    RC2_Transmit_PDO_Mapping_Torque_actual_value_6077_00 : INT;
    RC2_Transmit_PDO_Mapping_Digital_inputs_60FD_00 : UDINT;
    RC2_Transmit_PDO_Mapping_Error_code_603F_00 : UINT;
    RC3_Receive_PDO_Mapping_ControlWord_6040_00 : UINT;
    RC3_Receive_PDO_Mapping_Target_Position_607A_00 : DINT;
    RC3_Receive_PDO_Mapping_Mode_of_operation_6060_00 : SINT;
    RC3_Receive_PDO_Mapping_Profile_velocity_6081_00 : UDINT;
    RC3_Receive_PDO_Mapping_Profile_acceleration_6083_00 : UDINT;
    RC3_Receive_PDO_Mapping_Profile_deceleration_6084_00 : UDINT;
    RC3_Receive_PDO_Mapping_Physical_outputs_60FE_01 : UDINT;
    RC3_Transmit_PDO_Mapping_StatusWord_6041_00 : UINT;
    RC3_Transmit_PDO_Mapping_Position_actual_value_6064_00 : DINT;
    RC3_Transmit_PDO_Mapping_Mode_of_operation_display_6061_00 : SINT;
    RC3_Transmit_PDO_Mapping_Following_error_actual_valu_60F4_00 : DINT;
    RC3_Transmit_PDO_Mapping_Torque_actual_value_6077_00 : INT;
    RC3_Transmit_PDO_Mapping_Digital_inputs_60FD_00 : UDINT;
    RC3_Transmit_PDO_Mapping_Error_code_603F_00 : UINT;
    RC4_Receive_PDO_Mapping_ControlWord_6040_00 : UINT;
    RC4_Receive_PDO_Mapping_Target_Position_607A_00 : DINT;
    RC4_Receive_PDO_Mapping_Mode_of_operation_6060_00 : SINT;
    RC4_Receive_PDO_Mapping_Profile_velocity_6081_00 : UDINT;
    RC4_Receive_PDO_Mapping_Profile_acceleration_6083_00 : UDINT;
    RC4_Receive_PDO_Mapping_Profile_deceleration_6084_00 : UDINT;
    RC4_Receive_PDO_Mapping_Physical_outputs_60FE_01 : UDINT;
    RC4_Transmit_PDO_Mapping_StatusWord_6041_00 : UINT;
    RC4_Transmit_PDO_Mapping_Position_actual_value_6064_00 : DINT;
    RC4_Transmit_PDO_Mapping_Mode_of_operation_display_6061_00 : SINT;
    RC4_Transmit_PDO_Mapping_Following_error_actual_valu_60F4_00 : DINT;
    RC4_Transmit_PDO_Mapping_Torque_actual_value_6077_00 : INT;
    RC4_Transmit_PDO_Mapping_Digital_inputs_60FD_00 : UDINT;
    RC4_Transmit_PDO_Mapping_Error_code_603F_00 : UINT;
    RC5_Receive_PDO_Mapping_ControlWord_6040_00 : UINT;
    RC5_Receive_PDO_Mapping_Target_Position_607A_00 : DINT;
    RC5_Receive_PDO_Mapping_Mode_of_operation_6060_00 : SINT;
    RC5_Receive_PDO_Mapping_Profile_velocity_6081_00 : UDINT;
    RC5_Receive_PDO_Mapping_Profile_acceleration_6083_00 : UDINT;
    RC5_Receive_PDO_Mapping_Profile_deceleration_6084_00 : UDINT;
    RC5_Receive_PDO_Mapping_Physical_outputs_60FE_01 : UDINT;
    RC5_Transmit_PDO_Mapping_StatusWord_6041_00 : UINT;
    RC5_Transmit_PDO_Mapping_Position_actual_value_6064_00 : DINT;
    RC5_Transmit_PDO_Mapping_Mode_of_operation_display_6061_00 : SINT;
    RC5_Transmit_PDO_Mapping_Following_error_actual_valu_60F4_00 : DINT;
    RC5_Transmit_PDO_Mapping_Torque_actual_value_6077_00 : INT;
    RC5_Transmit_PDO_Mapping_Digital_inputs_60FD_00 : UDINT;
    RC5_Transmit_PDO_Mapping_Error_code_603F_00 : UINT;
    RC6_Receive_PDO_Mapping_ControlWord_6040_00 : UINT;
    RC6_Receive_PDO_Mapping_ControlWord_6040_00_1 : UINT;
    RC6_Receive_PDO_Mapping_Target_Position_607A_00 : DINT;
    RC6_Receive_PDO_Mapping_Mode_of_operation_6060_00 : SINT;
    RC6_Receive_PDO_Mapping_Profile_velocity_6081_00 : UDINT;
    RC6_Receive_PDO_Mapping_Profile_acceleration_6083_00 : UDINT;
    RC6_Receive_PDO_Mapping_Profile_deceleration_6084_00 : UDINT;
    RC6_Receive_PDO_Mapping_Physical_outputs_60FE_01 : UDINT;
    RC6_Transmit_PDO_Mapping_StatusWord_6041_00 : UINT;
    RC6_Transmit_PDO_Mapping_Position_actual_value_6064_00 : DINT;
    RC6_Transmit_PDO_Mapping_Mode_of_operation_display_6061_00 : SINT;
    RC6_Transmit_PDO_Mapping_Following_error_actual_valu_60F4_00 : DINT;
    RC6_Transmit_PDO_Mapping_Torque_actual_value_6077_00 : INT;
    RC6_Transmit_PDO_Mapping_Digital_inputs_60FD_00 : UDINT;
    RC6_Transmit_PDO_Mapping_Error_code_603F_00 : UINT;
END_VAR
VAR_GLOBAL RETAIN
    RCON1_OUT : ARRAY[1..6] OF ST_RCON_Direct_OUT_Axis;  (* RCON1 (PLC→RCON); [2] 2軸目; [3] 3軸目; [4] 4軸目; [5] 5軸目; [6] 6軸目; [1].Control.Pause 一時停止（STP/b2）; [1] 1軸目 *)
    RCON1_IN : ARRAY[1..6] OF ST_RCON_Direct_IN_Axis;  (* RCON1 (RCON→PLC); [1] 1軸目; [2] 2軸目; [3] 3軸目; [4] 4軸目; [5] 5軸目; [6] 6軸目 *)
END_VAR
VAR_GLOBAL
    RCON1_SpeedUnit_mm_s : LREAL;  (* RCON1 速度単位 [mm/s/カウント]（1.0/0.1） *)
    RCON1_OUT_GwControl0Raw : UINT;  (* 未割付・不使用 OUT00 共通制御（MON/RTE） *)
    RCON1_OUT_GwControl1ReservedRaw : UINT;  (* 未割付・不使用 OUT01 予約（書込禁止） *)
    RCON1_OUT_ReservedOut02Raw : UINT;  (* 未割付・不使用 OUT02 予約（書込禁止） *)
    RCON1_OUT_ReservedOut03Raw : UINT;  (* 未割付・不使用 OUT03 予約（書込禁止） *)
    RCON1_OUT_ReservedOut04Raw : UINT;  (* 未割付・不使用 OUT04 予約（書込禁止） *)
    RCON1_OUT_ReservedOut05Raw : UINT;  (* 未割付・不使用 OUT05 予約（書込禁止） *)
    RCON1_OUT_ReservedOut06Raw : UINT;  (* 未割付・不使用 OUT06 予約（書込禁止） *)
    RCON1_OUT_ReservedOut07Raw : UINT;  (* 未割付・不使用 OUT07 予約（書込禁止） *)
    RCON1_OUT_Axis1_TargetPosLoRaw : UINT;  (* 未割付・不使用 OUT08 1軸目 目標位置 下位 [0.01mm] *)
    RCON1_OUT_Axis1_TargetPosHiRaw : UINT;  (* 未割付・不使用 OUT09 1軸目 目標位置 上位 [0.01mm] *)
    RCON1_OUT_Axis1_PositionBandLoRaw : UINT;  (* 未割付・不使用 OUT10 1軸目 位置決め幅 下位 [0.01mm] *)
    RCON1_OUT_Axis1_PositionBandHiRaw : UINT;  (* 未割付・不使用 OUT11 1軸目 位置決め幅 上位 [0.01mm] *)
    RCON1_OUT_Axis1_SpeedRaw : UINT;  (* 未割付・不使用 OUT12 1軸目 速度指令 [実機単位] *)
    RCON1_OUT_Axis1_AccDecRaw : UINT;  (* 未割付・不使用 OUT13 1軸目 共通加減速 [0.01G] *)
    RCON1_OUT_Axis1_PushLimitRaw : UINT;  (* 未割付・不使用 OUT14 1軸目 押付け制限 [255=100%] *)
    RCON1_OUT_Axis1_ControlRaw : UINT;  (* 未割付・不使用 OUT15 1軸目 制御信号（DSTR/SON等） *)
    RCON1_OUT_Axis2_TargetPosLoRaw : UINT;  (* 未割付・不使用 OUT16 2軸目 目標位置 下位 [0.01mm] *)
    RCON1_OUT_Axis2_TargetPosHiRaw : UINT;  (* 未割付・不使用 OUT17 2軸目 目標位置 上位 [0.01mm] *)
    RCON1_OUT_Axis2_PositionBandLoRaw : UINT;  (* 未割付・不使用 OUT18 2軸目 位置決め幅 下位 [0.01mm] *)
    RCON1_OUT_Axis2_PositionBandHiRaw : UINT;  (* 未割付・不使用 OUT19 2軸目 位置決め幅 上位 [0.01mm] *)
    RCON1_OUT_Axis2_SpeedRaw : UINT;  (* 未割付・不使用 OUT20 2軸目 速度指令 [実機単位] *)
    RCON1_OUT_Axis2_AccDecRaw : UINT;  (* 未割付・不使用 OUT21 2軸目 共通加減速 [0.01G] *)
    RCON1_OUT_Axis2_PushLimitRaw : UINT;  (* 未割付・不使用 OUT22 2軸目 押付け制限 [255=100%] *)
    RCON1_OUT_Axis2_ControlRaw : UINT;  (* 未割付・不使用 OUT23 2軸目 制御信号（DSTR/SON等） *)
    RCON1_OUT_Axis3_TargetPosLoRaw : UINT;  (* 未割付・不使用 OUT24 3軸目 目標位置 下位 [0.01mm] *)
    RCON1_OUT_Axis3_TargetPosHiRaw : UINT;  (* 未割付・不使用 OUT25 3軸目 目標位置 上位 [0.01mm] *)
    RCON1_OUT_Axis3_PositionBandLoRaw : UINT;  (* 未割付・不使用 OUT26 3軸目 位置決め幅 下位 [0.01mm] *)
    RCON1_OUT_Axis3_PositionBandHiRaw : UINT;  (* 未割付・不使用 OUT27 3軸目 位置決め幅 上位 [0.01mm] *)
    RCON1_OUT_Axis3_SpeedRaw : UINT;  (* 未割付・不使用 OUT28 3軸目 速度指令 [実機単位] *)
    RCON1_OUT_Axis3_AccDecRaw : UINT;  (* 未割付・不使用 OUT29 3軸目 共通加減速 [0.01G] *)
    RCON1_OUT_Axis3_PushLimitRaw : UINT;  (* 未割付・不使用 OUT30 3軸目 押付け制限 [255=100%] *)
    RCON1_OUT_Axis3_ControlRaw : UINT;  (* 未割付・不使用 OUT31 3軸目 制御信号（DSTR/SON等） *)
    RCON1_OUT_Axis4_TargetPosLoRaw : UINT;  (* 未割付・不使用 OUT32 4軸目 目標位置 下位 [0.01mm] *)
    RCON1_OUT_Axis4_TargetPosHiRaw : UINT;  (* 未割付・不使用 OUT33 4軸目 目標位置 上位 [0.01mm] *)
    RCON1_OUT_Axis4_PositionBandLoRaw : UINT;  (* 未割付・不使用 OUT34 4軸目 位置決め幅 下位 [0.01mm] *)
    RCON1_OUT_Axis4_PositionBandHiRaw : UINT;  (* 未割付・不使用 OUT35 4軸目 位置決め幅 上位 [0.01mm] *)
    RCON1_OUT_Axis4_SpeedRaw : UINT;  (* 未割付・不使用 OUT36 4軸目 速度指令 [実機単位] *)
    RCON1_OUT_Axis4_AccDecRaw : UINT;  (* 未割付・不使用 OUT37 4軸目 共通加減速 [0.01G] *)
    RCON1_OUT_Axis4_PushLimitRaw : UINT;  (* 未割付・不使用 OUT38 4軸目 押付け制限 [255=100%] *)
    RCON1_OUT_Axis4_ControlRaw : UINT;  (* 未割付・不使用 OUT39 4軸目 制御信号（DSTR/SON等） *)
    RCON1_OUT_Axis5_TargetPosLoRaw : UINT;  (* 未割付・不使用 OUT40 5軸目 目標位置 下位 [0.01mm] *)
    RCON1_OUT_Axis5_TargetPosHiRaw : UINT;  (* 未割付・不使用 OUT41 5軸目 目標位置 上位 [0.01mm] *)
    RCON1_OUT_Axis5_PositionBandLoRaw : UINT;  (* 未割付・不使用 OUT42 5軸目 位置決め幅 下位 [0.01mm] *)
    RCON1_OUT_Axis5_PositionBandHiRaw : UINT;  (* 未割付・不使用 OUT43 5軸目 位置決め幅 上位 [0.01mm] *)
    RCON1_OUT_Axis5_SpeedRaw : UINT;  (* 未割付・不使用 OUT44 5軸目 速度指令 [実機単位] *)
    RCON1_OUT_Axis5_AccDecRaw : UINT;  (* 未割付・不使用 OUT45 5軸目 共通加減速 [0.01G] *)
    RCON1_OUT_Axis5_PushLimitRaw : UINT;  (* 未割付・不使用 OUT46 5軸目 押付け制限 [255=100%] *)
    RCON1_OUT_Axis5_ControlRaw : UINT;  (* 未割付・不使用 OUT47 5軸目 制御信号（DSTR/SON等） *)
    RCON1_OUT_Axis6_TargetPosLoRaw : UINT;  (* 未割付・不使用 OUT48 6軸目 目標位置 下位 [0.01mm] *)
    RCON1_OUT_Axis6_TargetPosHiRaw : UINT;  (* 未割付・不使用 OUT49 6軸目 目標位置 上位 [0.01mm] *)
    RCON1_OUT_Axis6_PositionBandLoRaw : UINT;  (* 未割付・不使用 OUT50 6軸目 位置決め幅 下位 [0.01mm] *)
    RCON1_OUT_Axis6_PositionBandHiRaw : UINT;  (* 未割付・不使用 OUT51 6軸目 位置決め幅 上位 [0.01mm] *)
    RCON1_OUT_Axis6_SpeedRaw : UINT;  (* 未割付・不使用 OUT52 6軸目 速度指令 [実機単位] *)
    RCON1_OUT_Axis6_AccDecRaw : UINT;  (* 未割付・不使用 OUT53 6軸目 共通加減速 [0.01G] *)
    RCON1_OUT_Axis6_PushLimitRaw : UINT;  (* 未割付・不使用 OUT54 6軸目 押付け制限 [255=100%] *)
    RCON1_OUT_Axis6_ControlRaw : UINT;  (* 未割付・不使用 OUT55 6軸目 制御信号（DSTR/SON等） *)
    RCON1_IN_GwStatus0Raw : UINT;  (* 未割付・不使用 IN00 GW状態 *)
    RCON1_IN_AxisLinkStatusRaw : UINT;  (* 未割付・不使用 IN01 軸リンク状態 *)
    RCON1_IN_PowerStatus0Raw : UINT;  (* 未割付・不使用 IN02 電源状態0 *)
    RCON1_IN_PowerStatus1Raw : UINT;  (* 未割付・不使用 IN03 電源状態1 *)
    RCON1_IN_PowerStatus2Raw : UINT;  (* 未割付・不使用 IN04 電源状態2 *)
    RCON1_IN_PowerStatus3Raw : UINT;  (* 未割付・不使用 IN05 電源状態3 *)
    RCON1_IN_PowerStatus4MaintenanceRaw : UINT;  (* 未割付・不使用 IN06 電源状態4（構成依存） *)
    RCON1_IN_ReservedIn07Raw : UINT;  (* 未割付・不使用 IN07 予約（使用禁止） *)
    RCON1_IN_Axis1_ActualPosLoRaw : UINT;  (* 未割付・不使用 IN08 1軸目 現在位置 下位 [0.01mm] *)
    RCON1_IN_Axis1_ActualPosHiRaw : UINT;  (* 未割付・不使用 IN09 1軸目 現在位置 上位 [0.01mm] *)
    RCON1_IN_Axis1_CurrentLoRaw : UINT;  (* 未割付・不使用 IN10 1軸目 指令電流 下位 [mA] *)
    RCON1_IN_Axis1_CurrentHiRaw : UINT;  (* 未割付・不使用 IN11 1軸目 指令電流 上位 [mA] *)
    RCON1_IN_Axis1_ActualSpeedRaw : UINT;  (* 未割付・不使用 IN12 1軸目 現在速度 [実機単位・符号付き] *)
    RCON1_IN_Axis1_ReservedInRaw : UINT;  (* 未割付・不使用 IN13 1軸目 予約（使用禁止） *)
    RCON1_IN_Axis1_AlarmCodeRaw : UINT;  (* 未割付・不使用 IN14 1軸目 軸異常コード *)
    RCON1_IN_Axis1_StatusRaw : UINT;  (* 未割付・不使用 IN15 1軸目 状態信号（PEND/SV等） *)
    RCON1_IN_Axis2_ActualPosLoRaw : UINT;  (* 未割付・不使用 IN16 2軸目 現在位置 下位 [0.01mm] *)
    RCON1_IN_Axis2_ActualPosHiRaw : UINT;  (* 未割付・不使用 IN17 2軸目 現在位置 上位 [0.01mm] *)
    RCON1_IN_Axis2_CurrentLoRaw : UINT;  (* 未割付・不使用 IN18 2軸目 指令電流 下位 [mA] *)
    RCON1_IN_Axis2_CurrentHiRaw : UINT;  (* 未割付・不使用 IN19 2軸目 指令電流 上位 [mA] *)
    RCON1_IN_Axis2_ActualSpeedRaw : UINT;  (* 未割付・不使用 IN20 2軸目 現在速度 [実機単位・符号付き] *)
    RCON1_IN_Axis2_ReservedInRaw : UINT;  (* 未割付・不使用 IN21 2軸目 予約（使用禁止） *)
    RCON1_IN_Axis2_AlarmCodeRaw : UINT;  (* 未割付・不使用 IN22 2軸目 軸異常コード *)
    RCON1_IN_Axis2_StatusRaw : UINT;  (* 未割付・不使用 IN23 2軸目 状態信号（PEND/SV等） *)
    RCON1_IN_Axis3_ActualPosLoRaw : UINT;  (* 未割付・不使用 IN24 3軸目 現在位置 下位 [0.01mm] *)
    RCON1_IN_Axis3_ActualPosHiRaw : UINT;  (* 未割付・不使用 IN25 3軸目 現在位置 上位 [0.01mm] *)
    RCON1_IN_Axis3_CurrentLoRaw : UINT;  (* 未割付・不使用 IN26 3軸目 指令電流 下位 [mA] *)
    RCON1_IN_Axis3_CurrentHiRaw : UINT;  (* 未割付・不使用 IN27 3軸目 指令電流 上位 [mA] *)
    RCON1_IN_Axis3_ActualSpeedRaw : UINT;  (* 未割付・不使用 IN28 3軸目 現在速度 [実機単位・符号付き] *)
    RCON1_IN_Axis3_ReservedInRaw : UINT;  (* 未割付・不使用 IN29 3軸目 予約（使用禁止） *)
    RCON1_IN_Axis3_AlarmCodeRaw : UINT;  (* 未割付・不使用 IN30 3軸目 軸異常コード *)
    RCON1_IN_Axis3_StatusRaw : UINT;  (* 未割付・不使用 IN31 3軸目 状態信号（PEND/SV等） *)
    RCON1_IN_Axis4_ActualPosLoRaw : UINT;  (* 未割付・不使用 IN32 4軸目 現在位置 下位 [0.01mm] *)
    RCON1_IN_Axis4_ActualPosHiRaw : UINT;  (* 未割付・不使用 IN33 4軸目 現在位置 上位 [0.01mm] *)
    RCON1_IN_Axis4_CurrentLoRaw : UINT;  (* 未割付・不使用 IN34 4軸目 指令電流 下位 [mA] *)
    RCON1_IN_Axis4_CurrentHiRaw : UINT;  (* 未割付・不使用 IN35 4軸目 指令電流 上位 [mA] *)
    RCON1_IN_Axis4_ActualSpeedRaw : UINT;  (* 未割付・不使用 IN36 4軸目 現在速度 [実機単位・符号付き] *)
    RCON1_IN_Axis4_ReservedInRaw : UINT;  (* 未割付・不使用 IN37 4軸目 予約（使用禁止） *)
    RCON1_IN_Axis4_AlarmCodeRaw : UINT;  (* 未割付・不使用 IN38 4軸目 軸異常コード *)
    RCON1_IN_Axis4_StatusRaw : UINT;  (* 未割付・不使用 IN39 4軸目 状態信号（PEND/SV等） *)
    RCON1_IN_Axis5_ActualPosLoRaw : UINT;  (* 未割付・不使用 IN40 5軸目 現在位置 下位 [0.01mm] *)
    RCON1_IN_Axis5_ActualPosHiRaw : UINT;  (* 未割付・不使用 IN41 5軸目 現在位置 上位 [0.01mm] *)
    RCON1_IN_Axis5_CurrentLoRaw : UINT;  (* 未割付・不使用 IN42 5軸目 指令電流 下位 [mA] *)
    RCON1_IN_Axis5_CurrentHiRaw : UINT;  (* 未割付・不使用 IN43 5軸目 指令電流 上位 [mA] *)
    RCON1_IN_Axis5_ActualSpeedRaw : UINT;  (* 未割付・不使用 IN44 5軸目 現在速度 [実機単位・符号付き] *)
    RCON1_IN_Axis5_ReservedInRaw : UINT;  (* 未割付・不使用 IN45 5軸目 予約（使用禁止） *)
    RCON1_IN_Axis5_AlarmCodeRaw : UINT;  (* 未割付・不使用 IN46 5軸目 軸異常コード *)
    RCON1_IN_Axis5_StatusRaw : UINT;  (* 未割付・不使用 IN47 5軸目 状態信号（PEND/SV等） *)
    RCON1_IN_Axis6_ActualPosLoRaw : UINT;  (* 未割付・不使用 IN48 6軸目 現在位置 下位 [0.01mm] *)
    RCON1_IN_Axis6_ActualPosHiRaw : UINT;  (* 未割付・不使用 IN49 6軸目 現在位置 上位 [0.01mm] *)
    RCON1_IN_Axis6_CurrentLoRaw : UINT;  (* 未割付・不使用 IN50 6軸目 指令電流 下位 [mA] *)
    RCON1_IN_Axis6_CurrentHiRaw : UINT;  (* 未割付・不使用 IN51 6軸目 指令電流 上位 [mA] *)
    RCON1_IN_Axis6_ActualSpeedRaw : UINT;  (* 未割付・不使用 IN52 6軸目 現在速度 [実機単位・符号付き] *)
    RCON1_IN_Axis6_ReservedInRaw : UINT;  (* 未割付・不使用 IN53 6軸目 予約（使用禁止） *)
    RCON1_IN_Axis6_AlarmCodeRaw : UINT;  (* 未割付・不使用 IN54 6軸目 軸異常コード *)
END_VAR
VAR_GLOBAL RETAIN
    RCON1_IN_Axis6_StatusRaw : UINT;  (* 未割付・不使用 IN55 6軸目 状態信号（PEND/SV等） *)
    RCON2_OUT : ARRAY[1..5] OF ST_RCON_Direct_OUT_Axis;  (* RCON2 出力指令（PLC→RCON）; [1] 1軸目（No.0）出力指令; [2] 2軸目（No.1）出力指令; [3] 3軸目（No.2）出力指令; [4] 4軸目（No.3）出力指令; [5] 5軸目（No.4）出力指令 *)
END_VAR
VAR_GLOBAL
    RCON2_IN : ARRAY[1..5] OF ST_RCON_Direct_IN_Axis;  (* RCON2 入力情報（RCON→PLC）; [1] 1軸目（No.0）入力情報; [2] 2軸目（No.1）入力情報; [3] 3軸目（No.2）入力情報; [4] 4軸目（No.3）入力情報; [5] 5軸目（No.4）入力情報 *)
    RCON2_SpeedUnit_mm_s : LREAL;  (* RCON2 速度単位 [mm/s/カウント]（1.0/0.1） *)
    RCON2_OUT_GwControl0Raw : UINT;  (* 未割付・不使用 OUT00 共通制御（MON/RTE） *)
    RCON2_OUT_GwControl1ReservedRaw : UINT;  (* 未割付・不使用 OUT01 予約（書込禁止） *)
    RCON2_OUT_ReservedOut02Raw : UINT;  (* 未割付・不使用 OUT02 予約（書込禁止） *)
    RCON2_OUT_ReservedOut03Raw : UINT;  (* 未割付・不使用 OUT03 予約（書込禁止） *)
    RCON2_OUT_ReservedOut04Raw : UINT;  (* 未割付・不使用 OUT04 予約（書込禁止） *)
    RCON2_OUT_ReservedOut05Raw : UINT;  (* 未割付・不使用 OUT05 予約（書込禁止） *)
    RCON2_OUT_ReservedOut06Raw : UINT;  (* 未割付・不使用 OUT06 予約（書込禁止） *)
    RCON2_OUT_ReservedOut07Raw : UINT;  (* 未割付・不使用 OUT07 予約（書込禁止） *)
    RCON2_OUT_Axis1_TargetPosLoRaw : UINT;  (* 未割付・不使用 OUT08 1軸目 目標位置 下位 [0.01mm] *)
    RCON2_OUT_Axis1_TargetPosHiRaw : UINT;  (* 未割付・不使用 OUT09 1軸目 目標位置 上位 [0.01mm] *)
    RCON2_OUT_Axis1_PositionBandLoRaw : UINT;  (* 未割付・不使用 OUT10 1軸目 位置決め幅 下位 [0.01mm] *)
    RCON2_OUT_Axis1_PositionBandHiRaw : UINT;  (* 未割付・不使用 OUT11 1軸目 位置決め幅 上位 [0.01mm] *)
    RCON2_OUT_Axis1_SpeedRaw : UINT;  (* 未割付・不使用 OUT12 1軸目 速度指令 [実機単位] *)
    RCON2_OUT_Axis1_AccDecRaw : UINT;  (* 未割付・不使用 OUT13 1軸目 共通加減速 [0.01G] *)
    RCON2_OUT_Axis1_PushLimitRaw : UINT;  (* 未割付・不使用 OUT14 1軸目 押付け制限 [255=100%] *)
    RCON2_OUT_Axis1_ControlRaw : UINT;  (* 未割付・不使用 OUT15 1軸目 制御信号（DSTR/SON等） *)
    RCON2_OUT_Axis2_TargetPosLoRaw : UINT;  (* 未割付・不使用 OUT16 2軸目 目標位置 下位 [0.01mm] *)
    RCON2_OUT_Axis2_TargetPosHiRaw : UINT;  (* 未割付・不使用 OUT17 2軸目 目標位置 上位 [0.01mm] *)
    RCON2_OUT_Axis2_PositionBandLoRaw : UINT;  (* 未割付・不使用 OUT18 2軸目 位置決め幅 下位 [0.01mm] *)
    RCON2_OUT_Axis2_PositionBandHiRaw : UINT;  (* 未割付・不使用 OUT19 2軸目 位置決め幅 上位 [0.01mm] *)
    RCON2_OUT_Axis2_SpeedRaw : UINT;  (* 未割付・不使用 OUT20 2軸目 速度指令 [実機単位] *)
    RCON2_OUT_Axis2_AccDecRaw : UINT;  (* 未割付・不使用 OUT21 2軸目 共通加減速 [0.01G] *)
    RCON2_OUT_Axis2_PushLimitRaw : UINT;  (* 未割付・不使用 OUT22 2軸目 押付け制限 [255=100%] *)
    RCON2_OUT_Axis2_ControlRaw : UINT;  (* 未割付・不使用 OUT23 2軸目 制御信号（DSTR/SON等） *)
    RCON2_OUT_Axis3_TargetPosLoRaw : UINT;  (* 未割付・不使用 OUT24 3軸目 目標位置 下位 [0.01mm] *)
    RCON2_OUT_Axis3_TargetPosHiRaw : UINT;  (* 未割付・不使用 OUT25 3軸目 目標位置 上位 [0.01mm] *)
    RCON2_OUT_Axis3_PositionBandLoRaw : UINT;  (* 未割付・不使用 OUT26 3軸目 位置決め幅 下位 [0.01mm] *)
    RCON2_OUT_Axis3_PositionBandHiRaw : UINT;  (* 未割付・不使用 OUT27 3軸目 位置決め幅 上位 [0.01mm] *)
    RCON2_OUT_Axis3_SpeedRaw : UINT;  (* 未割付・不使用 OUT28 3軸目 速度指令 [実機単位] *)
    RCON2_OUT_Axis3_AccDecRaw : UINT;  (* 未割付・不使用 OUT29 3軸目 共通加減速 [0.01G] *)
    RCON2_OUT_Axis3_PushLimitRaw : UINT;  (* 未割付・不使用 OUT30 3軸目 押付け制限 [255=100%] *)
    RCON2_OUT_Axis3_ControlRaw : UINT;  (* 未割付・不使用 OUT31 3軸目 制御信号（DSTR/SON等） *)
    RCON2_OUT_Axis4_TargetPosLoRaw : UINT;  (* 未割付・不使用 OUT32 4軸目 目標位置 下位 [0.01mm] *)
    RCON2_OUT_Axis4_TargetPosHiRaw : UINT;  (* 未割付・不使用 OUT33 4軸目 目標位置 上位 [0.01mm] *)
    RCON2_OUT_Axis4_PositionBandLoRaw : UINT;  (* 未割付・不使用 OUT34 4軸目 位置決め幅 下位 [0.01mm] *)
    RCON2_OUT_Axis4_PositionBandHiRaw : UINT;  (* 未割付・不使用 OUT35 4軸目 位置決め幅 上位 [0.01mm] *)
    RCON2_OUT_Axis4_SpeedRaw : UINT;  (* 未割付・不使用 OUT36 4軸目 速度指令 [実機単位] *)
    RCON2_OUT_Axis4_AccDecRaw : UINT;  (* 未割付・不使用 OUT37 4軸目 共通加減速 [0.01G] *)
    RCON2_OUT_Axis4_PushLimitRaw : UINT;  (* 未割付・不使用 OUT38 4軸目 押付け制限 [255=100%] *)
    RCON2_OUT_Axis4_ControlRaw : UINT;  (* 未割付・不使用 OUT39 4軸目 制御信号（DSTR/SON等） *)
    RCON2_OUT_Axis5_TargetPosLoRaw : UINT;  (* 未割付・不使用 OUT40 5軸目 目標位置 下位 [0.01mm] *)
    RCON2_OUT_Axis5_TargetPosHiRaw : UINT;  (* 未割付・不使用 OUT41 5軸目 目標位置 上位 [0.01mm] *)
    RCON2_OUT_Axis5_PositionBandLoRaw : UINT;  (* 未割付・不使用 OUT42 5軸目 位置決め幅 下位 [0.01mm] *)
    RCON2_OUT_Axis5_PositionBandHiRaw : UINT;  (* 未割付・不使用 OUT43 5軸目 位置決め幅 上位 [0.01mm] *)
    RCON2_OUT_Axis5_SpeedRaw : UINT;  (* 未割付・不使用 OUT44 5軸目 速度指令 [実機単位] *)
    RCON2_OUT_Axis5_AccDecRaw : UINT;  (* 未割付・不使用 OUT45 5軸目 共通加減速 [0.01G] *)
    RCON2_OUT_Axis5_PushLimitRaw : UINT;  (* 未割付・不使用 OUT46 5軸目 押付け制限 [255=100%] *)
    RCON2_OUT_Axis5_ControlRaw : UINT;  (* 未割付・不使用 OUT47 5軸目 制御信号（DSTR/SON等） *)
    RCON2_IN_GwStatus0Raw : UINT;  (* 未割付・不使用 IN00 GW状態 *)
    RCON2_IN_AxisLinkStatusRaw : UINT;  (* 未割付・不使用 IN01 軸リンク状態 *)
    RCON2_IN_PowerStatus0Raw : UINT;  (* 未割付・不使用 IN02 電源状態0 *)
    RCON2_IN_PowerStatus1Raw : UINT;  (* 未割付・不使用 IN03 電源状態1 *)
    RCON2_IN_PowerStatus2Raw : UINT;  (* 未割付・不使用 IN04 電源状態2 *)
    RCON2_IN_PowerStatus3Raw : UINT;  (* 未割付・不使用 IN05 電源状態3 *)
    RCON2_IN_PowerStatus4MaintenanceRaw : UINT;  (* 未割付・不使用 IN06 電源状態4（構成依存） *)
    RCON2_IN_ReservedIn07Raw : UINT;  (* 未割付・不使用 IN07 予約（使用禁止） *)
    RCON2_IN_Axis1_ActualPosLoRaw : UINT;  (* 未割付・不使用 IN08 1軸目 現在位置 下位 [0.01mm] *)
    RCON2_IN_Axis1_ActualPosHiRaw : UINT;  (* 未割付・不使用 IN09 1軸目 現在位置 上位 [0.01mm] *)
    RCON2_IN_Axis1_CurrentLoRaw : UINT;  (* 未割付・不使用 IN10 1軸目 指令電流 下位 [mA] *)
    RCON2_IN_Axis1_CurrentHiRaw : UINT;  (* 未割付・不使用 IN11 1軸目 指令電流 上位 [mA] *)
    RCON2_IN_Axis1_ActualSpeedRaw : UINT;  (* 未割付・不使用 IN12 1軸目 現在速度 [実機単位・符号付き] *)
    RCON2_IN_Axis1_ReservedInRaw : UINT;  (* 未割付・不使用 IN13 1軸目 予約（使用禁止） *)
    RCON2_IN_Axis1_AlarmCodeRaw : UINT;  (* 未割付・不使用 IN14 1軸目 軸異常コード *)
    RCON2_IN_Axis1_StatusRaw : UINT;  (* 未割付・不使用 IN15 1軸目 状態信号（PEND/SV等） *)
    RCON2_IN_Axis2_ActualPosLoRaw : UINT;  (* 未割付・不使用 IN16 2軸目 現在位置 下位 [0.01mm] *)
    RCON2_IN_Axis2_ActualPosHiRaw : UINT;  (* 未割付・不使用 IN17 2軸目 現在位置 上位 [0.01mm] *)
    RCON2_IN_Axis2_CurrentLoRaw : UINT;  (* 未割付・不使用 IN18 2軸目 指令電流 下位 [mA] *)
    RCON2_IN_Axis2_CurrentHiRaw : UINT;  (* 未割付・不使用 IN19 2軸目 指令電流 上位 [mA] *)
    RCON2_IN_Axis2_ActualSpeedRaw : UINT;  (* 未割付・不使用 IN20 2軸目 現在速度 [実機単位・符号付き] *)
    RCON2_IN_Axis2_ReservedInRaw : UINT;  (* 未割付・不使用 IN21 2軸目 予約（使用禁止） *)
    RCON2_IN_Axis2_AlarmCodeRaw : UINT;  (* 未割付・不使用 IN22 2軸目 軸異常コード *)
    RCON2_IN_Axis2_StatusRaw : UINT;  (* 未割付・不使用 IN23 2軸目 状態信号（PEND/SV等） *)
    RCON2_IN_Axis3_ActualPosLoRaw : UINT;  (* 未割付・不使用 IN24 3軸目 現在位置 下位 [0.01mm] *)
    RCON2_IN_Axis3_ActualPosHiRaw : UINT;  (* 未割付・不使用 IN25 3軸目 現在位置 上位 [0.01mm] *)
    RCON2_IN_Axis3_CurrentLoRaw : UINT;  (* 未割付・不使用 IN26 3軸目 指令電流 下位 [mA] *)
    RCON2_IN_Axis3_CurrentHiRaw : UINT;  (* 未割付・不使用 IN27 3軸目 指令電流 上位 [mA] *)
    RCON2_IN_Axis3_ActualSpeedRaw : UINT;  (* 未割付・不使用 IN28 3軸目 現在速度 [実機単位・符号付き] *)
    RCON2_IN_Axis3_ReservedInRaw : UINT;  (* 未割付・不使用 IN29 3軸目 予約（使用禁止） *)
    RCON2_IN_Axis3_AlarmCodeRaw : UINT;  (* 未割付・不使用 IN30 3軸目 軸異常コード *)
    RCON2_IN_Axis3_StatusRaw : UINT;  (* 未割付・不使用 IN31 3軸目 状態信号（PEND/SV等） *)
    RCON2_IN_Axis4_ActualPosLoRaw : UINT;  (* 未割付・不使用 IN32 4軸目 現在位置 下位 [0.01mm] *)
    RCON2_IN_Axis4_ActualPosHiRaw : UINT;  (* 未割付・不使用 IN33 4軸目 現在位置 上位 [0.01mm] *)
    RCON2_IN_Axis4_CurrentLoRaw : UINT;  (* 未割付・不使用 IN34 4軸目 指令電流 下位 [mA] *)
    RCON2_IN_Axis4_CurrentHiRaw : UINT;  (* 未割付・不使用 IN35 4軸目 指令電流 上位 [mA] *)
    RCON2_IN_Axis4_ActualSpeedRaw : UINT;  (* 未割付・不使用 IN36 4軸目 現在速度 [実機単位・符号付き] *)
    RCON2_IN_Axis4_ReservedInRaw : UINT;  (* 未割付・不使用 IN37 4軸目 予約（使用禁止） *)
    RCON2_IN_Axis4_AlarmCodeRaw : UINT;  (* 未割付・不使用 IN38 4軸目 軸異常コード *)
    RCON2_IN_Axis4_StatusRaw : UINT;  (* 未割付・不使用 IN39 4軸目 状態信号（PEND/SV等） *)
    RCON2_IN_Axis5_ActualPosLoRaw : UINT;  (* 未割付・不使用 IN40 5軸目 現在位置 下位 [0.01mm] *)
    RCON2_IN_Axis5_ActualPosHiRaw : UINT;  (* 未割付・不使用 IN41 5軸目 現在位置 上位 [0.01mm] *)
    RCON2_IN_Axis5_CurrentLoRaw : UINT;  (* 未割付・不使用 IN42 5軸目 指令電流 下位 [mA] *)
    RCON2_IN_Axis5_CurrentHiRaw : UINT;  (* 未割付・不使用 IN43 5軸目 指令電流 上位 [mA] *)
    RCON2_IN_Axis5_ActualSpeedRaw : UINT;  (* 未割付・不使用 IN44 5軸目 現在速度 [実機単位・符号付き] *)
    RCON2_IN_Axis5_ReservedInRaw : UINT;  (* 未割付・不使用 IN45 5軸目 予約（使用禁止） *)
    RCON2_IN_Axis5_AlarmCodeRaw : UINT;  (* 未割付・不使用 IN46 5軸目 軸異常コード *)
    RCON2_IN_Axis5_StatusRaw : UINT;  (* 未割付・不使用 IN47 5軸目 状態信号（PEND/SV等） *)
    E005_Out_OUT00_2003_01 : UINT;  (* 旧I/O候補（未割付・不使用） *)
    E005_Out_OUT01_2003_02 : UINT;  (* 旧I/O候補（未割付・不使用） *)
    E005_Out_OUT02_2003_03 : UINT;  (* 旧I/O候補（未割付・不使用） *)
    E005_Out_OUT03_2003_04 : UINT;  (* 旧I/O候補（未割付・不使用） *)
    E005_Out_OUT04_2003_05 : UINT;  (* 旧I/O候補（未割付・不使用） *)
    E005_Out_OUT05_2003_06 : UINT;  (* 旧I/O候補（未割付・不使用） *)
    E005_Out_OUT06_2003_07 : UINT;  (* 旧I/O候補（未割付・不使用） *)
    E005_Out_OUT07_2003_08 : UINT;  (* 旧I/O候補（未割付・不使用） *)
    E005_Out_OUT08_2003_09 : UINT;  (* 旧I/O候補（未割付・不使用） *)
    E005_Out_OUT09_2003_0A : UINT;  (* 旧I/O候補（未割付・不使用） *)
    E005_Out_OUT10_2003_0B : UINT;  (* 旧I/O候補（未割付・不使用） *)
    E005_Out_OUT11_2003_0C : UINT;  (* 旧I/O候補（未割付・不使用） *)
    E005_Out_OUT12_2003_0D : UINT;  (* 旧I/O候補（未割付・不使用） *)
    E005_Out_OUT13_2003_0E : UINT;  (* 旧I/O候補（未割付・不使用） *)
    E005_Out_OUT14_2003_0F : UINT;  (* 旧I/O候補（未割付・不使用） *)
    E005_Out_OUT15_2003_10 : UINT;  (* 旧I/O候補（未割付・不使用） *)
    E005_Out_OUT16_2003_11 : UINT;  (* 旧I/O候補（未割付・不使用） *)
    E005_Out_OUT17_2003_12 : UINT;  (* 旧I/O候補（未割付・不使用） *)
    E005_Out_OUT18_2003_13 : UINT;  (* 旧I/O候補（未割付・不使用） *)
    E005_Out_OUT19_2003_14 : UINT;  (* 旧I/O候補（未割付・不使用） *)
    E005_Out_OUT20_2003_15 : UINT;  (* 旧I/O候補（未割付・不使用） *)
    E005_Out_OUT21_2003_16 : UINT;  (* 旧I/O候補（未割付・不使用） *)
    E005_Out_OUT22_2003_17 : UINT;  (* 旧I/O候補（未割付・不使用） *)
    E005_Out_OUT23_2003_18 : UINT;  (* 旧I/O候補（未割付・不使用） *)
    E005_Out_OUT24_2003_19 : UINT;  (* 旧I/O候補（未割付・不使用） *)
    E005_Out_OUT25_2003_1A : UINT;  (* 旧I/O候補（未割付・不使用） *)
    E005_Out_OUT26_2003_1B : UINT;  (* 旧I/O候補（未割付・不使用） *)
    E005_Out_OUT27_2003_1C : UINT;  (* 旧I/O候補（未割付・不使用） *)
    E005_Out_OUT28_2003_1D : UINT;  (* 旧I/O候補（未割付・不使用） *)
    E005_Out_OUT29_2003_1E : UINT;  (* 旧I/O候補（未割付・不使用） *)
    E005_Out_OUT30_2003_1F : UINT;  (* 旧I/O候補（未割付・不使用） *)
    E005_Out_OUT31_2003_20 : UINT;  (* 旧I/O候補（未割付・不使用） *)
    E005_Out_OUT32_2003_21 : UINT;  (* 旧I/O候補（未割付・不使用） *)
    E005_Out_OUT33_2003_22 : UINT;  (* 旧I/O候補（未割付・不使用） *)
    E005_Out_OUT34_2003_23 : UINT;  (* 旧I/O候補（未割付・不使用） *)
    E005_Out_OUT35_2003_24 : UINT;  (* 旧I/O候補（未割付・不使用） *)
    E005_Out_OUT36_2003_25 : UINT;  (* 旧I/O候補（未割付・不使用） *)
    E005_Out_OUT37_2003_26 : UINT;  (* 旧I/O候補（未割付・不使用） *)
    E005_Out_OUT38_2003_27 : UINT;  (* 旧I/O候補（未割付・不使用） *)
    E005_Out_OUT39_2003_28 : UINT;  (* 旧I/O候補（未割付・不使用） *)
    E005_Out_OUT40_2003_29 : UINT;  (* 旧I/O候補（未割付・不使用） *)
    E005_Out_OUT41_2003_2A : UINT;  (* 旧I/O候補（未割付・不使用） *)
    E005_Out_OUT42_2003_2B : UINT;  (* 旧I/O候補（未割付・不使用） *)
    E005_Out_OUT43_2003_2C : UINT;  (* 旧I/O候補（未割付・不使用） *)
    E005_Out_OUT44_2003_2D : UINT;  (* 旧I/O候補（未割付・不使用） *)
    E005_Out_OUT45_2003_2E : UINT;  (* 旧I/O候補（未割付・不使用） *)
    E005_Out_OUT46_2003_2F : UINT;  (* 旧I/O候補（未割付・不使用） *)
    E005_Out_OUT47_2003_30 : UINT;  (* 旧I/O候補（未割付・不使用） *)
    E005_Out_OUT48_2003_31 : UINT;  (* 旧I/O候補（未割付・不使用） *)
    E005_Out_OUT49_2003_32 : UINT;  (* 旧I/O候補（未割付・不使用） *)
    E005_Out_OUT50_2003_33 : UINT;  (* 旧I/O候補（未割付・不使用） *)
    E005_Out_OUT51_2003_34 : UINT;  (* 旧I/O候補（未割付・不使用） *)
    E005_Out_OUT52_2003_35 : UINT;  (* 旧I/O候補（未割付・不使用） *)
    E005_Out_OUT53_2003_36 : UINT;  (* 旧I/O候補（未割付・不使用） *)
    E005_Out_OUT54_2003_37 : UINT;  (* 旧I/O候補（未割付・不使用） *)
    E005_Out_OUT55_2003_38 : UINT;  (* 旧I/O候補（未割付・不使用） *)
    E005_Out_OUT56_2003_39 : UINT;  (* 旧I/O候補（未割付・不使用） *)
    E005_Out_OUT57_2003_3A : UINT;  (* 旧I/O候補（未割付・不使用） *)
    E005_Out_OUT58_2003_3B : UINT;  (* 旧I/O候補（未割付・不使用） *)
    E005_Out_OUT59_2003_3C : UINT;  (* 旧I/O候補（未割付・不使用） *)
    E005_Out_OUT60_2003_3D : UINT;  (* 旧I/O候補（未割付・不使用） *)
    E005_Out_OUT61_2003_3E : UINT;  (* 旧I/O候補（未割付・不使用） *)
    E005_Out_OUT62_2003_3F : UINT;  (* 旧I/O候補（未割付・不使用） *)
    E005_Out_OUT63_2003_40 : UINT;  (* 旧I/O候補（未割付・不使用） *)
    E005_Out_OUT64_2003_41 : UINT;  (* 旧I/O候補（未割付・不使用） *)
    E005_Out_OUT65_2003_42 : UINT;  (* 旧I/O候補（未割付・不使用） *)
    E005_Out_OUT66_2003_43 : UINT;  (* 旧I/O候補（未割付・不使用） *)
    E005_Out_OUT67_2003_44 : UINT;  (* 旧I/O候補（未割付・不使用） *)
    E005_Out_OUT68_2003_45 : UINT;  (* 旧I/O候補（未割付・不使用） *)
    E005_Out_OUT69_2003_46 : UINT;  (* 旧I/O候補（未割付・不使用） *)
    E005_Out_OUT70_2003_47 : UINT;  (* 旧I/O候補（未割付・不使用） *)
    E005_Out_OUT71_2003_48 : UINT;  (* 旧I/O候補（未割付・不使用） *)
    E005_In_IN00_2004_01 : UINT;  (* 旧I/O候補（未割付・不使用） *)
    E005_In_IN01_2004_02 : UINT;  (* 旧I/O候補（未割付・不使用） *)
    E005_In_IN02_2004_03 : UINT;  (* 旧I/O候補（未割付・不使用） *)
    E005_In_IN03_2004_04 : UINT;  (* 旧I/O候補（未割付・不使用） *)
    E005_In_IN04_2004_05 : UINT;  (* 旧I/O候補（未割付・不使用） *)
    E005_In_IN05_2004_06 : UINT;  (* 旧I/O候補（未割付・不使用） *)
    E005_In_IN06_2004_07 : UINT;  (* 旧I/O候補（未割付・不使用） *)
    E005_In_IN07_2004_08 : UINT;  (* 旧I/O候補（未割付・不使用） *)
    E005_In_IN08_2004_09 : UINT;  (* 旧I/O候補（未割付・不使用） *)
    E005_In_IN09_2004_0A : UINT;  (* 旧I/O候補（未割付・不使用） *)
    E005_In_IN10_2004_0B : UINT;  (* 旧I/O候補（未割付・不使用） *)
    E005_In_IN11_2004_0C : UINT;  (* 旧I/O候補（未割付・不使用） *)
    E005_In_IN12_2004_0D : UINT;  (* 旧I/O候補（未割付・不使用） *)
    E005_In_IN13_2004_0E : UINT;  (* 旧I/O候補（未割付・不使用） *)
    E005_In_IN14_2004_0F : UINT;  (* 旧I/O候補（未割付・不使用） *)
    E005_In_IN15_2004_10 : UINT;  (* 旧I/O候補（未割付・不使用） *)
    E005_In_IN16_2004_11 : UINT;  (* 旧I/O候補（未割付・不使用） *)
    E005_In_IN17_2004_12 : UINT;  (* 旧I/O候補（未割付・不使用） *)
    E005_In_IN18_2004_13 : UINT;  (* 旧I/O候補（未割付・不使用） *)
    E005_In_IN19_2004_14 : UINT;  (* 旧I/O候補（未割付・不使用） *)
    E005_In_IN20_2004_15 : UINT;  (* 旧I/O候補（未割付・不使用） *)
    E005_In_IN21_2004_16 : UINT;  (* 旧I/O候補（未割付・不使用） *)
    E005_In_IN22_2004_17 : UINT;  (* 旧I/O候補（未割付・不使用） *)
    E005_In_IN23_2004_18 : UINT;  (* 旧I/O候補（未割付・不使用） *)
    E005_In_IN24_2004_19 : UINT;  (* 旧I/O候補（未割付・不使用） *)
    E005_In_IN25_2004_1A : UINT;  (* 旧I/O候補（未割付・不使用） *)
    E005_In_IN26_2004_1B : UINT;  (* 旧I/O候補（未割付・不使用） *)
    E005_In_IN27_2004_1C : UINT;  (* 旧I/O候補（未割付・不使用） *)
    E005_In_IN28_2004_1D : UINT;  (* 旧I/O候補（未割付・不使用） *)
    E005_In_IN29_2004_1E : UINT;  (* 旧I/O候補（未割付・不使用） *)
    E005_In_IN30_2004_1F : UINT;  (* 旧I/O候補（未割付・不使用） *)
    E005_In_IN31_2004_20 : UINT;  (* 旧I/O候補（未割付・不使用） *)
    E005_In_IN32_2004_21 : UINT;  (* 旧I/O候補（未割付・不使用） *)
    E005_In_IN33_2004_22 : UINT;  (* 旧I/O候補（未割付・不使用） *)
    E005_In_IN34_2004_23 : UINT;  (* 旧I/O候補（未割付・不使用） *)
    E005_In_IN35_2004_24 : UINT;  (* 旧I/O候補（未割付・不使用） *)
    E005_In_IN36_2004_25 : UINT;  (* 旧I/O候補（未割付・不使用） *)
    E005_In_IN37_2004_26 : UINT;  (* 旧I/O候補（未割付・不使用） *)
    E005_In_IN38_2004_27 : UINT;  (* 旧I/O候補（未割付・不使用） *)
    E005_In_IN39_2004_28 : UINT;  (* 旧I/O候補（未割付・不使用） *)
    E005_In_IN40_2004_29 : UINT;  (* 旧I/O候補（未割付・不使用） *)
    E005_In_IN41_2004_2A : UINT;  (* 旧I/O候補（未割付・不使用） *)
    E005_In_IN42_2004_2B : UINT;  (* 旧I/O候補（未割付・不使用） *)
    E005_In_IN43_2004_2C : UINT;  (* 旧I/O候補（未割付・不使用） *)
    E005_In_IN44_2004_2D : UINT;  (* 旧I/O候補（未割付・不使用） *)
    E005_In_IN45_2004_2E : UINT;  (* 旧I/O候補（未割付・不使用） *)
    E005_In_IN46_2004_2F : UINT;  (* 旧I/O候補（未割付・不使用） *)
    E005_In_IN47_2004_30 : UINT;  (* 旧I/O候補（未割付・不使用） *)
    E005_In_IN48_2004_31 : UINT;  (* 旧I/O候補（未割付・不使用） *)
    E005_In_IN49_2004_32 : UINT;  (* 旧I/O候補（未割付・不使用） *)
    E005_In_IN50_2004_33 : UINT;  (* 旧I/O候補（未割付・不使用） *)
    E005_In_IN51_2004_34 : UINT;  (* 旧I/O候補（未割付・不使用） *)
    E005_In_IN52_2004_35 : UINT;  (* 旧I/O候補（未割付・不使用） *)
    E005_In_IN53_2004_36 : UINT;  (* 旧I/O候補（未割付・不使用） *)
    E005_In_IN54_2004_37 : UINT;  (* 旧I/O候補（未割付・不使用） *)
    E005_In_IN55_2004_38 : UINT;  (* 旧I/O候補（未割付・不使用） *)
    E005_In_IN56_2004_39 : UINT;  (* 旧I/O候補（未割付・不使用） *)
    E005_In_IN57_2004_3A : UINT;  (* 旧I/O候補（未割付・不使用） *)
    E005_In_IN58_2004_3B : UINT;  (* 旧I/O候補（未割付・不使用） *)
    E005_In_IN59_2004_3C : UINT;  (* 旧I/O候補（未割付・不使用） *)
    E005_In_IN60_2004_3D : UINT;  (* 旧I/O候補（未割付・不使用） *)
    E005_In_IN61_2004_3E : UINT;  (* 旧I/O候補（未割付・不使用） *)
    E005_In_IN62_2004_3F : UINT;  (* 旧I/O候補（未割付・不使用） *)
    E005_In_IN63_2004_40 : UINT;  (* 旧I/O候補（未割付・不使用） *)
    E005_In_IN64_2004_41 : UINT;  (* 旧I/O候補（未割付・不使用） *)
    E005_In_IN65_2004_42 : UINT;  (* 旧I/O候補（未割付・不使用） *)
    E005_In_IN66_2004_43 : UINT;  (* 旧I/O候補（未割付・不使用） *)
    E005_In_IN67_2004_44 : UINT;  (* 旧I/O候補（未割付・不使用） *)
    E005_In_IN68_2004_45 : UINT;  (* 旧I/O候補（未割付・不使用） *)
    E005_In_IN69_2004_46 : UINT;  (* 旧I/O候補（未割付・不使用） *)
    E005_In_IN70_2004_47 : UINT;  (* 旧I/O候補（未割付・不使用） *)
    E005_In_IN71_2004_48 : UINT;  (* 旧I/O候補（未割付・不使用） *)
    E005_Out_OUT00_2003_01_1 : UINT;  (* RCON2 OUT00 共通制御（MON/RTE）; at ECAT://node#5/Out_OUT00_2003_01 *)
    E005_Out_OUT01_2003_02_1 : UINT;  (* RCON2 OUT01 予約（書込禁止）; at ECAT://node#5/Out_OUT01_2003_02 *)
    E005_Out_OUT02_2003_03_1 : UINT;  (* RCON2 OUT02 予約（書込禁止）; at ECAT://node#5/Out_OUT02_2003_03 *)
    E005_Out_OUT03_2003_04_1 : UINT;  (* RCON2 OUT03 予約（書込禁止）; at ECAT://node#5/Out_OUT03_2003_04 *)
    E005_Out_OUT04_2003_05_1 : UINT;  (* RCON2 OUT04 予約（書込禁止）; at ECAT://node#5/Out_OUT04_2003_05 *)
    E005_Out_OUT05_2003_06_1 : UINT;  (* RCON2 OUT05 予約（書込禁止）; at ECAT://node#5/Out_OUT05_2003_06 *)
    E005_Out_OUT06_2003_07_1 : UINT;  (* RCON2 OUT06 予約（書込禁止）; at ECAT://node#5/Out_OUT06_2003_07 *)
    E005_Out_OUT07_2003_08_1 : UINT;  (* RCON2 OUT07 予約（書込禁止）; at ECAT://node#5/Out_OUT07_2003_08 *)
    E005_Out_OUT08_2003_09_1 : UINT;  (* RCON2 OUT08 1軸目 目標位置 下位 [0.01mm]; at ECAT://node#5/Out_OUT08_2003_09 *)
    E005_Out_OUT09_2003_0A_1 : UINT;  (* RCON2 OUT09 1軸目 目標位置 上位 [0.01mm]; at ECAT://node#5/Out_OUT09_2003_0A *)
    E005_Out_OUT10_2003_0B_1 : UINT;  (* RCON2 OUT10 1軸目 位置決め幅 下位 [0.01mm]; at ECAT://node#5/Out_OUT10_2003_0B *)
    E005_Out_OUT11_2003_0C_1 : UINT;  (* RCON2 OUT11 1軸目 位置決め幅 上位 [0.01mm]; at ECAT://node#5/Out_OUT11_2003_0C *)
    E005_Out_OUT12_2003_0D_1 : UINT;  (* RCON2 OUT12 1軸目 速度指令 [実機単位]; at ECAT://node#5/Out_OUT12_2003_0D *)
    E005_Out_OUT13_2003_0E_1 : UINT;  (* RCON2 OUT13 1軸目 共通加減速 [0.01G]; at ECAT://node#5/Out_OUT13_2003_0E *)
    E005_Out_OUT14_2003_0F_1 : UINT;  (* RCON2 OUT14 1軸目 押付け制限 [255=100%]; at ECAT://node#5/Out_OUT14_2003_0F *)
    E005_Out_OUT15_2003_10_1 : UINT;  (* RCON2 OUT15 1軸目 制御信号（DSTR/SON等）; at ECAT://node#5/Out_OUT15_2003_10 *)
    E005_Out_OUT16_2003_11_1 : UINT;  (* RCON2 OUT16 2軸目 目標位置 下位 [0.01mm]; at ECAT://node#5/Out_OUT16_2003_11 *)
    E005_Out_OUT17_2003_12_1 : UINT;  (* RCON2 OUT17 2軸目 目標位置 上位 [0.01mm]; at ECAT://node#5/Out_OUT17_2003_12 *)
    E005_Out_OUT18_2003_13_1 : UINT;  (* RCON2 OUT18 2軸目 位置決め幅 下位 [0.01mm]; at ECAT://node#5/Out_OUT18_2003_13 *)
    E005_Out_OUT19_2003_14_1 : UINT;  (* RCON2 OUT19 2軸目 位置決め幅 上位 [0.01mm]; at ECAT://node#5/Out_OUT19_2003_14 *)
    E005_Out_OUT20_2003_15_1 : UINT;  (* RCON2 OUT20 2軸目 速度指令 [実機単位]; at ECAT://node#5/Out_OUT20_2003_15 *)
    E005_Out_OUT21_2003_16_1 : UINT;  (* RCON2 OUT21 2軸目 共通加減速 [0.01G]; at ECAT://node#5/Out_OUT21_2003_16 *)
    E005_Out_OUT22_2003_17_1 : UINT;  (* RCON2 OUT22 2軸目 押付け制限 [255=100%]; at ECAT://node#5/Out_OUT22_2003_17 *)
    E005_Out_OUT23_2003_18_1 : UINT;  (* RCON2 OUT23 2軸目 制御信号（DSTR/SON等）; at ECAT://node#5/Out_OUT23_2003_18 *)
    E005_Out_OUT24_2003_19_1 : UINT;  (* RCON2 OUT24 3軸目 目標位置 下位 [0.01mm]; at ECAT://node#5/Out_OUT24_2003_19 *)
    E005_Out_OUT25_2003_1A_1 : UINT;  (* RCON2 OUT25 3軸目 目標位置 上位 [0.01mm]; at ECAT://node#5/Out_OUT25_2003_1A *)
    E005_Out_OUT26_2003_1B_1 : UINT;  (* RCON2 OUT26 3軸目 位置決め幅 下位 [0.01mm]; at ECAT://node#5/Out_OUT26_2003_1B *)
    E005_Out_OUT27_2003_1C_1 : UINT;  (* RCON2 OUT27 3軸目 位置決め幅 上位 [0.01mm]; at ECAT://node#5/Out_OUT27_2003_1C *)
    E005_Out_OUT28_2003_1D_1 : UINT;  (* RCON2 OUT28 3軸目 速度指令 [実機単位]; at ECAT://node#5/Out_OUT28_2003_1D *)
    E005_Out_OUT29_2003_1E_1 : UINT;  (* RCON2 OUT29 3軸目 共通加減速 [0.01G]; at ECAT://node#5/Out_OUT29_2003_1E *)
    E005_Out_OUT30_2003_1F_1 : UINT;  (* RCON2 OUT30 3軸目 押付け制限 [255=100%]; at ECAT://node#5/Out_OUT30_2003_1F *)
    E005_Out_OUT31_2003_20_1 : UINT;  (* RCON2 OUT31 3軸目 制御信号（DSTR/SON等）; at ECAT://node#5/Out_OUT31_2003_20 *)
    E005_Out_OUT32_2003_21_1 : UINT;  (* RCON2 OUT32 4軸目 目標位置 下位 [0.01mm]; at ECAT://node#5/Out_OUT32_2003_21 *)
    E005_Out_OUT33_2003_22_1 : UINT;  (* RCON2 OUT33 4軸目 目標位置 上位 [0.01mm]; at ECAT://node#5/Out_OUT33_2003_22 *)
    E005_Out_OUT34_2003_23_1 : UINT;  (* RCON2 OUT34 4軸目 位置決め幅 下位 [0.01mm]; at ECAT://node#5/Out_OUT34_2003_23 *)
    E005_Out_OUT35_2003_24_1 : UINT;  (* RCON2 OUT35 4軸目 位置決め幅 上位 [0.01mm]; at ECAT://node#5/Out_OUT35_2003_24 *)
    E005_Out_OUT36_2003_25_1 : UINT;  (* RCON2 OUT36 4軸目 速度指令 [実機単位]; at ECAT://node#5/Out_OUT36_2003_25 *)
    E005_Out_OUT37_2003_26_1 : UINT;  (* RCON2 OUT37 4軸目 共通加減速 [0.01G]; at ECAT://node#5/Out_OUT37_2003_26 *)
    E005_Out_OUT38_2003_27_1 : UINT;  (* RCON2 OUT38 4軸目 押付け制限 [255=100%]; at ECAT://node#5/Out_OUT38_2003_27 *)
    E005_Out_OUT39_2003_28_1 : UINT;  (* RCON2 OUT39 4軸目 制御信号（DSTR/SON等）; at ECAT://node#5/Out_OUT39_2003_28 *)
    E005_Out_OUT40_2003_29_1 : UINT;  (* RCON2 OUT40 5軸目 目標位置 下位 [0.01mm]; at ECAT://node#5/Out_OUT40_2003_29 *)
    E005_Out_OUT41_2003_2A_1 : UINT;  (* RCON2 OUT41 5軸目 目標位置 上位 [0.01mm]; at ECAT://node#5/Out_OUT41_2003_2A *)
    E005_Out_OUT42_2003_2B_1 : UINT;  (* RCON2 OUT42 5軸目 位置決め幅 下位 [0.01mm]; at ECAT://node#5/Out_OUT42_2003_2B *)
    E005_Out_OUT43_2003_2C_1 : UINT;  (* RCON2 OUT43 5軸目 位置決め幅 上位 [0.01mm]; at ECAT://node#5/Out_OUT43_2003_2C *)
    E005_Out_OUT44_2003_2D_1 : UINT;  (* RCON2 OUT44 5軸目 速度指令 [実機単位]; at ECAT://node#5/Out_OUT44_2003_2D *)
    E005_Out_OUT45_2003_2E_1 : UINT;  (* RCON2 OUT45 5軸目 共通加減速 [0.01G]; at ECAT://node#5/Out_OUT45_2003_2E *)
    E005_Out_OUT46_2003_2F_1 : UINT;  (* RCON2 OUT46 5軸目 押付け制限 [255=100%]; at ECAT://node#5/Out_OUT46_2003_2F *)
    E005_Out_OUT47_2003_30_1 : UINT;  (* RCON2 OUT47 5軸目 制御信号（DSTR/SON等）; at ECAT://node#5/Out_OUT47_2003_30 *)
    E005_Out_OUT48_2003_31_1 : UINT;  (* RCON2 OUT48 用途未確認（今回未使用）; at ECAT://node#5/Out_OUT48_2003_31 *)
    E005_Out_OUT49_2003_32_1 : UINT;  (* RCON2 OUT49 用途未確認（今回未使用）; at ECAT://node#5/Out_OUT49_2003_32 *)
    E005_Out_OUT50_2003_33_1 : UINT;  (* RCON2 OUT50 用途未確認（今回未使用）; at ECAT://node#5/Out_OUT50_2003_33 *)
    E005_Out_OUT51_2003_34_1 : UINT;  (* RCON2 OUT51 用途未確認（今回未使用）; at ECAT://node#5/Out_OUT51_2003_34 *)
    E005_Out_OUT52_2003_35_1 : UINT;  (* RCON2 OUT52 用途未確認（今回未使用）; at ECAT://node#5/Out_OUT52_2003_35 *)
    E005_Out_OUT53_2003_36_1 : UINT;  (* RCON2 OUT53 用途未確認（今回未使用）; at ECAT://node#5/Out_OUT53_2003_36 *)
    E005_Out_OUT54_2003_37_1 : UINT;  (* RCON2 OUT54 用途未確認（今回未使用）; at ECAT://node#5/Out_OUT54_2003_37 *)
    E005_Out_OUT55_2003_38_1 : UINT;  (* RCON2 OUT55 用途未確認（今回未使用）; at ECAT://node#5/Out_OUT55_2003_38 *)
    E005_In_IN00_2004_01_1 : UINT;  (* RCON2 IN00 GW状態; at ECAT://node#5/In_IN00_2004_01 *)
    E005_In_IN01_2004_02_1 : UINT;  (* RCON2 IN01 軸リンク状態; at ECAT://node#5/In_IN01_2004_02 *)
    E005_In_IN02_2004_03_1 : UINT;  (* RCON2 IN02 電源状態0; at ECAT://node#5/In_IN02_2004_03 *)
    E005_In_IN03_2004_04_1 : UINT;  (* RCON2 IN03 電源状態1; at ECAT://node#5/In_IN03_2004_04 *)
    E005_In_IN04_2004_05_1 : UINT;  (* RCON2 IN04 電源状態2; at ECAT://node#5/In_IN04_2004_05 *)
    E005_In_IN05_2004_06_1 : UINT;  (* RCON2 IN05 電源状態3; at ECAT://node#5/In_IN05_2004_06 *)
    E005_In_IN06_2004_07_1 : UINT;  (* RCON2 IN06 電源状態4（構成依存）; at ECAT://node#5/In_IN06_2004_07 *)
    E005_In_IN07_2004_08_1 : UINT;  (* RCON2 IN07 予約（使用禁止）; at ECAT://node#5/In_IN07_2004_08 *)
    E005_In_IN08_2004_09_1 : UINT;  (* RCON2 IN08 1軸目 現在位置 下位 [0.01mm]; at ECAT://node#5/In_IN08_2004_09 *)
    E005_In_IN09_2004_0A_1 : UINT;  (* RCON2 IN09 1軸目 現在位置 上位 [0.01mm]; at ECAT://node#5/In_IN09_2004_0A *)
    E005_In_IN10_2004_0B_1 : UINT;  (* RCON2 IN10 1軸目 指令電流 下位 [mA]; at ECAT://node#5/In_IN10_2004_0B *)
    E005_In_IN11_2004_0C_1 : UINT;  (* RCON2 IN11 1軸目 指令電流 上位 [mA]; at ECAT://node#5/In_IN11_2004_0C *)
    E005_In_IN12_2004_0D_1 : UINT;  (* RCON2 IN12 1軸目 現在速度 [実機単位・符号付き]; at ECAT://node#5/In_IN12_2004_0D *)
    E005_In_IN13_2004_0E_1 : UINT;  (* RCON2 IN13 1軸目 予約（使用禁止）; at ECAT://node#5/In_IN13_2004_0E *)
    E005_In_IN14_2004_0F_1 : UINT;  (* RCON2 IN14 1軸目 軸異常コード; at ECAT://node#5/In_IN14_2004_0F *)
    E005_In_IN15_2004_10_1 : UINT;  (* RCON2 IN15 1軸目 状態信号（PEND/SV等）; at ECAT://node#5/In_IN15_2004_10 *)
    E005_In_IN16_2004_11_1 : UINT;  (* RCON2 IN16 2軸目 現在位置 下位 [0.01mm]; at ECAT://node#5/In_IN16_2004_11 *)
    E005_In_IN17_2004_12_1 : UINT;  (* RCON2 IN17 2軸目 現在位置 上位 [0.01mm]; at ECAT://node#5/In_IN17_2004_12 *)
    E005_In_IN18_2004_13_1 : UINT;  (* RCON2 IN18 2軸目 指令電流 下位 [mA]; at ECAT://node#5/In_IN18_2004_13 *)
    E005_In_IN19_2004_14_1 : UINT;  (* RCON2 IN19 2軸目 指令電流 上位 [mA]; at ECAT://node#5/In_IN19_2004_14 *)
    E005_In_IN20_2004_15_1 : UINT;  (* RCON2 IN20 2軸目 現在速度 [実機単位・符号付き]; at ECAT://node#5/In_IN20_2004_15 *)
    E005_In_IN21_2004_16_1 : UINT;  (* RCON2 IN21 2軸目 予約（使用禁止）; at ECAT://node#5/In_IN21_2004_16 *)
    E005_In_IN22_2004_17_1 : UINT;  (* RCON2 IN22 2軸目 軸異常コード; at ECAT://node#5/In_IN22_2004_17 *)
    E005_In_IN23_2004_18_1 : UINT;  (* RCON2 IN23 2軸目 状態信号（PEND/SV等）; at ECAT://node#5/In_IN23_2004_18 *)
    E005_In_IN24_2004_19_1 : UINT;  (* RCON2 IN24 3軸目 現在位置 下位 [0.01mm]; at ECAT://node#5/In_IN24_2004_19 *)
    E005_In_IN25_2004_1A_1 : UINT;  (* RCON2 IN25 3軸目 現在位置 上位 [0.01mm]; at ECAT://node#5/In_IN25_2004_1A *)
    E005_In_IN26_2004_1B_1 : UINT;  (* RCON2 IN26 3軸目 指令電流 下位 [mA]; at ECAT://node#5/In_IN26_2004_1B *)
    E005_In_IN27_2004_1C_1 : UINT;  (* RCON2 IN27 3軸目 指令電流 上位 [mA]; at ECAT://node#5/In_IN27_2004_1C *)
    E005_In_IN28_2004_1D_1 : UINT;  (* RCON2 IN28 3軸目 現在速度 [実機単位・符号付き]; at ECAT://node#5/In_IN28_2004_1D *)
    E005_In_IN29_2004_1E_1 : UINT;  (* RCON2 IN29 3軸目 予約（使用禁止）; at ECAT://node#5/In_IN29_2004_1E *)
    E005_In_IN30_2004_1F_1 : UINT;  (* RCON2 IN30 3軸目 軸異常コード; at ECAT://node#5/In_IN30_2004_1F *)
    E005_In_IN31_2004_20_1 : UINT;  (* RCON2 IN31 3軸目 状態信号（PEND/SV等）; at ECAT://node#5/In_IN31_2004_20 *)
    E005_In_IN32_2004_21_1 : UINT;  (* RCON2 IN32 4軸目 現在位置 下位 [0.01mm]; at ECAT://node#5/In_IN32_2004_21 *)
    E005_In_IN33_2004_22_1 : UINT;  (* RCON2 IN33 4軸目 現在位置 上位 [0.01mm]; at ECAT://node#5/In_IN33_2004_22 *)
    E005_In_IN34_2004_23_1 : UINT;  (* RCON2 IN34 4軸目 指令電流 下位 [mA]; at ECAT://node#5/In_IN34_2004_23 *)
    E005_In_IN35_2004_24_1 : UINT;  (* RCON2 IN35 4軸目 指令電流 上位 [mA]; at ECAT://node#5/In_IN35_2004_24 *)
    E005_In_IN36_2004_25_1 : UINT;  (* RCON2 IN36 4軸目 現在速度 [実機単位・符号付き]; at ECAT://node#5/In_IN36_2004_25 *)
    E005_In_IN37_2004_26_1 : UINT;  (* RCON2 IN37 4軸目 予約（使用禁止）; at ECAT://node#5/In_IN37_2004_26 *)
    E005_In_IN38_2004_27_1 : UINT;  (* RCON2 IN38 4軸目 軸異常コード; at ECAT://node#5/In_IN38_2004_27 *)
    E005_In_IN39_2004_28_1 : UINT;  (* RCON2 IN39 4軸目 状態信号（PEND/SV等）; at ECAT://node#5/In_IN39_2004_28 *)
    E005_In_IN40_2004_29_1 : UINT;  (* RCON2 IN40 5軸目 現在位置 下位 [0.01mm]; at ECAT://node#5/In_IN40_2004_29 *)
    E005_In_IN41_2004_2A_1 : UINT;  (* RCON2 IN41 5軸目 現在位置 上位 [0.01mm]; at ECAT://node#5/In_IN41_2004_2A *)
    E005_In_IN42_2004_2B_1 : UINT;  (* RCON2 IN42 5軸目 指令電流 下位 [mA]; at ECAT://node#5/In_IN42_2004_2B *)
    E005_In_IN43_2004_2C_1 : UINT;  (* RCON2 IN43 5軸目 指令電流 上位 [mA]; at ECAT://node#5/In_IN43_2004_2C *)
    E005_In_IN44_2004_2D_1 : UINT;  (* RCON2 IN44 5軸目 現在速度 [実機単位・符号付き]; at ECAT://node#5/In_IN44_2004_2D *)
    E005_In_IN45_2004_2E_1 : UINT;  (* RCON2 IN45 5軸目 予約（使用禁止）; at ECAT://node#5/In_IN45_2004_2E *)
    E005_In_IN46_2004_2F_1 : UINT;  (* RCON2 IN46 5軸目 軸異常コード; at ECAT://node#5/In_IN46_2004_2F *)
    E005_In_IN47_2004_30_1 : UINT;  (* RCON2 IN47 5軸目 状態信号（PEND/SV等）; at ECAT://node#5/In_IN47_2004_30 *)
    E005_In_IN48_2004_31_1 : UINT;  (* RCON2 IN48 用途未確認（今回未使用）; at ECAT://node#5/In_IN48_2004_31 *)
    E005_In_IN49_2004_32_1 : UINT;  (* RCON2 IN49 用途未確認（今回未使用）; at ECAT://node#5/In_IN49_2004_32 *)
    E005_In_IN50_2004_33_1 : UINT;  (* RCON2 IN50 用途未確認（今回未使用）; at ECAT://node#5/In_IN50_2004_33 *)
    E005_In_IN51_2004_34_1 : UINT;  (* RCON2 IN51 用途未確認（今回未使用）; at ECAT://node#5/In_IN51_2004_34 *)
    E005_In_IN52_2004_35_1 : UINT;  (* RCON2 IN52 用途未確認（今回未使用）; at ECAT://node#5/In_IN52_2004_35 *)
    E005_In_IN53_2004_36_1 : UINT;  (* RCON2 IN53 用途未確認（今回未使用）; at ECAT://node#5/In_IN53_2004_36 *)
    E005_In_IN54_2004_37_1 : UINT;  (* RCON2 IN54 用途未確認（今回未使用）; at ECAT://node#5/In_IN54_2004_37 *)
    E005_In_IN55_2004_38_1 : UINT;  (* RCON2 IN55 用途未確認（今回未使用）; at ECAT://node#5/In_IN55_2004_38 *)
    E001_Out_OUT00_2003_01 : UINT;  (* RCON1 OUT00 共通制御（MON/RTE）; at ECAT://node#1/Out_OUT00_2003_01 *)
    E001_Out_OUT01_2003_02 : UINT;  (* RCON1 OUT01 予約（書込禁止）; at ECAT://node#1/Out_OUT01_2003_02 *)
    E001_Out_OUT02_2003_03 : UINT;  (* RCON1 OUT02 予約（書込禁止）; at ECAT://node#1/Out_OUT02_2003_03 *)
    E001_Out_OUT03_2003_04 : UINT;  (* RCON1 OUT03 予約（書込禁止）; at ECAT://node#1/Out_OUT03_2003_04 *)
    E001_Out_OUT04_2003_05 : UINT;  (* RCON1 OUT04 予約（書込禁止）; at ECAT://node#1/Out_OUT04_2003_05 *)
    E001_Out_OUT05_2003_06 : UINT;  (* RCON1 OUT05 予約（書込禁止）; at ECAT://node#1/Out_OUT05_2003_06 *)
    E001_Out_OUT06_2003_07 : UINT;  (* RCON1 OUT06 予約（書込禁止）; at ECAT://node#1/Out_OUT06_2003_07 *)
    E001_Out_OUT07_2003_08 : UINT;  (* RCON1 OUT07 予約（書込禁止）; at ECAT://node#1/Out_OUT07_2003_08 *)
    E001_Out_OUT08_2003_09 : UINT;  (* RCON1 OUT08 1軸目 目標位置 下位 [0.01mm]; at ECAT://node#1/Out_OUT08_2003_09 *)
    E001_Out_OUT09_2003_0A : UINT;  (* RCON1 OUT09 1軸目 目標位置 上位 [0.01mm]; at ECAT://node#1/Out_OUT09_2003_0A *)
    E001_Out_OUT10_2003_0B : UINT;  (* RCON1 OUT10 1軸目 位置決め幅 下位 [0.01mm]; at ECAT://node#1/Out_OUT10_2003_0B *)
    E001_Out_OUT11_2003_0C : UINT;  (* RCON1 OUT11 1軸目 位置決め幅 上位 [0.01mm]; at ECAT://node#1/Out_OUT11_2003_0C *)
    E001_Out_OUT12_2003_0D : UINT;  (* RCON1 OUT12 1軸目 速度指令 [実機単位]; at ECAT://node#1/Out_OUT12_2003_0D *)
    E001_Out_OUT13_2003_0E : UINT;  (* RCON1 OUT13 1軸目 共通加減速 [0.01G]; at ECAT://node#1/Out_OUT13_2003_0E *)
    E001_Out_OUT14_2003_0F : UINT;  (* RCON1 OUT14 1軸目 押付け制限 [255=100%]; at ECAT://node#1/Out_OUT14_2003_0F *)
    E001_Out_OUT15_2003_10 : UINT;  (* RCON1 OUT15 1軸目 制御信号（DSTR/SON等）; at ECAT://node#1/Out_OUT15_2003_10 *)
    E001_Out_OUT16_2003_11 : UINT;  (* RCON1 OUT16 2軸目 目標位置 下位 [0.01mm]; at ECAT://node#1/Out_OUT16_2003_11 *)
    E001_Out_OUT17_2003_12 : UINT;  (* RCON1 OUT17 2軸目 目標位置 上位 [0.01mm]; at ECAT://node#1/Out_OUT17_2003_12 *)
    E001_Out_OUT18_2003_13 : UINT;  (* RCON1 OUT18 2軸目 位置決め幅 下位 [0.01mm]; at ECAT://node#1/Out_OUT18_2003_13 *)
    E001_Out_OUT19_2003_14 : UINT;  (* RCON1 OUT19 2軸目 位置決め幅 上位 [0.01mm]; at ECAT://node#1/Out_OUT19_2003_14 *)
    E001_Out_OUT20_2003_15 : UINT;  (* RCON1 OUT20 2軸目 速度指令 [実機単位]; at ECAT://node#1/Out_OUT20_2003_15 *)
    E001_Out_OUT21_2003_16 : UINT;  (* RCON1 OUT21 2軸目 共通加減速 [0.01G]; at ECAT://node#1/Out_OUT21_2003_16 *)
    E001_Out_OUT22_2003_17 : UINT;  (* RCON1 OUT22 2軸目 押付け制限 [255=100%]; at ECAT://node#1/Out_OUT22_2003_17 *)
    E001_Out_OUT23_2003_18 : UINT;  (* RCON1 OUT23 2軸目 制御信号（DSTR/SON等）; at ECAT://node#1/Out_OUT23_2003_18 *)
    E001_Out_OUT24_2003_19 : UINT;  (* RCON1 OUT24 3軸目 目標位置 下位 [0.01mm]; at ECAT://node#1/Out_OUT24_2003_19 *)
    E001_Out_OUT25_2003_1A : UINT;  (* RCON1 OUT25 3軸目 目標位置 上位 [0.01mm]; at ECAT://node#1/Out_OUT25_2003_1A *)
    E001_Out_OUT26_2003_1B : UINT;  (* RCON1 OUT26 3軸目 位置決め幅 下位 [0.01mm]; at ECAT://node#1/Out_OUT26_2003_1B *)
    E001_Out_OUT27_2003_1C : UINT;  (* RCON1 OUT27 3軸目 位置決め幅 上位 [0.01mm]; at ECAT://node#1/Out_OUT27_2003_1C *)
    E001_Out_OUT28_2003_1D : UINT;  (* RCON1 OUT28 3軸目 速度指令 [実機単位]; at ECAT://node#1/Out_OUT28_2003_1D *)
    E001_Out_OUT29_2003_1E : UINT;  (* RCON1 OUT29 3軸目 共通加減速 [0.01G]; at ECAT://node#1/Out_OUT29_2003_1E *)
    E001_Out_OUT30_2003_1F : UINT;  (* RCON1 OUT30 3軸目 押付け制限 [255=100%]; at ECAT://node#1/Out_OUT30_2003_1F *)
    E001_Out_OUT31_2003_20 : UINT;  (* RCON1 OUT31 3軸目 制御信号（DSTR/SON等）; at ECAT://node#1/Out_OUT31_2003_20 *)
    E001_Out_OUT32_2003_21 : UINT;  (* RCON1 OUT32 4軸目 目標位置 下位 [0.01mm]; at ECAT://node#1/Out_OUT32_2003_21 *)
    E001_Out_OUT33_2003_22 : UINT;  (* RCON1 OUT33 4軸目 目標位置 上位 [0.01mm]; at ECAT://node#1/Out_OUT33_2003_22 *)
    E001_Out_OUT34_2003_23 : UINT;  (* RCON1 OUT34 4軸目 位置決め幅 下位 [0.01mm]; at ECAT://node#1/Out_OUT34_2003_23 *)
    E001_Out_OUT35_2003_24 : UINT;  (* RCON1 OUT35 4軸目 位置決め幅 上位 [0.01mm]; at ECAT://node#1/Out_OUT35_2003_24 *)
    E001_Out_OUT36_2003_25 : UINT;  (* RCON1 OUT36 4軸目 速度指令 [実機単位]; at ECAT://node#1/Out_OUT36_2003_25 *)
    E001_Out_OUT37_2003_26 : UINT;  (* RCON1 OUT37 4軸目 共通加減速 [0.01G]; at ECAT://node#1/Out_OUT37_2003_26 *)
    E001_Out_OUT38_2003_27 : UINT;  (* RCON1 OUT38 4軸目 押付け制限 [255=100%]; at ECAT://node#1/Out_OUT38_2003_27 *)
    E001_Out_OUT39_2003_28 : UINT;  (* RCON1 OUT39 4軸目 制御信号（DSTR/SON等）; at ECAT://node#1/Out_OUT39_2003_28 *)
    E001_Out_OUT40_2003_29 : UINT;  (* RCON1 OUT40 5軸目 目標位置 下位 [0.01mm]; at ECAT://node#1/Out_OUT40_2003_29 *)
    E001_Out_OUT41_2003_2A : UINT;  (* RCON1 OUT41 5軸目 目標位置 上位 [0.01mm]; at ECAT://node#1/Out_OUT41_2003_2A *)
    E001_Out_OUT42_2003_2B : UINT;  (* RCON1 OUT42 5軸目 位置決め幅 下位 [0.01mm]; at ECAT://node#1/Out_OUT42_2003_2B *)
    E001_Out_OUT43_2003_2C : UINT;  (* RCON1 OUT43 5軸目 位置決め幅 上位 [0.01mm]; at ECAT://node#1/Out_OUT43_2003_2C *)
    E001_Out_OUT44_2003_2D : UINT;  (* RCON1 OUT44 5軸目 速度指令 [実機単位]; at ECAT://node#1/Out_OUT44_2003_2D *)
    E001_Out_OUT45_2003_2E : UINT;  (* RCON1 OUT45 5軸目 共通加減速 [0.01G]; at ECAT://node#1/Out_OUT45_2003_2E *)
    E001_Out_OUT46_2003_2F : UINT;  (* RCON1 OUT46 5軸目 押付け制限 [255=100%]; at ECAT://node#1/Out_OUT46_2003_2F *)
    E001_Out_OUT47_2003_30 : UINT;  (* RCON1 OUT47 5軸目 制御信号（DSTR/SON等）; at ECAT://node#1/Out_OUT47_2003_30 *)
    E001_Out_OUT48_2003_31 : UINT;  (* RCON1 OUT48 6軸目 目標位置 下位 [0.01mm]; at ECAT://node#1/Out_OUT48_2003_31 *)
    E001_Out_OUT49_2003_32 : UINT;  (* RCON1 OUT49 6軸目 目標位置 上位 [0.01mm]; at ECAT://node#1/Out_OUT49_2003_32 *)
    E001_Out_OUT50_2003_33 : UINT;  (* RCON1 OUT50 6軸目 位置決め幅 下位 [0.01mm]; at ECAT://node#1/Out_OUT50_2003_33 *)
    E001_Out_OUT51_2003_34 : UINT;  (* RCON1 OUT51 6軸目 位置決め幅 上位 [0.01mm]; at ECAT://node#1/Out_OUT51_2003_34 *)
    E001_Out_OUT52_2003_35 : UINT;  (* RCON1 OUT52 6軸目 速度指令 [実機単位]; at ECAT://node#1/Out_OUT52_2003_35 *)
    E001_Out_OUT53_2003_36 : UINT;  (* RCON1 OUT53 6軸目 共通加減速 [0.01G]; at ECAT://node#1/Out_OUT53_2003_36 *)
    E001_Out_OUT54_2003_37 : UINT;  (* RCON1 OUT54 6軸目 押付け制限 [255=100%]; at ECAT://node#1/Out_OUT54_2003_37 *)
    E001_Out_OUT55_2003_38 : UINT;  (* RCON1 OUT55 6軸目 制御信号（DSTR/SON等）; at ECAT://node#1/Out_OUT55_2003_38 *)
    E001_Out_OUT56_2003_39 : UINT;  (* RCON1 OUT56 用途未確認（今回未使用）; at ECAT://node#1/Out_OUT56_2003_39 *)
    E001_Out_OUT57_2003_3A : UINT;  (* RCON1 OUT57 用途未確認（今回未使用）; at ECAT://node#1/Out_OUT57_2003_3A *)
    E001_Out_OUT58_2003_3B : UINT;  (* RCON1 OUT58 用途未確認（今回未使用）; at ECAT://node#1/Out_OUT58_2003_3B *)
    E001_Out_OUT59_2003_3C : UINT;  (* RCON1 OUT59 用途未確認（今回未使用）; at ECAT://node#1/Out_OUT59_2003_3C *)
    E001_Out_OUT60_2003_3D : UINT;  (* RCON1 OUT60 用途未確認（今回未使用）; at ECAT://node#1/Out_OUT60_2003_3D *)
    E001_Out_OUT61_2003_3E : UINT;  (* RCON1 OUT61 用途未確認（今回未使用）; at ECAT://node#1/Out_OUT61_2003_3E *)
    E001_Out_OUT62_2003_3F : UINT;  (* RCON1 OUT62 用途未確認（今回未使用）; at ECAT://node#1/Out_OUT62_2003_3F *)
    E001_Out_OUT63_2003_40 : UINT;  (* RCON1 OUT63 用途未確認（今回未使用）; at ECAT://node#1/Out_OUT63_2003_40 *)
    E001_Out_OUT64_2003_41 : UINT;  (* RCON1 OUT64 用途未確認（今回未使用）; at ECAT://node#1/Out_OUT64_2003_41 *)
    E001_Out_OUT65_2003_42 : UINT;  (* RCON1 OUT65 用途未確認（今回未使用）; at ECAT://node#1/Out_OUT65_2003_42 *)
    E001_Out_OUT66_2003_43 : UINT;  (* RCON1 OUT66 用途未確認（今回未使用）; at ECAT://node#1/Out_OUT66_2003_43 *)
    E001_Out_OUT67_2003_44 : UINT;  (* RCON1 OUT67 用途未確認（今回未使用）; at ECAT://node#1/Out_OUT67_2003_44 *)
    E001_Out_OUT68_2003_45 : UINT;  (* RCON1 OUT68 用途未確認（今回未使用）; at ECAT://node#1/Out_OUT68_2003_45 *)
    E001_Out_OUT69_2003_46 : UINT;  (* RCON1 OUT69 用途未確認（今回未使用）; at ECAT://node#1/Out_OUT69_2003_46 *)
    E001_Out_OUT70_2003_47 : UINT;  (* RCON1 OUT70 用途未確認（今回未使用）; at ECAT://node#1/Out_OUT70_2003_47 *)
    E001_Out_OUT71_2003_48 : UINT;  (* RCON1 OUT71 用途未確認（今回未使用）; at ECAT://node#1/Out_OUT71_2003_48 *)
    E001_In_IN00_2004_01 : UINT;  (* RCON1 IN00 GW状態; at ECAT://node#1/In_IN00_2004_01 *)
    E001_In_IN01_2004_02 : UINT;  (* RCON1 IN01 軸リンク状態; at ECAT://node#1/In_IN01_2004_02 *)
    E001_In_IN02_2004_03 : UINT;  (* RCON1 IN02 電源状態0; at ECAT://node#1/In_IN02_2004_03 *)
    E001_In_IN03_2004_04 : UINT;  (* RCON1 IN03 電源状態1; at ECAT://node#1/In_IN03_2004_04 *)
    E001_In_IN04_2004_05 : UINT;  (* RCON1 IN04 電源状態2; at ECAT://node#1/In_IN04_2004_05 *)
    E001_In_IN05_2004_06 : UINT;  (* RCON1 IN05 電源状態3; at ECAT://node#1/In_IN05_2004_06 *)
    E001_In_IN06_2004_07 : UINT;  (* RCON1 IN06 電源状態4（構成依存）; at ECAT://node#1/In_IN06_2004_07 *)
    E001_In_IN07_2004_08 : UINT;  (* RCON1 IN07 予約（使用禁止）; at ECAT://node#1/In_IN07_2004_08 *)
    E001_In_IN08_2004_09 : UINT;  (* RCON1 IN08 1軸目 現在位置 下位 [0.01mm]; at ECAT://node#1/In_IN08_2004_09 *)
    E001_In_IN09_2004_0A : UINT;  (* RCON1 IN09 1軸目 現在位置 上位 [0.01mm]; at ECAT://node#1/In_IN09_2004_0A *)
    E001_In_IN10_2004_0B : UINT;  (* RCON1 IN10 1軸目 指令電流 下位 [mA]; at ECAT://node#1/In_IN10_2004_0B *)
    E001_In_IN11_2004_0C : UINT;  (* RCON1 IN11 1軸目 指令電流 上位 [mA]; at ECAT://node#1/In_IN11_2004_0C *)
    E001_In_IN12_2004_0D : UINT;  (* RCON1 IN12 1軸目 現在速度 [実機単位・符号付き]; at ECAT://node#1/In_IN12_2004_0D *)
    E001_In_IN13_2004_0E : UINT;  (* RCON1 IN13 1軸目 予約（使用禁止）; at ECAT://node#1/In_IN13_2004_0E *)
    E001_In_IN14_2004_0F : UINT;  (* RCON1 IN14 1軸目 軸異常コード; at ECAT://node#1/In_IN14_2004_0F *)
    E001_In_IN15_2004_10 : UINT;  (* RCON1 IN15 1軸目 状態信号（PEND/SV等）; at ECAT://node#1/In_IN15_2004_10 *)
    E001_In_IN16_2004_11 : UINT;  (* RCON1 IN16 2軸目 現在位置 下位 [0.01mm]; at ECAT://node#1/In_IN16_2004_11 *)
    E001_In_IN17_2004_12 : UINT;  (* RCON1 IN17 2軸目 現在位置 上位 [0.01mm]; at ECAT://node#1/In_IN17_2004_12 *)
    E001_In_IN18_2004_13 : UINT;  (* RCON1 IN18 2軸目 指令電流 下位 [mA]; at ECAT://node#1/In_IN18_2004_13 *)
    E001_In_IN19_2004_14 : UINT;  (* RCON1 IN19 2軸目 指令電流 上位 [mA]; at ECAT://node#1/In_IN19_2004_14 *)
    E001_In_IN20_2004_15 : UINT;  (* RCON1 IN20 2軸目 現在速度 [実機単位・符号付き]; at ECAT://node#1/In_IN20_2004_15 *)
    E001_In_IN21_2004_16 : UINT;  (* RCON1 IN21 2軸目 予約（使用禁止）; at ECAT://node#1/In_IN21_2004_16 *)
    E001_In_IN22_2004_17 : UINT;  (* RCON1 IN22 2軸目 軸異常コード; at ECAT://node#1/In_IN22_2004_17 *)
    E001_In_IN23_2004_18 : UINT;  (* RCON1 IN23 2軸目 状態信号（PEND/SV等）; at ECAT://node#1/In_IN23_2004_18 *)
    E001_In_IN24_2004_19 : UINT;  (* RCON1 IN24 3軸目 現在位置 下位 [0.01mm]; at ECAT://node#1/In_IN24_2004_19 *)
    E001_In_IN25_2004_1A : UINT;  (* RCON1 IN25 3軸目 現在位置 上位 [0.01mm]; at ECAT://node#1/In_IN25_2004_1A *)
    E001_In_IN26_2004_1B : UINT;  (* RCON1 IN26 3軸目 指令電流 下位 [mA]; at ECAT://node#1/In_IN26_2004_1B *)
    E001_In_IN27_2004_1C : UINT;  (* RCON1 IN27 3軸目 指令電流 上位 [mA]; at ECAT://node#1/In_IN27_2004_1C *)
    E001_In_IN28_2004_1D : UINT;  (* RCON1 IN28 3軸目 現在速度 [実機単位・符号付き]; at ECAT://node#1/In_IN28_2004_1D *)
    E001_In_IN29_2004_1E : UINT;  (* RCON1 IN29 3軸目 予約（使用禁止）; at ECAT://node#1/In_IN29_2004_1E *)
    E001_In_IN30_2004_1F : UINT;  (* RCON1 IN30 3軸目 軸異常コード; at ECAT://node#1/In_IN30_2004_1F *)
    E001_In_IN31_2004_20 : UINT;  (* RCON1 IN31 3軸目 状態信号（PEND/SV等）; at ECAT://node#1/In_IN31_2004_20 *)
    E001_In_IN32_2004_21 : UINT;  (* RCON1 IN32 4軸目 現在位置 下位 [0.01mm]; at ECAT://node#1/In_IN32_2004_21 *)
    E001_In_IN33_2004_22 : UINT;  (* RCON1 IN33 4軸目 現在位置 上位 [0.01mm]; at ECAT://node#1/In_IN33_2004_22 *)
    E001_In_IN34_2004_23 : UINT;  (* RCON1 IN34 4軸目 指令電流 下位 [mA]; at ECAT://node#1/In_IN34_2004_23 *)
    E001_In_IN35_2004_24 : UINT;  (* RCON1 IN35 4軸目 指令電流 上位 [mA]; at ECAT://node#1/In_IN35_2004_24 *)
    E001_In_IN36_2004_25 : UINT;  (* RCON1 IN36 4軸目 現在速度 [実機単位・符号付き]; at ECAT://node#1/In_IN36_2004_25 *)
    E001_In_IN37_2004_26 : UINT;  (* RCON1 IN37 4軸目 予約（使用禁止）; at ECAT://node#1/In_IN37_2004_26 *)
    E001_In_IN38_2004_27 : UINT;  (* RCON1 IN38 4軸目 軸異常コード; at ECAT://node#1/In_IN38_2004_27 *)
    E001_In_IN39_2004_28 : UINT;  (* RCON1 IN39 4軸目 状態信号（PEND/SV等）; at ECAT://node#1/In_IN39_2004_28 *)
    E001_In_IN40_2004_29 : UINT;  (* RCON1 IN40 5軸目 現在位置 下位 [0.01mm]; at ECAT://node#1/In_IN40_2004_29 *)
    E001_In_IN41_2004_2A : UINT;  (* RCON1 IN41 5軸目 現在位置 上位 [0.01mm]; at ECAT://node#1/In_IN41_2004_2A *)
    E001_In_IN42_2004_2B : UINT;  (* RCON1 IN42 5軸目 指令電流 下位 [mA]; at ECAT://node#1/In_IN42_2004_2B *)
    E001_In_IN43_2004_2C : UINT;  (* RCON1 IN43 5軸目 指令電流 上位 [mA]; at ECAT://node#1/In_IN43_2004_2C *)
    E001_In_IN44_2004_2D : UINT;  (* RCON1 IN44 5軸目 現在速度 [実機単位・符号付き]; at ECAT://node#1/In_IN44_2004_2D *)
    E001_In_IN45_2004_2E : UINT;  (* RCON1 IN45 5軸目 予約（使用禁止）; at ECAT://node#1/In_IN45_2004_2E *)
    E001_In_IN46_2004_2F : UINT;  (* RCON1 IN46 5軸目 軸異常コード; at ECAT://node#1/In_IN46_2004_2F *)
    E001_In_IN47_2004_30 : UINT;  (* RCON1 IN47 5軸目 状態信号（PEND/SV等）; at ECAT://node#1/In_IN47_2004_30 *)
    E001_In_IN48_2004_31 : UINT;  (* RCON1 IN48 6軸目 現在位置 下位 [0.01mm]; at ECAT://node#1/In_IN48_2004_31 *)
    E001_In_IN49_2004_32 : UINT;  (* RCON1 IN49 6軸目 現在位置 上位 [0.01mm]; at ECAT://node#1/In_IN49_2004_32 *)
    E001_In_IN50_2004_33 : UINT;  (* RCON1 IN50 6軸目 指令電流 下位 [mA]; at ECAT://node#1/In_IN50_2004_33 *)
    E001_In_IN51_2004_34 : UINT;  (* RCON1 IN51 6軸目 指令電流 上位 [mA]; at ECAT://node#1/In_IN51_2004_34 *)
    E001_In_IN52_2004_35 : UINT;  (* RCON1 IN52 6軸目 現在速度 [実機単位・符号付き]; at ECAT://node#1/In_IN52_2004_35 *)
    E001_In_IN53_2004_36 : UINT;  (* RCON1 IN53 6軸目 予約（使用禁止）; at ECAT://node#1/In_IN53_2004_36 *)
    E001_In_IN54_2004_37 : UINT;  (* RCON1 IN54 6軸目 軸異常コード; at ECAT://node#1/In_IN54_2004_37 *)
    E001_In_IN55_2004_38 : UINT;  (* RCON1 IN55 6軸目 状態信号（PEND/SV等）; at ECAT://node#1/In_IN55_2004_38 *)
    E001_In_IN56_2004_39 : UINT;  (* RCON1 IN56 用途未確認（今回未使用）; at ECAT://node#1/In_IN56_2004_39 *)
    E001_In_IN57_2004_3A : UINT;  (* RCON1 IN57 用途未確認（今回未使用）; at ECAT://node#1/In_IN57_2004_3A *)
    E001_In_IN58_2004_3B : UINT;  (* RCON1 IN58 用途未確認（今回未使用）; at ECAT://node#1/In_IN58_2004_3B *)
    E001_In_IN59_2004_3C : UINT;  (* RCON1 IN59 用途未確認（今回未使用）; at ECAT://node#1/In_IN59_2004_3C *)
    E001_In_IN60_2004_3D : UINT;  (* RCON1 IN60 用途未確認（今回未使用）; at ECAT://node#1/In_IN60_2004_3D *)
    E001_In_IN61_2004_3E : UINT;  (* RCON1 IN61 用途未確認（今回未使用）; at ECAT://node#1/In_IN61_2004_3E *)
    E001_In_IN62_2004_3F : UINT;  (* RCON1 IN62 用途未確認（今回未使用）; at ECAT://node#1/In_IN62_2004_3F *)
    E001_In_IN63_2004_40 : UINT;  (* RCON1 IN63 用途未確認（今回未使用）; at ECAT://node#1/In_IN63_2004_40 *)
    E001_In_IN64_2004_41 : UINT;  (* RCON1 IN64 用途未確認（今回未使用）; at ECAT://node#1/In_IN64_2004_41 *)
    E001_In_IN65_2004_42 : UINT;  (* RCON1 IN65 用途未確認（今回未使用）; at ECAT://node#1/In_IN65_2004_42 *)
    E001_In_IN66_2004_43 : UINT;  (* RCON1 IN66 用途未確認（今回未使用）; at ECAT://node#1/In_IN66_2004_43 *)
    E001_In_IN67_2004_44 : UINT;  (* RCON1 IN67 用途未確認（今回未使用）; at ECAT://node#1/In_IN67_2004_44 *)
    E001_In_IN68_2004_45 : UINT;  (* RCON1 IN68 用途未確認（今回未使用）; at ECAT://node#1/In_IN68_2004_45 *)
    E001_In_IN69_2004_46 : UINT;  (* RCON1 IN69 用途未確認（今回未使用）; at ECAT://node#1/In_IN69_2004_46 *)
    E001_In_IN70_2004_47 : UINT;  (* RCON1 IN70 用途未確認（今回未使用）; at ECAT://node#1/In_IN70_2004_47 *)
    E001_In_IN71_2004_48 : UINT;  (* RCON1 IN71 用途未確認（今回未使用）; at ECAT://node#1/In_IN71_2004_48 *)
    RCON1_RxRaw : ARRAY[0..71] OF UINT;  (* RCON1 受信値（バイト交換前）; [0] IN00 GW状態; [1] IN01 軸リンク状態; [2] IN02 電源状態0; [3] IN03 電源状態1; [4] IN04 電源状態2; [5] IN05 電源状態3; [6] IN06 電源状態4（構成依存）; [7] IN07 予約（使用禁止）; [8] IN08 1軸目 現在位置 下位 [0.01mm]; [9] IN09 1軸目 現在位置 上位 [0.01mm]; [10] IN10 1軸目 指令電流 下位 [mA]; [11] IN11 1軸目 指令電流 上位 [mA]; [12] IN12 1軸目 現在速度 [実機単位・符号付き]; [13] IN13 1軸目 予約（使用禁止）; [14] IN14 1軸目 軸異常コード; [15] IN15 1軸目 状態信号（PEND/SV等）; [16] IN16 2軸目 現在位置 下位 [0.01mm]; [17] IN17 2軸目 現在位置 上位 [0.01mm]; [18] IN18 2軸目 指令電流 下位 [mA]; [19] IN19 2軸目 指令電流 上位 [mA]; [20] IN20 2軸目 現在速度 [実機単位・符号付き]; [21] IN21 2軸目 予約（使用禁止）; [22] IN22 2軸目 軸異常コード; [23] IN23 2軸目 状態信号（PEND/SV等）; [24] IN24 3軸目 現在位置 下位 [0.01mm]; [25] IN25 3軸目 現在位置 上位 [0.01mm]; [26] IN26 3軸目 指令電流 下位 [mA]; [27] IN27 3軸目 指令電流 上位 [mA]; [28] IN28 3軸目 現在速度 [実機単位・符号付き]; [29] IN29 3軸目 予約（使用禁止）; [30] IN30 3軸目 軸異常コード; [31] IN31 3軸目 状態信号（PEND/SV等）; [32] IN32 4軸目 現在位置 下位 [0.01mm]; [33] IN33 4軸目 現在位置 上位 [0.01mm]; [34] IN34 4軸目 指令電流 下位 [mA]; [35] IN35 4軸目 指令電流 上位 [mA]; [36] IN36 4軸目 現在速度 [実機単位・符号付き]; [37] IN37 4軸目 予約（使用禁止）; [38] IN38 4軸目 軸異常コード; [39] IN39 4軸目 状態信号（PEND/SV等）; [40] IN40 5軸目 現在位置 下位 [0.01mm]; [41] IN41 5軸目 現在位置 上位 [0.01mm]; [42] IN42 5軸目 指令電流 下位 [mA]; [43] IN43 5軸目 指令電流 上位 [mA]; [44] IN44 5軸目 現在速度 [実機単位・符号付き]; [45] IN45 5軸目 予約（使用禁止）; [46] IN46 5軸目 軸異常コード; [47] IN47 5軸目 状態信号（PEND/SV等）; [48] IN48 6軸目 現在位置 下位 [0.01mm]; [49] IN49 6軸目 現在位置 上位 [0.01mm]; [50] IN50 6軸目 指令電流 下位 [mA]; [51] IN51 6軸目 指令電流 上位 [mA]; [52] IN52 6軸目 現在速度 [実機単位・符号付き]; [53] IN53 6軸目 予約（使用禁止）; [54] IN54 6軸目 軸異常コード; [55] IN55 6軸目 状態信号（PEND/SV等）; [56] IN56 用途未確認（今回未使用）; [57] IN57 用途未確認（今回未使用）; [58] IN58 用途未確認（今回未使用）; [59] IN59 用途未確認（今回未使用）; [60] IN60 用途未確認（今回未使用）; [61] IN61 用途未確認（今回未使用）; [62] IN62 用途未確認（今回未使用）; [63] IN63 用途未確認（今回未使用）; [64] IN64 用途未確認（今回未使用）; [65] IN65 用途未確認（今回未使用）; [66] IN66 用途未確認（今回未使用）; [67] IN67 用途未確認（今回未使用）; [68] IN68 用途未確認（今回未使用）; [69] IN69 用途未確認（今回未使用）; [70] IN70 用途未確認（今回未使用）; [71] IN71 用途未確認（今回未使用） *)
    RCON1_RxWord : ARRAY[0..71] OF WORD;  (* RCON1 受信ワード（正規化後）; [0] IN00 GW状態; [1] IN01 軸リンク状態; [2] IN02 電源状態0; [3] IN03 電源状態1; [4] IN04 電源状態2; [5] IN05 電源状態3; [6] IN06 電源状態4（構成依存）; [7] IN07 予約（使用禁止）; [8] IN08 1軸目 現在位置 下位 [0.01mm]; [9] IN09 1軸目 現在位置 上位 [0.01mm]; [10] IN10 1軸目 指令電流 下位 [mA]; [11] IN11 1軸目 指令電流 上位 [mA]; [12] IN12 1軸目 現在速度 [実機単位・符号付き]; [13] IN13 1軸目 予約（使用禁止）; [14] IN14 1軸目 軸異常コード; [15] IN15 1軸目 状態信号（PEND/SV等）; [16] IN16 2軸目 現在位置 下位 [0.01mm]; [17] IN17 2軸目 現在位置 上位 [0.01mm]; [18] IN18 2軸目 指令電流 下位 [mA]; [19] IN19 2軸目 指令電流 上位 [mA]; [20] IN20 2軸目 現在速度 [実機単位・符号付き]; [21] IN21 2軸目 予約（使用禁止）; [22] IN22 2軸目 軸異常コード; [23] IN23 2軸目 状態信号（PEND/SV等）; [24] IN24 3軸目 現在位置 下位 [0.01mm]; [25] IN25 3軸目 現在位置 上位 [0.01mm]; [26] IN26 3軸目 指令電流 下位 [mA]; [27] IN27 3軸目 指令電流 上位 [mA]; [28] IN28 3軸目 現在速度 [実機単位・符号付き]; [29] IN29 3軸目 予約（使用禁止）; [30] IN30 3軸目 軸異常コード; [31] IN31 3軸目 状態信号（PEND/SV等）; [32] IN32 4軸目 現在位置 下位 [0.01mm]; [33] IN33 4軸目 現在位置 上位 [0.01mm]; [34] IN34 4軸目 指令電流 下位 [mA]; [35] IN35 4軸目 指令電流 上位 [mA]; [36] IN36 4軸目 現在速度 [実機単位・符号付き]; [37] IN37 4軸目 予約（使用禁止）; [38] IN38 4軸目 軸異常コード; [39] IN39 4軸目 状態信号（PEND/SV等）; [40] IN40 5軸目 現在位置 下位 [0.01mm]; [41] IN41 5軸目 現在位置 上位 [0.01mm]; [42] IN42 5軸目 指令電流 下位 [mA]; [43] IN43 5軸目 指令電流 上位 [mA]; [44] IN44 5軸目 現在速度 [実機単位・符号付き]; [45] IN45 5軸目 予約（使用禁止）; [46] IN46 5軸目 軸異常コード; [47] IN47 5軸目 状態信号（PEND/SV等）; [48] IN48 6軸目 現在位置 下位 [0.01mm]; [49] IN49 6軸目 現在位置 上位 [0.01mm]; [50] IN50 6軸目 指令電流 下位 [mA]; [51] IN51 6軸目 指令電流 上位 [mA]; [52] IN52 6軸目 現在速度 [実機単位・符号付き]; [53] IN53 6軸目 予約（使用禁止）; [54] IN54 6軸目 軸異常コード; [55] IN55 6軸目 状態信号（PEND/SV等）; [56] IN56 用途未確認（今回未使用）; [57] IN57 用途未確認（今回未使用）; [58] IN58 用途未確認（今回未使用）; [59] IN59 用途未確認（今回未使用）; [60] IN60 用途未確認（今回未使用）; [61] IN61 用途未確認（今回未使用）; [62] IN62 用途未確認（今回未使用）; [63] IN63 用途未確認（今回未使用）; [64] IN64 用途未確認（今回未使用）; [65] IN65 用途未確認（今回未使用）; [66] IN66 用途未確認（今回未使用）; [67] IN67 用途未確認（今回未使用）; [68] IN68 用途未確認（今回未使用）; [69] IN69 用途未確認（今回未使用）; [70] IN70 用途未確認（今回未使用）; [71] IN71 用途未確認（今回未使用） *)
    RCON1_TxWord : ARRAY[0..55] OF WORD;  (* RCON1 送信ワード候補; [0] OUT00 共通制御（MON/RTE）; [1] OUT01 予約（書込禁止）; [2] OUT02 予約（書込禁止）; [3] OUT03 予約（書込禁止）; [4] OUT04 予約（書込禁止）; [5] OUT05 予約（書込禁止）; [6] OUT06 予約（書込禁止）; [7] OUT07 予約（書込禁止）; [8] OUT08 1軸目 目標位置 下位 [0.01mm]; [9] OUT09 1軸目 目標位置 上位 [0.01mm]; [10] OUT10 1軸目 位置決め幅 下位 [0.01mm]; [11] OUT11 1軸目 位置決め幅 上位 [0.01mm]; [12] OUT12 1軸目 速度指令 [実機単位]; [13] OUT13 1軸目 共通加減速 [0.01G]; [14] OUT14 1軸目 押付け制限 [255=100%]; [15] OUT15 1軸目 制御信号（DSTR/SON等）; [16] OUT16 2軸目 目標位置 下位 [0.01mm]; [17] OUT17 2軸目 目標位置 上位 [0.01mm]; [18] OUT18 2軸目 位置決め幅 下位 [0.01mm]; [19] OUT19 2軸目 位置決め幅 上位 [0.01mm]; [20] OUT20 2軸目 速度指令 [実機単位]; [21] OUT21 2軸目 共通加減速 [0.01G]; [22] OUT22 2軸目 押付け制限 [255=100%]; [23] OUT23 2軸目 制御信号（DSTR/SON等）; [24] OUT24 3軸目 目標位置 下位 [0.01mm]; [25] OUT25 3軸目 目標位置 上位 [0.01mm]; [26] OUT26 3軸目 位置決め幅 下位 [0.01mm]; [27] OUT27 3軸目 位置決め幅 上位 [0.01mm]; [28] OUT28 3軸目 速度指令 [実機単位]; [29] OUT29 3軸目 共通加減速 [0.01G]; [30] OUT30 3軸目 押付け制限 [255=100%]; [31] OUT31 3軸目 制御信号（DSTR/SON等）; [32] OUT32 4軸目 目標位置 下位 [0.01mm]; [33] OUT33 4軸目 目標位置 上位 [0.01mm]; [34] OUT34 4軸目 位置決め幅 下位 [0.01mm]; [35] OUT35 4軸目 位置決め幅 上位 [0.01mm]; [36] OUT36 4軸目 速度指令 [実機単位]; [37] OUT37 4軸目 共通加減速 [0.01G]; [38] OUT38 4軸目 押付け制限 [255=100%]; [39] OUT39 4軸目 制御信号（DSTR/SON等）; [40] OUT40 5軸目 目標位置 下位 [0.01mm]; [41] OUT41 5軸目 目標位置 上位 [0.01mm]; [42] OUT42 5軸目 位置決め幅 下位 [0.01mm]; [43] OUT43 5軸目 位置決め幅 上位 [0.01mm]; [44] OUT44 5軸目 速度指令 [実機単位]; [45] OUT45 5軸目 共通加減速 [0.01G]; [46] OUT46 5軸目 押付け制限 [255=100%]; [47] OUT47 5軸目 制御信号（DSTR/SON等）; [48] OUT48 6軸目 目標位置 下位 [0.01mm]; [49] OUT49 6軸目 目標位置 上位 [0.01mm]; [50] OUT50 6軸目 位置決め幅 下位 [0.01mm]; [51] OUT51 6軸目 位置決め幅 上位 [0.01mm]; [52] OUT52 6軸目 速度指令 [実機単位]; [53] OUT53 6軸目 共通加減速 [0.01G]; [54] OUT54 6軸目 押付け制限 [255=100%]; [55] OUT55 6軸目 制御信号（DSTR/SON等） *)
    RCON1_TxUInt : ARRAY[0..55] OF UINT;  (* RCON1 送信UINT候補（実I/Oではない）; [0] OUT00 共通制御（MON/RTE）; [1] OUT01 予約（書込禁止）; [2] OUT02 予約（書込禁止）; [3] OUT03 予約（書込禁止）; [4] OUT04 予約（書込禁止）; [5] OUT05 予約（書込禁止）; [6] OUT06 予約（書込禁止）; [7] OUT07 予約（書込禁止）; [8] OUT08 1軸目 目標位置 下位 [0.01mm]; [9] OUT09 1軸目 目標位置 上位 [0.01mm]; [10] OUT10 1軸目 位置決め幅 下位 [0.01mm]; [11] OUT11 1軸目 位置決め幅 上位 [0.01mm]; [12] OUT12 1軸目 速度指令 [実機単位]; [13] OUT13 1軸目 共通加減速 [0.01G]; [14] OUT14 1軸目 押付け制限 [255=100%]; [15] OUT15 1軸目 制御信号（DSTR/SON等）; [16] OUT16 2軸目 目標位置 下位 [0.01mm]; [17] OUT17 2軸目 目標位置 上位 [0.01mm]; [18] OUT18 2軸目 位置決め幅 下位 [0.01mm]; [19] OUT19 2軸目 位置決め幅 上位 [0.01mm]; [20] OUT20 2軸目 速度指令 [実機単位]; [21] OUT21 2軸目 共通加減速 [0.01G]; [22] OUT22 2軸目 押付け制限 [255=100%]; [23] OUT23 2軸目 制御信号（DSTR/SON等）; [24] OUT24 3軸目 目標位置 下位 [0.01mm]; [25] OUT25 3軸目 目標位置 上位 [0.01mm]; [26] OUT26 3軸目 位置決め幅 下位 [0.01mm]; [27] OUT27 3軸目 位置決め幅 上位 [0.01mm]; [28] OUT28 3軸目 速度指令 [実機単位]; [29] OUT29 3軸目 共通加減速 [0.01G]; [30] OUT30 3軸目 押付け制限 [255=100%]; [31] OUT31 3軸目 制御信号（DSTR/SON等）; [32] OUT32 4軸目 目標位置 下位 [0.01mm]; [33] OUT33 4軸目 目標位置 上位 [0.01mm]; [34] OUT34 4軸目 位置決め幅 下位 [0.01mm]; [35] OUT35 4軸目 位置決め幅 上位 [0.01mm]; [36] OUT36 4軸目 速度指令 [実機単位]; [37] OUT37 4軸目 共通加減速 [0.01G]; [38] OUT38 4軸目 押付け制限 [255=100%]; [39] OUT39 4軸目 制御信号（DSTR/SON等）; [40] OUT40 5軸目 目標位置 下位 [0.01mm]; [41] OUT41 5軸目 目標位置 上位 [0.01mm]; [42] OUT42 5軸目 位置決め幅 下位 [0.01mm]; [43] OUT43 5軸目 位置決め幅 上位 [0.01mm]; [44] OUT44 5軸目 速度指令 [実機単位]; [45] OUT45 5軸目 共通加減速 [0.01G]; [46] OUT46 5軸目 押付け制限 [255=100%]; [47] OUT47 5軸目 制御信号（DSTR/SON等）; [48] OUT48 6軸目 目標位置 下位 [0.01mm]; [49] OUT49 6軸目 目標位置 上位 [0.01mm]; [50] OUT50 6軸目 位置決め幅 下位 [0.01mm]; [51] OUT51 6軸目 位置決め幅 上位 [0.01mm]; [52] OUT52 6軸目 速度指令 [実機単位]; [53] OUT53 6軸目 共通加減速 [0.01G]; [54] OUT54 6軸目 押付け制限 [255=100%]; [55] OUT55 6軸目 制御信号（DSTR/SON等） *)
    RCON1_LayoutConfirmed : BOOL;  (* RCON1 I/O配置確認済み（初期OFF） *)
    RCON1_ByteOrderConfirmed : BOOL;  (* RCON1 ワード・バイト順確認済み（初期OFF） *)
    RCON1_SwapBytes : BOOL;  (* RCON1 上下バイト交換設定（ON=交換） *)
    RCON1_CommOK : BOOL;  (* RCON1 通信正常（外部判定・固定ON不可） *)
    RCON1_GwMON_Request : BOOL;  (* RCON1 MON要求（b15） *)
    RCON1_GwRTE_Request : BOOL;  (* RCON1 通信異常ラッチ解除要求（b13） *)
    RCON1_GwRun : BOOL;  (* RCON1 GW動作中（RUN/b15） *)
    RCON1_GwControllerCommLatch : BOOL;  (* RCON1 GW通信異常保持（LERC/b14） *)
    RCON1_GwAxisCommError : BOOL;  (* RCON1 GW－軸 通信異常（ERRT/b13） *)
    RCON1_GwManual : BOOL;  (* RCON1 手動モード（MOD/b12） *)
    RCON1_GwHeavyAlarm : BOOL;  (* RCON1 GW重故障（ALMH/b11） *)
    RCON1_GwLightAlarm : BOOL;  (* RCON1 GW軽故障（ALML/b10） *)
    RCON1_GwSystemStop : BOOL;  (* RCON1 システム停止状態（SEMG/b8・監視用） *)
    RCON1_GwAlarmCode : UINT;  (* RCON1 GW異常コード（ALMC/b0～7） *)
    RCON1_AxisLinked : ARRAY[1..6] OF BOOL;  (* RCON1 軸別リンク状態; [1] 1軸目（No.0）リンク状態; [2] 2軸目（No.1）リンク状態; [3] 3軸目（No.2）リンク状態; [4] 4軸目（No.3）リンク状態; [5] 5軸目（No.4）リンク状態; [6] 6軸目（No.5）リンク状態 *)
    RCON1_PowerStateRaw : ARRAY[0..4] OF WORD;  (* RCON1 電源状態ワード（詳細未確認）; [0] IN02 電源状態0（詳細未確認）; [1] IN03 電源状態1（詳細未確認）; [2] IN04 電源状態2（詳細未確認）; [3] IN05 電源状態3（詳細未確認）; [4] IN06 電源状態4（詳細未確認） *)
    RCON1_EncodeOK : ARRAY[1..6] OF BOOL;  (* RCON1 軸別変換正常（運転許可とは別）; [1] 1軸目（No.0）変換正常; [2] 2軸目（No.1）変換正常; [3] 3軸目（No.2）変換正常; [4] 4軸目（No.3）変換正常; [5] 5軸目（No.4）変換正常; [6] 6軸目（No.5）変換正常 *)
    RCON1_EncodeError : ARRAY[1..6] OF UINT;  (* RCON1 軸別変換エラー番号（0=正常）; [1] 1軸目（No.0）変換エラー番号; [2] 2軸目（No.1）変換エラー番号; [3] 3軸目（No.2）変換エラー番号; [4] 4軸目（No.3）変換エラー番号; [5] 5軸目（No.4）変換エラー番号; [6] 6軸目（No.5）変換エラー番号 *)
    RCON1_WriteEnable : BOOL;  (* RCON1 実出力書込み許可（OFF=前値保持・停止不可） *)
    RCON1_GwApply : BOOL;  (* RCON1 共通出力更新許可（OFF=前値保持） *)
    RCON1_AxisApply : ARRAY[1..6] OF BOOL;  (* RCON1 軸別出力更新許可（OFF=前値保持）; [1] 1軸目（No.0）出力更新許可（OFF=前値保持）; [2] 2軸目（No.1）出力更新許可（OFF=前値保持）; [3] 3軸目（No.2）出力更新許可（OFF=前値保持）; [4] 4軸目（No.3）出力更新許可（OFF=前値保持）; [5] 5軸目（No.4）出力更新許可（OFF=前値保持）; [6] 6軸目（No.5）出力更新許可（OFF=前値保持） *)
    RCON1_MotionPermit : ARRAY[1..6] OF BOOL;  (* RCON1 軸別運転許可（外部判定・初期OFF）; [1] 1軸目（No.0）運転許可（外部判定）; [2] 2軸目（No.1）運転許可（外部判定）; [3] 3軸目（No.2）運転許可（外部判定）; [4] 4軸目（No.3）運転許可（外部判定）; [5] 5軸目（No.4）運転許可（外部判定）; [6] 6軸目（No.5）運転許可（外部判定） *)
    RCON1_GwWritten : BOOL;  (* RCON1 共通出力代入済み（RCON受付とは別） *)
    RCON1_AxisWritten : ARRAY[1..6] OF BOOL;  (* RCON1 軸別出力代入済み（RCON受付とは別）; [1] 1軸目（No.0）出力代入済み（RCON受付とは別）; [2] 2軸目（No.1）出力代入済み（RCON受付とは別）; [3] 3軸目（No.2）出力代入済み（RCON受付とは別）; [4] 4軸目（No.3）出力代入済み（RCON受付とは別）; [5] 5軸目（No.4）出力代入済み（RCON受付とは別）; [6] 6軸目（No.5）出力代入済み（RCON受付とは別） *)
    RCON2_RxRaw : ARRAY[0..55] OF UINT;  (* RCON2 受信値（バイト交換前）; [0] IN00 GW状態; [1] IN01 軸リンク状態; [2] IN02 電源状態0; [3] IN03 電源状態1; [4] IN04 電源状態2; [5] IN05 電源状態3; [6] IN06 電源状態4（構成依存）; [7] IN07 予約（使用禁止）; [8] IN08 1軸目 現在位置 下位 [0.01mm]; [9] IN09 1軸目 現在位置 上位 [0.01mm]; [10] IN10 1軸目 指令電流 下位 [mA]; [11] IN11 1軸目 指令電流 上位 [mA]; [12] IN12 1軸目 現在速度 [実機単位・符号付き]; [13] IN13 1軸目 予約（使用禁止）; [14] IN14 1軸目 軸異常コード; [15] IN15 1軸目 状態信号（PEND/SV等）; [16] IN16 2軸目 現在位置 下位 [0.01mm]; [17] IN17 2軸目 現在位置 上位 [0.01mm]; [18] IN18 2軸目 指令電流 下位 [mA]; [19] IN19 2軸目 指令電流 上位 [mA]; [20] IN20 2軸目 現在速度 [実機単位・符号付き]; [21] IN21 2軸目 予約（使用禁止）; [22] IN22 2軸目 軸異常コード; [23] IN23 2軸目 状態信号（PEND/SV等）; [24] IN24 3軸目 現在位置 下位 [0.01mm]; [25] IN25 3軸目 現在位置 上位 [0.01mm]; [26] IN26 3軸目 指令電流 下位 [mA]; [27] IN27 3軸目 指令電流 上位 [mA]; [28] IN28 3軸目 現在速度 [実機単位・符号付き]; [29] IN29 3軸目 予約（使用禁止）; [30] IN30 3軸目 軸異常コード; [31] IN31 3軸目 状態信号（PEND/SV等）; [32] IN32 4軸目 現在位置 下位 [0.01mm]; [33] IN33 4軸目 現在位置 上位 [0.01mm]; [34] IN34 4軸目 指令電流 下位 [mA]; [35] IN35 4軸目 指令電流 上位 [mA]; [36] IN36 4軸目 現在速度 [実機単位・符号付き]; [37] IN37 4軸目 予約（使用禁止）; [38] IN38 4軸目 軸異常コード; [39] IN39 4軸目 状態信号（PEND/SV等）; [40] IN40 5軸目 現在位置 下位 [0.01mm]; [41] IN41 5軸目 現在位置 上位 [0.01mm]; [42] IN42 5軸目 指令電流 下位 [mA]; [43] IN43 5軸目 指令電流 上位 [mA]; [44] IN44 5軸目 現在速度 [実機単位・符号付き]; [45] IN45 5軸目 予約（使用禁止）; [46] IN46 5軸目 軸異常コード; [47] IN47 5軸目 状態信号（PEND/SV等）; [48] IN48 用途未確認（今回未使用）; [49] IN49 用途未確認（今回未使用）; [50] IN50 用途未確認（今回未使用）; [51] IN51 用途未確認（今回未使用）; [52] IN52 用途未確認（今回未使用）; [53] IN53 用途未確認（今回未使用）; [54] IN54 用途未確認（今回未使用）; [55] IN55 用途未確認（今回未使用） *)
    RCON2_RxWord : ARRAY[0..55] OF WORD;  (* RCON2 受信ワード（正規化後）; [0] IN00 GW状態; [1] IN01 軸リンク状態; [2] IN02 電源状態0; [3] IN03 電源状態1; [4] IN04 電源状態2; [5] IN05 電源状態3; [6] IN06 電源状態4（構成依存）; [7] IN07 予約（使用禁止）; [8] IN08 1軸目 現在位置 下位 [0.01mm]; [9] IN09 1軸目 現在位置 上位 [0.01mm]; [10] IN10 1軸目 指令電流 下位 [mA]; [11] IN11 1軸目 指令電流 上位 [mA]; [12] IN12 1軸目 現在速度 [実機単位・符号付き]; [13] IN13 1軸目 予約（使用禁止）; [14] IN14 1軸目 軸異常コード; [15] IN15 1軸目 状態信号（PEND/SV等）; [16] IN16 2軸目 現在位置 下位 [0.01mm]; [17] IN17 2軸目 現在位置 上位 [0.01mm]; [18] IN18 2軸目 指令電流 下位 [mA]; [19] IN19 2軸目 指令電流 上位 [mA]; [20] IN20 2軸目 現在速度 [実機単位・符号付き]; [21] IN21 2軸目 予約（使用禁止）; [22] IN22 2軸目 軸異常コード; [23] IN23 2軸目 状態信号（PEND/SV等）; [24] IN24 3軸目 現在位置 下位 [0.01mm]; [25] IN25 3軸目 現在位置 上位 [0.01mm]; [26] IN26 3軸目 指令電流 下位 [mA]; [27] IN27 3軸目 指令電流 上位 [mA]; [28] IN28 3軸目 現在速度 [実機単位・符号付き]; [29] IN29 3軸目 予約（使用禁止）; [30] IN30 3軸目 軸異常コード; [31] IN31 3軸目 状態信号（PEND/SV等）; [32] IN32 4軸目 現在位置 下位 [0.01mm]; [33] IN33 4軸目 現在位置 上位 [0.01mm]; [34] IN34 4軸目 指令電流 下位 [mA]; [35] IN35 4軸目 指令電流 上位 [mA]; [36] IN36 4軸目 現在速度 [実機単位・符号付き]; [37] IN37 4軸目 予約（使用禁止）; [38] IN38 4軸目 軸異常コード; [39] IN39 4軸目 状態信号（PEND/SV等）; [40] IN40 5軸目 現在位置 下位 [0.01mm]; [41] IN41 5軸目 現在位置 上位 [0.01mm]; [42] IN42 5軸目 指令電流 下位 [mA]; [43] IN43 5軸目 指令電流 上位 [mA]; [44] IN44 5軸目 現在速度 [実機単位・符号付き]; [45] IN45 5軸目 予約（使用禁止）; [46] IN46 5軸目 軸異常コード; [47] IN47 5軸目 状態信号（PEND/SV等）; [48] IN48 用途未確認（今回未使用）; [49] IN49 用途未確認（今回未使用）; [50] IN50 用途未確認（今回未使用）; [51] IN51 用途未確認（今回未使用）; [52] IN52 用途未確認（今回未使用）; [53] IN53 用途未確認（今回未使用）; [54] IN54 用途未確認（今回未使用）; [55] IN55 用途未確認（今回未使用） *)
    RCON2_TxWord : ARRAY[0..47] OF WORD;  (* RCON2 送信ワード候補; [0] OUT00 共通制御（MON/RTE）; [1] OUT01 予約（書込禁止）; [2] OUT02 予約（書込禁止）; [3] OUT03 予約（書込禁止）; [4] OUT04 予約（書込禁止）; [5] OUT05 予約（書込禁止）; [6] OUT06 予約（書込禁止）; [7] OUT07 予約（書込禁止）; [8] OUT08 1軸目 目標位置 下位 [0.01mm]; [9] OUT09 1軸目 目標位置 上位 [0.01mm]; [10] OUT10 1軸目 位置決め幅 下位 [0.01mm]; [11] OUT11 1軸目 位置決め幅 上位 [0.01mm]; [12] OUT12 1軸目 速度指令 [実機単位]; [13] OUT13 1軸目 共通加減速 [0.01G]; [14] OUT14 1軸目 押付け制限 [255=100%]; [15] OUT15 1軸目 制御信号（DSTR/SON等）; [16] OUT16 2軸目 目標位置 下位 [0.01mm]; [17] OUT17 2軸目 目標位置 上位 [0.01mm]; [18] OUT18 2軸目 位置決め幅 下位 [0.01mm]; [19] OUT19 2軸目 位置決め幅 上位 [0.01mm]; [20] OUT20 2軸目 速度指令 [実機単位]; [21] OUT21 2軸目 共通加減速 [0.01G]; [22] OUT22 2軸目 押付け制限 [255=100%]; [23] OUT23 2軸目 制御信号（DSTR/SON等）; [24] OUT24 3軸目 目標位置 下位 [0.01mm]; [25] OUT25 3軸目 目標位置 上位 [0.01mm]; [26] OUT26 3軸目 位置決め幅 下位 [0.01mm]; [27] OUT27 3軸目 位置決め幅 上位 [0.01mm]; [28] OUT28 3軸目 速度指令 [実機単位]; [29] OUT29 3軸目 共通加減速 [0.01G]; [30] OUT30 3軸目 押付け制限 [255=100%]; [31] OUT31 3軸目 制御信号（DSTR/SON等）; [32] OUT32 4軸目 目標位置 下位 [0.01mm]; [33] OUT33 4軸目 目標位置 上位 [0.01mm]; [34] OUT34 4軸目 位置決め幅 下位 [0.01mm]; [35] OUT35 4軸目 位置決め幅 上位 [0.01mm]; [36] OUT36 4軸目 速度指令 [実機単位]; [37] OUT37 4軸目 共通加減速 [0.01G]; [38] OUT38 4軸目 押付け制限 [255=100%]; [39] OUT39 4軸目 制御信号（DSTR/SON等）; [40] OUT40 5軸目 目標位置 下位 [0.01mm]; [41] OUT41 5軸目 目標位置 上位 [0.01mm]; [42] OUT42 5軸目 位置決め幅 下位 [0.01mm]; [43] OUT43 5軸目 位置決め幅 上位 [0.01mm]; [44] OUT44 5軸目 速度指令 [実機単位]; [45] OUT45 5軸目 共通加減速 [0.01G]; [46] OUT46 5軸目 押付け制限 [255=100%]; [47] OUT47 5軸目 制御信号（DSTR/SON等） *)
    RCON2_TxUInt : ARRAY[0..47] OF UINT;  (* RCON2 送信UINT候補（実I/Oではない）; [0] OUT00 共通制御（MON/RTE）; [1] OUT01 予約（書込禁止）; [2] OUT02 予約（書込禁止）; [3] OUT03 予約（書込禁止）; [4] OUT04 予約（書込禁止）; [5] OUT05 予約（書込禁止）; [6] OUT06 予約（書込禁止）; [7] OUT07 予約（書込禁止）; [8] OUT08 1軸目 目標位置 下位 [0.01mm]; [9] OUT09 1軸目 目標位置 上位 [0.01mm]; [10] OUT10 1軸目 位置決め幅 下位 [0.01mm]; [11] OUT11 1軸目 位置決め幅 上位 [0.01mm]; [12] OUT12 1軸目 速度指令 [実機単位]; [13] OUT13 1軸目 共通加減速 [0.01G]; [14] OUT14 1軸目 押付け制限 [255=100%]; [15] OUT15 1軸目 制御信号（DSTR/SON等）; [16] OUT16 2軸目 目標位置 下位 [0.01mm]; [17] OUT17 2軸目 目標位置 上位 [0.01mm]; [18] OUT18 2軸目 位置決め幅 下位 [0.01mm]; [19] OUT19 2軸目 位置決め幅 上位 [0.01mm]; [20] OUT20 2軸目 速度指令 [実機単位]; [21] OUT21 2軸目 共通加減速 [0.01G]; [22] OUT22 2軸目 押付け制限 [255=100%]; [23] OUT23 2軸目 制御信号（DSTR/SON等）; [24] OUT24 3軸目 目標位置 下位 [0.01mm]; [25] OUT25 3軸目 目標位置 上位 [0.01mm]; [26] OUT26 3軸目 位置決め幅 下位 [0.01mm]; [27] OUT27 3軸目 位置決め幅 上位 [0.01mm]; [28] OUT28 3軸目 速度指令 [実機単位]; [29] OUT29 3軸目 共通加減速 [0.01G]; [30] OUT30 3軸目 押付け制限 [255=100%]; [31] OUT31 3軸目 制御信号（DSTR/SON等）; [32] OUT32 4軸目 目標位置 下位 [0.01mm]; [33] OUT33 4軸目 目標位置 上位 [0.01mm]; [34] OUT34 4軸目 位置決め幅 下位 [0.01mm]; [35] OUT35 4軸目 位置決め幅 上位 [0.01mm]; [36] OUT36 4軸目 速度指令 [実機単位]; [37] OUT37 4軸目 共通加減速 [0.01G]; [38] OUT38 4軸目 押付け制限 [255=100%]; [39] OUT39 4軸目 制御信号（DSTR/SON等）; [40] OUT40 5軸目 目標位置 下位 [0.01mm]; [41] OUT41 5軸目 目標位置 上位 [0.01mm]; [42] OUT42 5軸目 位置決め幅 下位 [0.01mm]; [43] OUT43 5軸目 位置決め幅 上位 [0.01mm]; [44] OUT44 5軸目 速度指令 [実機単位]; [45] OUT45 5軸目 共通加減速 [0.01G]; [46] OUT46 5軸目 押付け制限 [255=100%]; [47] OUT47 5軸目 制御信号（DSTR/SON等） *)
    RCON2_LayoutConfirmed : BOOL;  (* RCON2 I/O配置確認済み（初期OFF） *)
    RCON2_ByteOrderConfirmed : BOOL;  (* RCON2 ワード・バイト順確認済み（初期OFF） *)
    RCON2_SwapBytes : BOOL;  (* RCON2 上下バイト交換設定（ON=交換） *)
    RCON2_CommOK : BOOL;  (* RCON2 通信正常（外部判定・固定ON不可） *)
    RCON2_GwMON_Request : BOOL;  (* RCON2 MON要求（b15） *)
    RCON2_GwRTE_Request : BOOL;  (* RCON2 通信異常ラッチ解除要求（b13） *)
    RCON2_GwRun : BOOL;  (* RCON2 GW動作中（RUN/b15） *)
    RCON2_GwControllerCommLatch : BOOL;  (* RCON2 GW通信異常保持（LERC/b14） *)
    RCON2_GwAxisCommError : BOOL;  (* RCON2 GW－軸 通信異常（ERRT/b13） *)
    RCON2_GwManual : BOOL;  (* RCON2 手動モード（MOD/b12） *)
    RCON2_GwHeavyAlarm : BOOL;  (* RCON2 GW重故障（ALMH/b11） *)
    RCON2_GwLightAlarm : BOOL;  (* RCON2 GW軽故障（ALML/b10） *)
    RCON2_GwSystemStop : BOOL;  (* RCON2 システム停止状態（SEMG/b8・監視用） *)
    RCON2_GwAlarmCode : UINT;  (* RCON2 GW異常コード（ALMC/b0～7） *)
    RCON2_AxisLinked : ARRAY[1..5] OF BOOL;  (* RCON2 軸別リンク状態; [1] 1軸目（No.0）リンク状態; [2] 2軸目（No.1）リンク状態; [3] 3軸目（No.2）リンク状態; [4] 4軸目（No.3）リンク状態; [5] 5軸目（No.4）リンク状態 *)
    RCON2_PowerStateRaw : ARRAY[0..4] OF WORD;  (* RCON2 電源状態ワード（詳細未確認）; [0] IN02 電源状態0（詳細未確認）; [1] IN03 電源状態1（詳細未確認）; [2] IN04 電源状態2（詳細未確認）; [3] IN05 電源状態3（詳細未確認）; [4] IN06 電源状態4（詳細未確認） *)
    RCON2_EncodeOK : ARRAY[1..5] OF BOOL;  (* RCON2 軸別変換正常（運転許可とは別）; [1] 1軸目（No.0）変換正常; [2] 2軸目（No.1）変換正常; [3] 3軸目（No.2）変換正常; [4] 4軸目（No.3）変換正常; [5] 5軸目（No.4）変換正常 *)
    RCON2_EncodeError : ARRAY[1..5] OF UINT;  (* RCON2 軸別変換エラー番号（0=正常）; [1] 1軸目（No.0）変換エラー番号; [2] 2軸目（No.1）変換エラー番号; [3] 3軸目（No.2）変換エラー番号; [4] 4軸目（No.3）変換エラー番号; [5] 5軸目（No.4）変換エラー番号 *)
    RCON2_WriteEnable : BOOL;  (* RCON2 実出力書込み許可（OFF=前値保持・停止不可） *)
    RCON2_GwApply : BOOL;  (* RCON2 共通出力更新許可（OFF=前値保持） *)
    RCON2_AxisApply : ARRAY[1..5] OF BOOL;  (* RCON2 軸別出力更新許可（OFF=前値保持）; [1] 1軸目（No.0）出力更新許可（OFF=前値保持）; [2] 2軸目（No.1）出力更新許可（OFF=前値保持）; [3] 3軸目（No.2）出力更新許可（OFF=前値保持）; [4] 4軸目（No.3）出力更新許可（OFF=前値保持）; [5] 5軸目（No.4）出力更新許可（OFF=前値保持） *)
    RCON2_MotionPermit : ARRAY[1..5] OF BOOL;  (* RCON2 軸別運転許可（外部判定・初期OFF）; [1] 1軸目（No.0）運転許可（外部判定）; [2] 2軸目（No.1）運転許可（外部判定）; [3] 3軸目（No.2）運転許可（外部判定）; [4] 4軸目（No.3）運転許可（外部判定）; [5] 5軸目（No.4）運転許可（外部判定） *)
    RCON2_GwWritten : BOOL;  (* RCON2 共通出力代入済み（RCON受付とは別） *)
    RCON2_AxisWritten : ARRAY[1..5] OF BOOL;  (* RCON2 軸別出力代入済み（RCON受付とは別）; [1] 1軸目（No.0）出力代入済み（RCON受付とは別）; [2] 2軸目（No.1）出力代入済み（RCON受付とは別）; [3] 3軸目（No.2）出力代入済み（RCON受付とは別）; [4] 4軸目（No.3）出力代入済み（RCON受付とは別）; [5] 5軸目（No.4）出力代入済み（RCON受付とは別） *)
    RCON1_IAI_Auto : ARRAY[0..99] OF Bool;  (* A(左側) RCON1/Node1/ NG排出：; [1] 原点位置移動; [2] NG仕分け; [3] 動作完了後 原点位置移動 *)
    RCON1_OUT_PositionBand_mm : LREAL;  (* RCON1位置決め幅 [mm] *)
    RCON1_OUT_TargetPos_mm : LREAL;  (* RCON1目標位置 [mm] *)
    RCON1_OUT_Speed_mm_s : LREAL;  (* 指令速度 [mm/s] *)
    RCON1_OUT_AccDec_G : LREAL;  (* 共通加減速度 [G] *)
    RCON1_OUT_PushLimit_pct : LREAL;  (* 押付け電流制限 [%] *)
    RCON1_ActualPos_mm : LREAL;  (* 現在位置 [mm] *)
    RCON1_Current_mA : DINT;  (* 指令電流 [mA] *)
    RCON1_ActualSpeed_mm_s : LREAL;  (* 現在速度 [mm/s・符号付き] *)
    RCON1_AlarmCode : UINT;  (* 軸異常コード *)
    RCON1_DataValid : BOOL;  (* 入力有効（運転許可とは別） *)
    RCON1_1_IN_PositionDone : BOOL;  (* 位置決め完了 *)
    RCON1_1_IN_HomeDone : BOOL;  (* 原点復帰完了 *)
    RCON1_1_IN_Moving : BOOL;  (* 移動中 *)
    RCON1_1_IN_EmergencyStop : BOOL;  (* 非常停止状態 *)
    RCON1_1_IN_ControllerReady : BOOL;  (* コントローラー準備完了 *)
    RCON1_1_IN_Zone2 : BOOL;  (* ゾーン2内 *)
    RCON1_1_IN_Zone1 : BOOL;  (* ゾーン1内 *)
    RCON1_1_IN_CommandDone : BOOL;  (* 指令完了 *)
    RCON1_1_IN_OverloadWarning : BOOL;  (* 過負荷警告等 *)
    RCON1_1_IN_PushMiss : BOOL;  (* 押付け空振り *)
    RCON1_1_IN_ServoReady : BOOL;  (* サーボON状態 *)
    RCON1_1_IN_Alarm : BOOL;  (* RCON1 軸異常 *)
    RCON1_1_Ready : BOOL;  (* 運転可能状態 *)
    RCON1_1_Error : BOOL;  (* RCON エラー *)
    RCON1_1_Error_Clear : BOOL;
    Error_M : ARRAY[0..99] OF Bool;  (* エラー：; [1] シリンダ; [2] コンベア＆ドアセンサ; [3] FH; [4] A(左側)検査コンベア ワーク不一致; [5] RCON1-1 異常; [6] GT2 エラー; [7] NG1仕分けエラー *)
    HMI_RCON1_OUT_TargetPos : ARRAY[0..99] OF LREAL;  (* HMI RC01 NG仕分け位置：; [1] 原点位置; [3] 高さNG位置; [4] カメラ キズNG位置; [5] カメラ 姿NG位置 *)
    RCON1_1_M : ARRAY[0..99] OF BOOL;  (* [1] 開始指令; [2] 動作完了 *)
    ST1_A_Ca1_M : ARRAY[0..99] OF Bool;  (* [6] ST2 検査前ワーク不一致エラー; [3] ワーク有無 判定; [1] ST1 A カメラ1 検査開始; [4] ST1 A ワーク有; [5] ST1 A ワーク無; [2] 【Y720】A(左側) 位置1ストッパー 戻; [7] ST1 FH測定開始 *)
    ST2_A_Hgt_M : ARRAY[0..99] OF Bool;  (* [4] 【Y721】A(左側) 位置2ストッパー戻; [6] ST2 A ワーク有; [7] ST2 A ワーク無 / 前工程NG; [5] ワーク有無 判定; [9] 【Y703】A(左側) 高さ検査持上行; [10] 【Y701】A(左側) 高さ検査押え行; [11] A(左側) 高さ検査OK判定; [12] A(左側) 高さ検査NG判定; [2] 【Y701】A(左側) 高さ検査押え行; [8] ST2 検査前ワーク不一致エラー *)
    ST3_A_Dis1_End : BOOL;  (* ST3 A 動作完了 *)
    ST3_A_Dis1_M : ARRAY[0..99] OF Bool;  (* [7] 原点位置 移動開始; [6] 原点位置移動 データ転送; [5] 【Y722】A(左側) 位置3ストッパー戻; [4] 【Y706】A(左側) NG1チャック戻; [8] ワーク有無 / 検査前ワーク不一致 判定; [9] S3 A ワーク有 工程NG; [10] S3 A ワーク無  前工程OK; [14] 【Y704】A(左側) NG1ピックアップ戻 ; [24] 仕分け完了; [16] 高さNG位置; [17] カメラ キズNG位置; [18] カメラ 姿NG位置; [21] 高さNG; [22] カメラ キズNG; [23] カメラ 姿NG; [11] ST3 検査前ワーク不一致エラー; [25] #動作完了後 原点位置移動 *)
    Homing_Para_Stm : _sHOMING_REF;
    Stm_A_Rev_Axis000_OriginDone : BOOL;  (* A(左側) ST4 反転1 モータ原点復帰完了 *)
    HMI_Home_SW : BOOL;  (* HMI 原点復帰SW *)
    Origin_Busy : BOOL;  (* 原点復帰中 *)
    Out_CYw_Rev_01_Pick_A_H_Origin : ARRAY[0..10] OF Bool;  (* 原点復帰【Y710】A(左側)ST4 反転1ピックアップ戻： *)
    Stm_A_Rev_Axis000_Origin : BOOL;  (* A(左側) ST4 反転1 モータ原点復帰開始 *)
    Out_CYw_Rev_01_Pick_A_F_Origin : ARRAY[0..99] OF Bool;  (* 原点復帰【Y711】A(左側)ST4 反転1ピックアップ行： *)
    Out_CYw_Rev_01_Chk_A_H_Origin : ARRAY[0..99] OF Bool;  (* 原点復帰【Y708】A(左側)ST4 反転1チャック閉： *)
    Stm_A_Rev_Axis001_Origin : BOOL;  (* A(左側) ST6 反転2 モータ原点復帰開始 *)
    Stm_A_Rev_Axis001_OriginDone : BOOL;  (* A(左側) ST6 反転2 モータ原点復帰完了 *)
    Out_CYw_Rev_02_Pick_A_H_Origin : ARRAY[0..10] OF Bool;  (* 原点復帰 【Y714】A(左側)ST6 反転2ピックアップ戻 *)
    Out_CYw_Rev_02_Pick_A_F_Origin : ARRAY[0..99] OF Bool;  (* 原点復帰 【Y715】A(左側)ST6 反転2ピックアップ行 *)
    Out_CYw_Rev_02_Chk_A_H_Origin : ARRAY[0..99] OF Bool;  (* 原点復帰 【Y712】A(左側)ST6 反転2チャック閉 戻 *)
    Auto_B_Start : BOOL;  (* B(右側)自動運転開始（後続処理未接続） *)
    Stm_B_Rev_Axis002_Origin : BOOL;  (* B(右側) ST4 反転1 モータ原点復帰開始 *)
    Stm_B_Rev_Axis002_OriginDone : BOOL;  (* B(右側) ST4 反転1 モータ原点復帰完了 *)
    Out_CYw_Rev_01_Pick_B_H_Origin : ARRAY[0..10] OF Bool;  (* 原点復帰 【Y810】B(右側)ST4 反転1ピックアップ戻 *)
    Out_CYw_Rev_01_Pick_B_F_Origin : ARRAY[0..99] OF Bool;  (* 原点復帰 【Y811】B(右側)ST4 反転1ピックアップ行 *)
    Out_CYw_Rev_01_Chk_B_H_Origin : ARRAY[0..99] OF Bool;  (* 原点復帰 【Y808】B(右側)ST4 反転1チャック閉 戻 *)
    Stm_B_Rev_Axis003_Origin : BOOL;  (* B(右側) ST6 反転2 モータ原点復帰開始 *)
    Stm_B_Rev_Axis003_OriginDone : BOOL;  (* B(右側) ST6 反転2 モータ原点復帰完了 *)
    Out_CYw_Rev_02_Pick_B_H_Origin : ARRAY[0..10] OF Bool;  (* 原点復帰 【Y814】B(右側)ST6 反転2ピックアップ戻 *)
    Out_CYw_Rev_02_Pick_B_F_Origin : ARRAY[0..99] OF Bool;  (* 原点復帰 【Y815】B(右側)ST6 反転2ピックアップ行 *)
    Out_CYw_Rev_02_Chk_B_H_Origin : ARRAY[0..99] OF Bool;  (* 原点復帰 【Y812】B(右側)ST6 反転2チャック閉 戻 *)
END_VAR

PROGRAM ModeManagement_モード管理
VAR
    Setting_M : BOOL;
    Manual_M : BOOL;
    Auto_M : BOOL;
    Dummy_M : BOOL;
    Inital_M : BOOL;
    Output_Error_M : ARRAY[0..99] OF Bool;
    Index_Error_001 : DINT;
    Index_B_001 : DINT;
    Index_Share_001 : DINT;
    Error_TON : ARRAY[0..99] OF TON;
    Error_TOF : ARRAY[0..99] OF TOF;
    AutoMode_A_M : ARRAY[0..99] OF Bool;
    ６ : DINT;
    ST4_A_Rev_01_Origin_M : ARRAY[0..99] OF Bool;  (* A(左側) ST4 反転1 原点復帰工程; [1] A(左側) ST4 反転1 原点復帰開始; [2] A(左側) ST4 反転1 原点復帰中; [3] A(左側) ST4 反転1 ピックアップ戻; [4] A(左側) ST4 反転1 モータ原点復帰開始; [5] A(左側) ST4 反転1 ピックアップ行; [6] A(左側) ST4 反転1 チャック閉; [7] A(左側) ST4 反転1 原点復帰完了（ワーク無） *)
    ST4_A_Rev_01_OriginDone : BOOL;  (* A(左側) ST4 反転1 原点復帰完了 *)
    ST4_A_Rev_02_Origin_M : ARRAY[0..99] OF Bool;  (* A(左側) ST6 反転2 原点復帰工程; [1] A(左側) ST6 反転2 原点復帰開始; [2] A(左側) ST6 反転2 原点復帰中; [3] A(左側) ST6 反転2 ピックアップ戻; [4] A(左側) ST6 反転2 モータ原点復帰開始; [5] A(左側) ST6 反転2 ピックアップ行; [6] A(左側) ST6 反転2 チャック閉; [7] A(左側) ST6 反転2 原点復帰完了（ワーク無） *)
    ST4_A_Rev_02_OriginDone : BOOL;  (* A(左側) ST6 反転2 原点復帰完了 *)
    ST4_B_Rev_01_Origin_M : ARRAY[0..99] OF Bool;  (* B(右側) ST4 反転1 原点復帰工程; [1] B(右側) ST4 反転1 原点復帰開始; [2] B(右側) ST4 反転1 原点復帰中; [3] B(右側) ST4 反転1 ピックアップ戻; [4] B(右側) ST4 反転1 モータ原点復帰開始; [5] B(右側) ST4 反転1 ピックアップ行; [6] B(右側) ST4 反転1 チャック閉; [7] B(右側) ST4 反転1 原点復帰完了（ワーク無） *)
    ST4_B_Rev_01_OriginDone : BOOL;  (* B(右側) ST4 反転1 原点復帰完了 *)
    ST4_B_Rev_02_Origin_M : ARRAY[0..99] OF Bool;  (* B(右側) ST6 反転2 原点復帰工程; [1] B(右側) ST6 反転2 原点復帰開始; [2] B(右側) ST6 反転2 原点復帰中; [3] B(右側) ST6 反転2 ピックアップ戻; [4] B(右側) ST6 反転2 モータ原点復帰開始; [5] B(右側) ST6 反転2 ピックアップ行; [6] B(右側) ST6 反転2 チャック閉; [7] B(右側) ST6 反転2 原点復帰完了（ワーク無） *)
    ST4_B_Rev_02_OriginDone : BOOL;  (* B(右側) ST6 反転2 原点復帰完了 *)
END_VAR
VAR_EXTERNAL
    Output_A_Error_M : ARRAY[0..99] OF Bool;
    Output_A_Restart_M : ARRAY[0..99] OF Bool;
    In_Sw_RESET : BOOL;
    In_Sw_START : BOOL;
    ManualMode : BOOL;
    M9999 : BOOL;
    Output_B_Error_M : ARRAY[0..99] OF Bool;  (* B(右側)シリンダエラー *)
    Output_B_Restart_M : ARRAY[0..99] OF Bool;  (* B(右側)シリンダ再開： *)
    Output_Share_Error_M : ARRAY[0..99] OF Bool;
    Output_Share_Restart_M : ARRAY[0..99] OF Bool;
    TimerQ_In_Sen_Accum_CV_A_Full : BOOL;
    Out_TDC_Stop : BOOL;
    In_Sen_Unl_Conv_A_Pass : BOOL;
    In_Sen_Accum_CV_A_Full : BOOL;
    In_Sen_Unl_Conv_B_Pass : BOOL;
    Pause : ARRAY[0..99] OF Bool;
    AutoMode : BOOL;
    In_Sen_DOOR_01 : BOOL;
    In_Sen_DOOR_02 : BOOL;
    In_Sen_DOOR_03 : BOOL;
    In_Sen_DOOR_04 : BOOL;
    In_Sen_DOOR_05 : BOOL;
    In_Sen_DOOR_06 : BOOL;
    In_Sw_EMS1 : BOOL;
    In_Sw_EMS2 : BOOL;
    In_Sw_EMS3 : BOOL;
    In_Sen_AIR１_Pressure_01 : BOOL;
    In_Sen_AIR１_Pressure_02 : BOOL;
    In_Sen_AIR１_Pressure_03 : BOOL;
    TEST_M : ARRAY[0..99] OF Bool;
    ST0_Sup_Start : BOOL;  (* ST0_動作開始 *)
    Out_CYw_Sply_Pick_A_H_Auto : ARRAY[0..10] OF Bool;
    Out_CYw_Sply_Pick_A_H_Done : BOOL;
    Out_CYw_Sply_Slide_A_H_Auto : ARRAY[0..10] OF Bool;
    Out_CYw_Sply_Slide_A_H_Done : BOOL;
    Out_CYw_Sup_Chuck_A_Cl_H_Auto : ARRAY[0..10] OF Bool;
    Out_CYw_Sup_Chuck_A_Cl_H_Done : BOOL;
    In_Sen_Accum_CV_A_Arrival : BOOL;
    In_Sen_Work_A_Pos_00 : BOOL;
    Out_CYw_Sply_Pick_A_F_Auto : ARRAY[0..10] OF Bool;
    Out_CYw_Sply_Pick_A_F_Done : BOOL;
    Out_CYw_Sup_Chuck_A_Cl_F_Auto : ARRAY[0..10] OF Bool;
    Out_CYw_Sup_Chuck_A_Cl_F_Done : BOOL;
    Out_CYw_Sply_Slide_A_F_Auto : ARRAY[0..10] OF Bool;
    Out_CYw_Sply_Slide_A_F_Done : BOOL;
    Ins_A_Cv_Error : BOOL;
    Station_A_Data : ARRAY[0..8] OF sData;
    Ins_A_Cv_M : ARRAY[0..99] OF Bool;
    HMI_MessageNo : ARRAY[0..9] OF UINT;
    FH_5552_10_A_Auto : BOOL;
    In_Sen_Accum_CV_B_Full : BOOL;
    FH_Line3_Error_Status_1 : BOOL;
    FH_Line0_Error_Status_1 : BOOL;
    FH_Line1_Error_Status_1 : BOOL;
    FH_Line2_Error_Status_1 : BOOL;
    FH_Line0_Error_Clear_1 : BOOL;
    FH_Line1_Error_Clear_1 : BOOL;
    FH_Line2_Error_Clear_1 : BOOL;
    FH_Line3_Error_Clear_1 : BOOL;
    Ins_A_Next_Cycle : BOOL;
    OriginDone : BOOL;  (* 原点復帰完了 *)
    DummyDone : BOOL;  (* ダミーチェック完了 *)
    HMI_CurrentPage : STRING[256];
    Ins_A_End : BOOL;
    Auto_A_Start : BOOL;  (* 自動運転 開始 *)
    Auto_Ready : BOOL;  (* 自動運転可能 *)
    ST0_A_Sup_Busy : BOOL;
    ST1_A_Ca1_Busy : BOOL;
    RCON1_1_IN_Alarm : BOOL;
    RCON1_1_IN_EmergencyStop : BOOL;
    RCON1_1_Error : BOOL;  (* RCON1 非常停止 *)
    RCON1_1_IN_HomeDone : BOOL;
    RCON1_1_Error_Clear : BOOL;
    Error_M : ARRAY[0..99] OF Bool;  (* エラー：; [1] シリンダ; [2] コンベア＆ドアセンサ; [3] FH; [4] A(左側)検査コンベア ワーク不一致; [5] RCON1-1 異常 *)
    ST1_A_Ca1_M : ARRAY[0..99] OF Bool;
    ST2_A_Hgt_M : ARRAY[0..99] OF Bool;
    ST3_A_Dis1_M : ARRAY[0..99] OF Bool;
    HMI_Home_SW : BOOL;
    Origin_Busy : BOOL;  (* 原点復帰中 *)
    Out_CYw_Rev_01_Pick_A_H_Origin : ARRAY[0..10] OF Bool;  (* 原点復帰【Y710】A(左側)ST4 反転1ピックアップ戻： *)
    Out_CYw_Rev_01_Pick_A_H_Done : BOOL;  (* 【Y710】A(左側)ST4 反転1ピックアップ戻 動作完了 *)
    Stm_A_Rev_Axis000_Origin : BOOL;  (* A(左側) ST4 反転1 モータ原点復帰開始 *)
    Stm_A_Rev_Axis000_OriginDone : BOOL;  (* A(左側) ST4 反転1 モータ原点復帰完了 *)
    Out_CYw_Rev_01_Pick_A_F_Origin : ARRAY[0..99] OF Bool;  (* 原点復帰【Y711】A(左側)ST4 反転1ピックアップ行： *)
    Out_CYw_Rev_01_Pick_A_F_Done : BOOL;  (* 【Y711】A(左側)ST4 反転1ピックアップ行 動作完了 *)
    Out_CYw_Rev_01_Chk_A_H_Origin : ARRAY[0..99] OF Bool;  (* 原点復帰【Y708】A(左側)ST4 反転1チャック閉： *)
    Out_CYw_Rev_01_Chk_A_H_Done : BOOL;  (* 【Y708】A(左側)ST4 反転1チャック閉 動作完了 *)
    TimerQ_In_Sen_Work_A_Pos_04 : BOOL;
    Out_CYw_Rev_02_Pick_A_H_Origin : ARRAY[0..10] OF Bool;  (* 原点復帰 【Y714】A(左側)ST6 反転2ピックアップ戻 *)
    Out_CYw_Rev_02_Pick_A_H_Done : BOOL;  (* 【Y714】A(左側)ST6 反転2ピックアップ戻 動作完了 *)
    Stm_A_Rev_Axis001_Origin : BOOL;  (* A(左側) ST6 反転2 モータ原点復帰開始 *)
    Stm_A_Rev_Axis001_OriginDone : BOOL;  (* A(左側) ST6 反転2 モータ原点復帰完了 *)
    Out_CYw_Rev_02_Pick_A_F_Origin : ARRAY[0..99] OF Bool;  (* 原点復帰 【Y715】A(左側)ST6 反転2ピックアップ行 *)
    Out_CYw_Rev_02_Pick_A_F_Done : BOOL;  (* 【Y715】A(左側)ST6 反転2ピックアップ行 動作完了 *)
    Out_CYw_Rev_02_Chk_A_H_Origin : ARRAY[0..99] OF Bool;  (* 原点復帰 【Y712】A(左側)ST6 反転2チャック閉 戻 *)
    Out_CYw_Rev_02_Chk_A_H_Done : BOOL;  (* 【Y712】A(左側)ST6 反転2チャック閉 戻 動作完了 *)
    TimerQ_In_Sen_Work_A_Pos_06 : BOOL;  (* 【X208】A(左側)ワーク位置6 *)
    Auto_B_Start : BOOL;  (* B(右側)自動運転開始（後続処理未接続） *)
    Out_CYw_Rev_01_Pick_B_H_Origin : ARRAY[0..10] OF Bool;  (* 原点復帰 【Y810】B(右側)ST4 反転1ピックアップ戻 *)
    Out_CYw_Rev_01_Pick_B_H_Done : BOOL;  (* 【Y810】B(右側)ST4 反転1ピックアップ戻 動作完了 *)
    Stm_B_Rev_Axis002_Origin : BOOL;  (* B(右側) ST4 反転1 モータ原点復帰開始 *)
    Stm_B_Rev_Axis002_OriginDone : BOOL;  (* B(右側) ST4 反転1 モータ原点復帰完了 *)
    Out_CYw_Rev_01_Pick_B_F_Origin : ARRAY[0..99] OF Bool;  (* 原点復帰 【Y811】B(右側)ST4 反転1ピックアップ行 *)
    Out_CYw_Rev_01_Pick_B_F_Done : BOOL;  (* 【Y811】B(右側)ST4 反転1ピックアップ行 動作完了 *)
    Out_CYw_Rev_01_Chk_B_H_Origin : ARRAY[0..99] OF Bool;  (* 原点復帰 【Y808】B(右側)ST4 反転1チャック閉 戻 *)
    Out_CYw_Rev_01_Chk_B_H_Done : BOOL;  (* 【Y808】B(右側)ST4 反転1チャック閉 戻 動作完了 *)
    TimerQ_In_Sen_Work_B_Pos_04 : BOOL;  (* 【X406】B(右側)ワーク位置4 *)
    Out_CYw_Rev_02_Pick_B_H_Origin : ARRAY[0..10] OF Bool;  (* 原点復帰 【Y814】B(右側)ST6 反転2ピックアップ戻 *)
    Out_CYw_Rev_02_Pick_B_H_Done : BOOL;  (* 【Y814】B(右側)ST6 反転2ピックアップ戻 動作完了 *)
    Stm_B_Rev_Axis003_Origin : BOOL;  (* B(右側) ST6 反転2 モータ原点復帰開始 *)
    Stm_B_Rev_Axis003_OriginDone : BOOL;  (* B(右側) ST6 反転2 モータ原点復帰完了 *)
    Out_CYw_Rev_02_Pick_B_F_Origin : ARRAY[0..99] OF Bool;  (* 原点復帰 【Y815】B(右側)ST6 反転2ピックアップ行 *)
    Out_CYw_Rev_02_Pick_B_F_Done : BOOL;  (* 【Y815】B(右側)ST6 反転2ピックアップ行 動作完了 *)
    Out_CYw_Rev_02_Chk_B_H_Origin : ARRAY[0..99] OF Bool;  (* 原点復帰 【Y812】B(右側)ST6 反転2チャック閉 戻 *)
    Out_CYw_Rev_02_Chk_B_H_Done : BOOL;  (* 【Y812】B(右側)ST6 反転2チャック閉 戻 動作完了 *)
    TimerQ_In_Sen_Work_B_Pos_06 : BOOL;  (* 【X408】B(右側)ワーク位置6 *)
END_VAR
VAR
    _p1 : BOOL;
    _p2 : BOOL;
    _p3 : BOOL;
    _p4 : BOOL;
    _p5 : BOOL;
    _p6 : BOOL;
    _p7 : BOOL;
    _p8 : BOOL;
    _p9 : BOOL;
    _p10 : BOOL;
    _p11 : BOOL;
    _p12 : BOOL;
    _p13 : BOOL;
    _p14 : BOOL;
    _p15 : BOOL;
    _p16 : BOOL;
    _p17 : BOOL;
    _p18 : BOOL;
    _p19 : BOOL;
    _p20 : BOOL;
    _p21 : BOOL;
    _p22 : BOOL;
    _p23 : BOOL;
    _p24 : BOOL;
    _e25 : R_TRIG;
    _e26 : R_TRIG;
    _e27 : R_TRIG;
    _e28 : R_TRIG;
    _e29 : R_TRIG;
    _e30 : R_TRIG;
    _e31 : R_TRIG;
    _e32 : R_TRIG;
    _e33 : R_TRIG;
    _p34 : BOOL;
    _p35 : BOOL;
    _p36 : BOOL;
    _p37 : BOOL;
    _e38 : R_TRIG;
    _p39 : BOOL;
    _e40 : R_TRIG;
    _e41 : R_TRIG;
    _e42 : R_TRIG;
    _e43 : R_TRIG;
    _e44 : R_TRIG;
    _e45 : R_TRIG;
    _e46 : R_TRIG;
    _p47 : BOOL;
    _p48 : BOOL;
    _p49 : BOOL;
    _p50 : BOOL;
END_VAR

(* Section Initial_初期化処理: ladder, written here as Structured Text *)

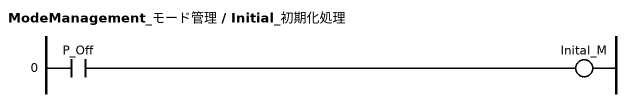
(* Rung 0 *)
Inital_M := P_Off;

(* Section Origin_原点復帰: ladder, written here as Structured Text *)

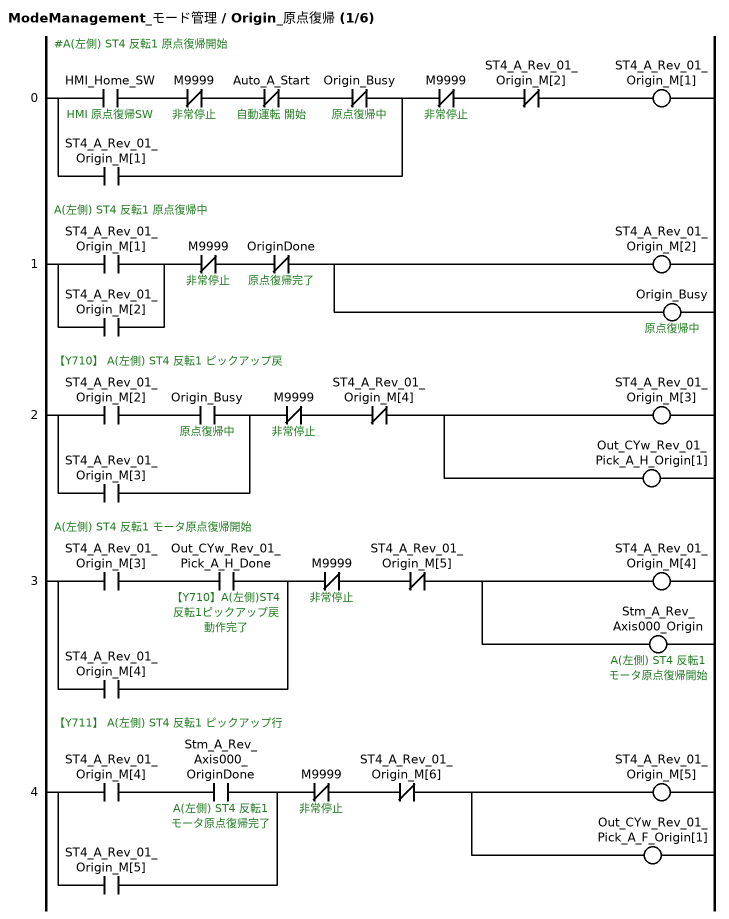
(* Rung 0: #A(左側) ST4 反転1 原点復帰開始 *)
ST4_A_Rev_01_Origin_M[1] := ((HMI_Home_SW AND NOT M9999 AND NOT Auto_A_Start AND NOT Origin_Busy) OR ST4_A_Rev_01_Origin_M[1]) AND NOT M9999 AND NOT ST4_A_Rev_01_Origin_M[2];
(* Rung 1: A(左側) ST4 反転1 原点復帰中 *)
_p1 := (ST4_A_Rev_01_Origin_M[1] OR ST4_A_Rev_01_Origin_M[2]) AND NOT M9999 AND NOT OriginDone;
ST4_A_Rev_01_Origin_M[2] := _p1;
Origin_Busy := _p1;
(* Rung 2: 【Y710】 A(左側) ST4 反転1 ピックアップ戻 *)
_p2 := ((ST4_A_Rev_01_Origin_M[2] AND Origin_Busy) OR ST4_A_Rev_01_Origin_M[3]) AND NOT M9999 AND NOT ST4_A_Rev_01_Origin_M[4];
ST4_A_Rev_01_Origin_M[3] := _p2;
Out_CYw_Rev_01_Pick_A_H_Origin[1] := _p2;
(* Rung 3: A(左側) ST4 反転1 モータ原点復帰開始 *)
_p3 := ((ST4_A_Rev_01_Origin_M[3] AND Out_CYw_Rev_01_Pick_A_H_Done) OR ST4_A_Rev_01_Origin_M[4]) AND NOT M9999 AND NOT ST4_A_Rev_01_Origin_M[5];
ST4_A_Rev_01_Origin_M[4] := _p3;
Stm_A_Rev_Axis000_Origin := _p3;
(* Rung 4: 【Y711】 A(左側) ST4 反転1 ピックアップ行 *)
_p4 := ((ST4_A_Rev_01_Origin_M[4] AND Stm_A_Rev_Axis000_OriginDone) OR ST4_A_Rev_01_Origin_M[5]) AND NOT M9999 AND NOT ST4_A_Rev_01_Origin_M[6];
ST4_A_Rev_01_Origin_M[5] := _p4;
Out_CYw_Rev_01_Pick_A_F_Origin[1] := _p4;

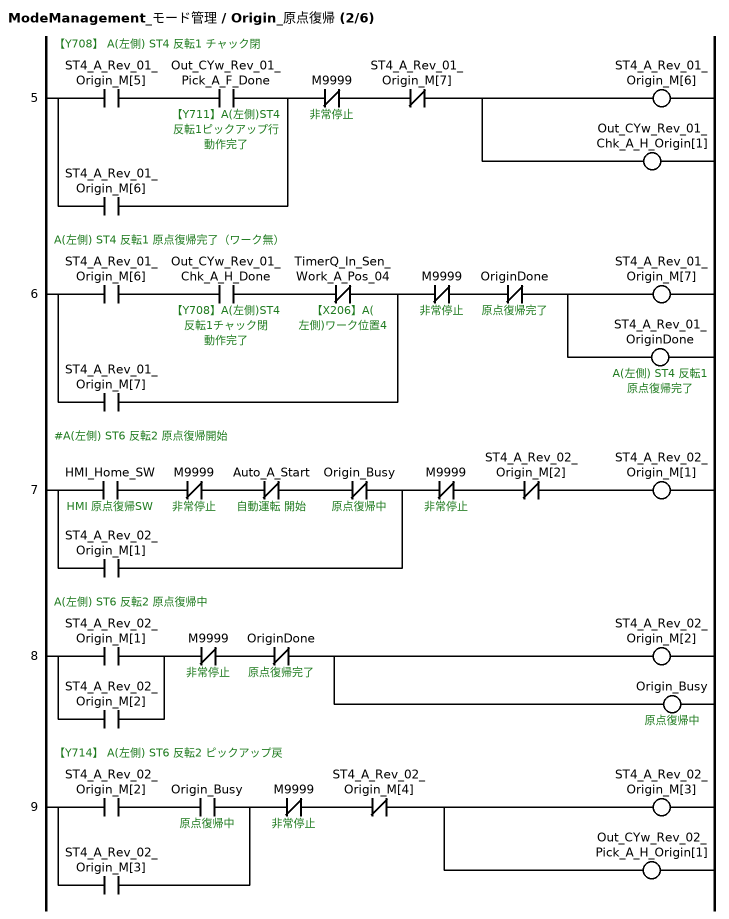
(* Rung 5: 【Y708】 A(左側) ST4 反転1 チャック閉 *)
_p5 := ((ST4_A_Rev_01_Origin_M[5] AND Out_CYw_Rev_01_Pick_A_F_Done) OR ST4_A_Rev_01_Origin_M[6]) AND NOT M9999 AND NOT ST4_A_Rev_01_Origin_M[7];
ST4_A_Rev_01_Origin_M[6] := _p5;
Out_CYw_Rev_01_Chk_A_H_Origin[1] := _p5;
(* Rung 6: A(左側) ST4 反転1 原点復帰完了（ワーク無） *)
_p6 := ((ST4_A_Rev_01_Origin_M[6] AND Out_CYw_Rev_01_Chk_A_H_Done AND NOT TimerQ_In_Sen_Work_A_Pos_04) OR ST4_A_Rev_01_Origin_M[7]) AND NOT M9999 AND NOT OriginDone;
ST4_A_Rev_01_Origin_M[7] := _p6;
ST4_A_Rev_01_OriginDone := _p6;
(* Rung 7: #A(左側) ST6 反転2 原点復帰開始 *)
ST4_A_Rev_02_Origin_M[1] := ((HMI_Home_SW AND NOT M9999 AND NOT Auto_A_Start AND NOT Origin_Busy) OR ST4_A_Rev_02_Origin_M[1]) AND NOT M9999 AND NOT ST4_A_Rev_02_Origin_M[2];
(* Rung 8: A(左側) ST6 反転2 原点復帰中 *)
_p7 := (ST4_A_Rev_02_Origin_M[1] OR ST4_A_Rev_02_Origin_M[2]) AND NOT M9999 AND NOT OriginDone;
ST4_A_Rev_02_Origin_M[2] := _p7;
Origin_Busy := _p7;
(* Rung 9: 【Y714】 A(左側) ST6 反転2 ピックアップ戻 *)
_p8 := ((ST4_A_Rev_02_Origin_M[2] AND Origin_Busy) OR ST4_A_Rev_02_Origin_M[3]) AND NOT M9999 AND NOT ST4_A_Rev_02_Origin_M[4];
ST4_A_Rev_02_Origin_M[3] := _p8;
Out_CYw_Rev_02_Pick_A_H_Origin[1] := _p8;

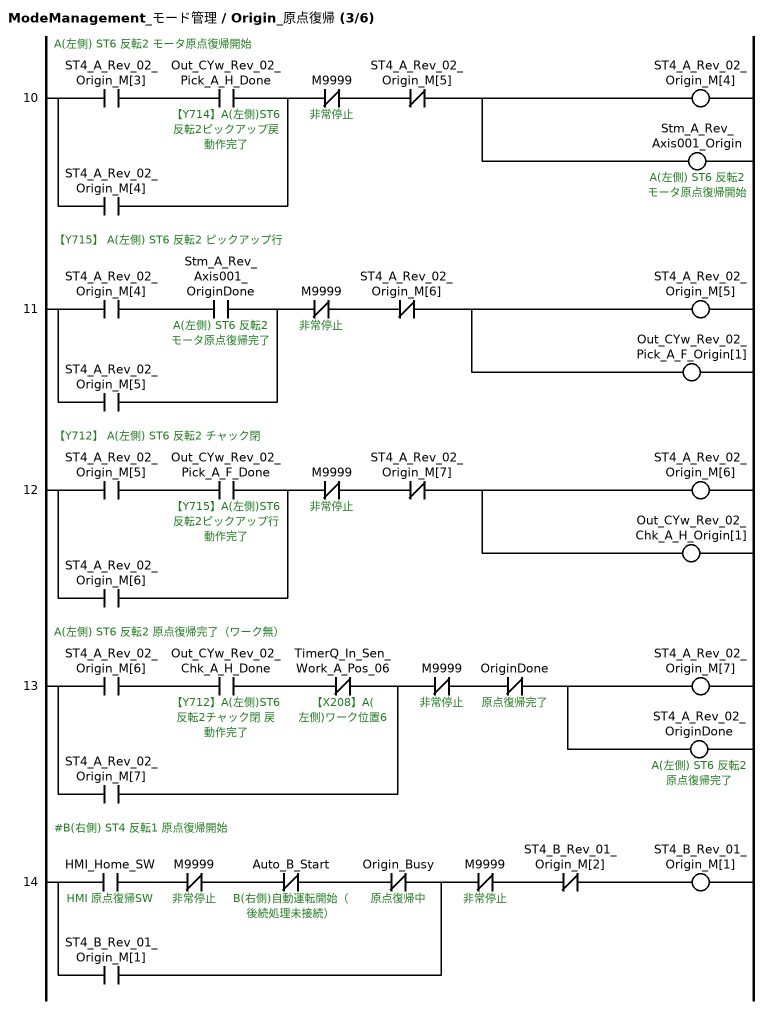
(* Rung 10: A(左側) ST6 反転2 モータ原点復帰開始 *)
_p9 := ((ST4_A_Rev_02_Origin_M[3] AND Out_CYw_Rev_02_Pick_A_H_Done) OR ST4_A_Rev_02_Origin_M[4]) AND NOT M9999 AND NOT ST4_A_Rev_02_Origin_M[5];
ST4_A_Rev_02_Origin_M[4] := _p9;
Stm_A_Rev_Axis001_Origin := _p9;
(* Rung 11: 【Y715】 A(左側) ST6 反転2 ピックアップ行 *)
_p10 := ((ST4_A_Rev_02_Origin_M[4] AND Stm_A_Rev_Axis001_OriginDone) OR ST4_A_Rev_02_Origin_M[5]) AND NOT M9999 AND NOT ST4_A_Rev_02_Origin_M[6];
ST4_A_Rev_02_Origin_M[5] := _p10;
Out_CYw_Rev_02_Pick_A_F_Origin[1] := _p10;
(* Rung 12: 【Y712】 A(左側) ST6 反転2 チャック閉 *)
_p11 := ((ST4_A_Rev_02_Origin_M[5] AND Out_CYw_Rev_02_Pick_A_F_Done) OR ST4_A_Rev_02_Origin_M[6]) AND NOT M9999 AND NOT ST4_A_Rev_02_Origin_M[7];
ST4_A_Rev_02_Origin_M[6] := _p11;
Out_CYw_Rev_02_Chk_A_H_Origin[1] := _p11;
(* Rung 13: A(左側) ST6 反転2 原点復帰完了（ワーク無） *)
_p12 := ((ST4_A_Rev_02_Origin_M[6] AND Out_CYw_Rev_02_Chk_A_H_Done AND NOT TimerQ_In_Sen_Work_A_Pos_06) OR ST4_A_Rev_02_Origin_M[7]) AND NOT M9999 AND NOT OriginDone;
ST4_A_Rev_02_Origin_M[7] := _p12;
ST4_A_Rev_02_OriginDone := _p12;
(* Rung 14: #B(右側) ST4 反転1 原点復帰開始 *)
ST4_B_Rev_01_Origin_M[1] := ((HMI_Home_SW AND NOT M9999 AND NOT Auto_B_Start AND NOT Origin_Busy) OR ST4_B_Rev_01_Origin_M[1]) AND NOT M9999 AND NOT ST4_B_Rev_01_Origin_M[2];

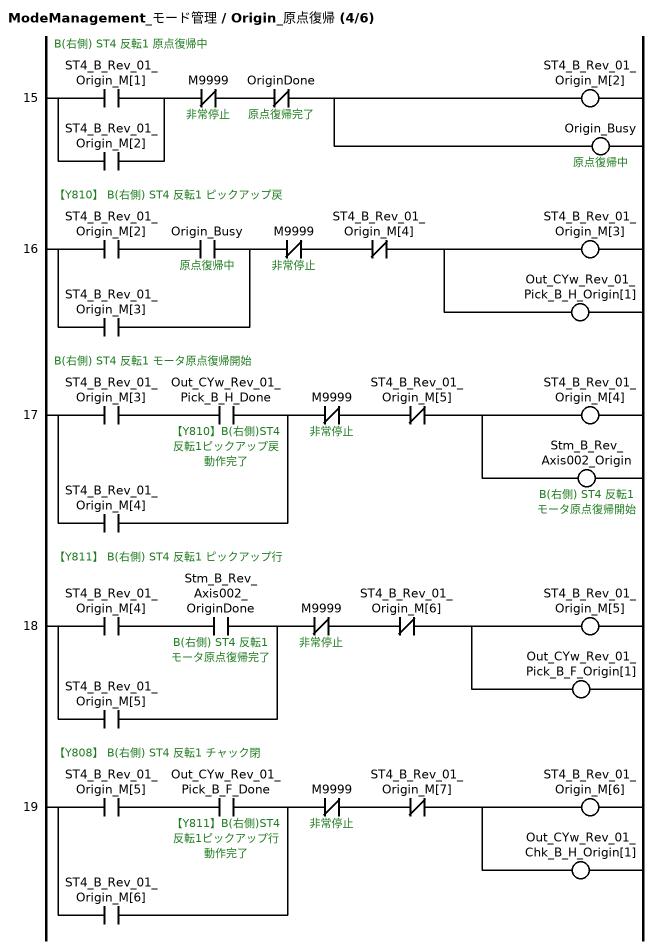
(* Rung 15: B(右側) ST4 反転1 原点復帰中 *)
_p13 := (ST4_B_Rev_01_Origin_M[1] OR ST4_B_Rev_01_Origin_M[2]) AND NOT M9999 AND NOT OriginDone;
ST4_B_Rev_01_Origin_M[2] := _p13;
Origin_Busy := _p13;
(* Rung 16: 【Y810】 B(右側) ST4 反転1 ピックアップ戻 *)
_p14 := ((ST4_B_Rev_01_Origin_M[2] AND Origin_Busy) OR ST4_B_Rev_01_Origin_M[3]) AND NOT M9999 AND NOT ST4_B_Rev_01_Origin_M[4];
ST4_B_Rev_01_Origin_M[3] := _p14;
Out_CYw_Rev_01_Pick_B_H_Origin[1] := _p14;
(* Rung 17: B(右側) ST4 反転1 モータ原点復帰開始 *)
_p15 := ((ST4_B_Rev_01_Origin_M[3] AND Out_CYw_Rev_01_Pick_B_H_Done) OR ST4_B_Rev_01_Origin_M[4]) AND NOT M9999 AND NOT ST4_B_Rev_01_Origin_M[5];
ST4_B_Rev_01_Origin_M[4] := _p15;
Stm_B_Rev_Axis002_Origin := _p15;
(* Rung 18: 【Y811】 B(右側) ST4 反転1 ピックアップ行 *)
_p16 := ((ST4_B_Rev_01_Origin_M[4] AND Stm_B_Rev_Axis002_OriginDone) OR ST4_B_Rev_01_Origin_M[5]) AND NOT M9999 AND NOT ST4_B_Rev_01_Origin_M[6];
ST4_B_Rev_01_Origin_M[5] := _p16;
Out_CYw_Rev_01_Pick_B_F_Origin[1] := _p16;
(* Rung 19: 【Y808】 B(右側) ST4 反転1 チャック閉 *)
_p17 := ((ST4_B_Rev_01_Origin_M[5] AND Out_CYw_Rev_01_Pick_B_F_Done) OR ST4_B_Rev_01_Origin_M[6]) AND NOT M9999 AND NOT ST4_B_Rev_01_Origin_M[7];
ST4_B_Rev_01_Origin_M[6] := _p17;
Out_CYw_Rev_01_Chk_B_H_Origin[1] := _p17;

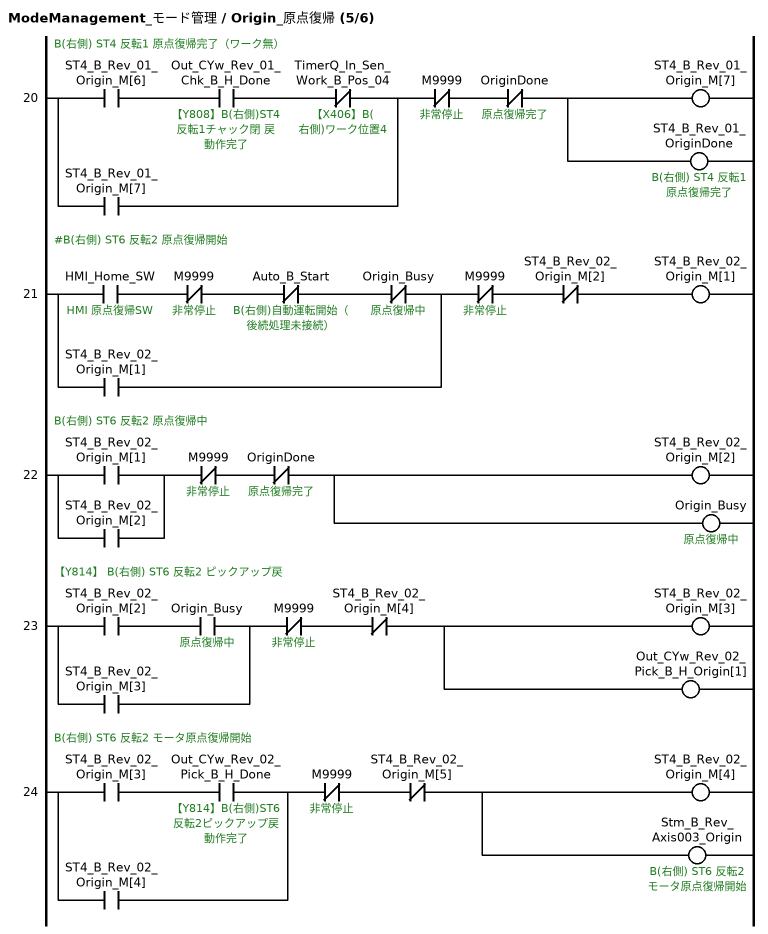
(* Rung 20: B(右側) ST4 反転1 原点復帰完了（ワーク無） *)
_p18 := ((ST4_B_Rev_01_Origin_M[6] AND Out_CYw_Rev_01_Chk_B_H_Done AND NOT TimerQ_In_Sen_Work_B_Pos_04) OR ST4_B_Rev_01_Origin_M[7]) AND NOT M9999 AND NOT OriginDone;
ST4_B_Rev_01_Origin_M[7] := _p18;
ST4_B_Rev_01_OriginDone := _p18;
(* Rung 21: #B(右側) ST6 反転2 原点復帰開始 *)
ST4_B_Rev_02_Origin_M[1] := ((HMI_Home_SW AND NOT M9999 AND NOT Auto_B_Start AND NOT Origin_Busy) OR ST4_B_Rev_02_Origin_M[1]) AND NOT M9999 AND NOT ST4_B_Rev_02_Origin_M[2];
(* Rung 22: B(右側) ST6 反転2 原点復帰中 *)
_p19 := (ST4_B_Rev_02_Origin_M[1] OR ST4_B_Rev_02_Origin_M[2]) AND NOT M9999 AND NOT OriginDone;
ST4_B_Rev_02_Origin_M[2] := _p19;
Origin_Busy := _p19;
(* Rung 23: 【Y814】 B(右側) ST6 反転2 ピックアップ戻 *)
_p20 := ((ST4_B_Rev_02_Origin_M[2] AND Origin_Busy) OR ST4_B_Rev_02_Origin_M[3]) AND NOT M9999 AND NOT ST4_B_Rev_02_Origin_M[4];
ST4_B_Rev_02_Origin_M[3] := _p20;
Out_CYw_Rev_02_Pick_B_H_Origin[1] := _p20;
(* Rung 24: B(右側) ST6 反転2 モータ原点復帰開始 *)
_p21 := ((ST4_B_Rev_02_Origin_M[3] AND Out_CYw_Rev_02_Pick_B_H_Done) OR ST4_B_Rev_02_Origin_M[4]) AND NOT M9999 AND NOT ST4_B_Rev_02_Origin_M[5];
ST4_B_Rev_02_Origin_M[4] := _p21;
Stm_B_Rev_Axis003_Origin := _p21;

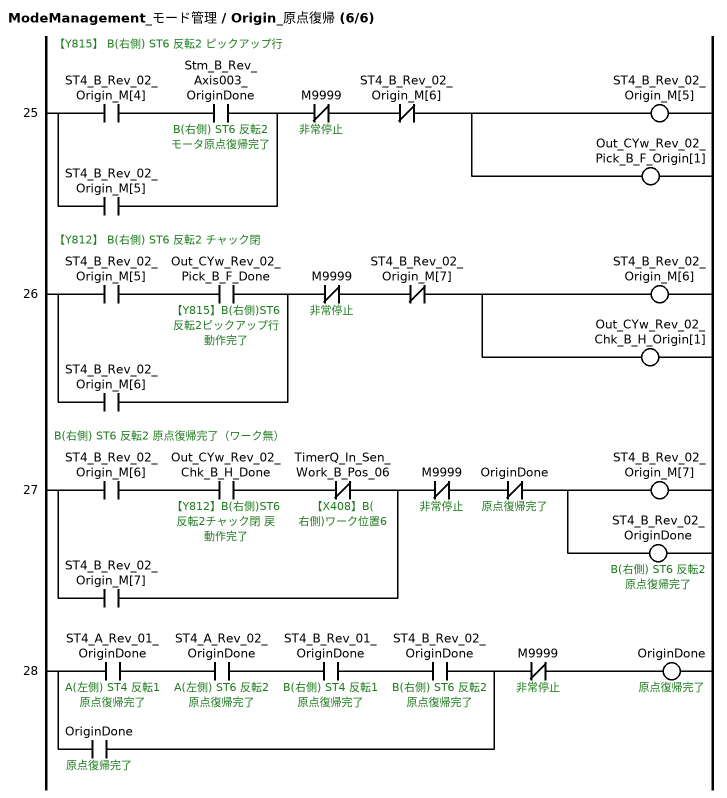
(* Rung 25: 【Y815】 B(右側) ST6 反転2 ピックアップ行 *)
_p22 := ((ST4_B_Rev_02_Origin_M[4] AND Stm_B_Rev_Axis003_OriginDone) OR ST4_B_Rev_02_Origin_M[5]) AND NOT M9999 AND NOT ST4_B_Rev_02_Origin_M[6];
ST4_B_Rev_02_Origin_M[5] := _p22;
Out_CYw_Rev_02_Pick_B_F_Origin[1] := _p22;
(* Rung 26: 【Y812】 B(右側) ST6 反転2 チャック閉 *)
_p23 := ((ST4_B_Rev_02_Origin_M[5] AND Out_CYw_Rev_02_Pick_B_F_Done) OR ST4_B_Rev_02_Origin_M[6]) AND NOT M9999 AND NOT ST4_B_Rev_02_Origin_M[7];
ST4_B_Rev_02_Origin_M[6] := _p23;
Out_CYw_Rev_02_Chk_B_H_Origin[1] := _p23;
(* Rung 27: B(右側) ST6 反転2 原点復帰完了（ワーク無） *)
_p24 := ((ST4_B_Rev_02_Origin_M[6] AND Out_CYw_Rev_02_Chk_B_H_Done AND NOT TimerQ_In_Sen_Work_B_Pos_06) OR ST4_B_Rev_02_Origin_M[7]) AND NOT M9999 AND NOT OriginDone;
ST4_B_Rev_02_Origin_M[7] := _p24;
ST4_B_Rev_02_OriginDone := _p24;
(* Rung 28 *)
OriginDone := ((ST4_A_Rev_01_OriginDone AND ST4_A_Rev_02_OriginDone AND ST4_B_Rev_01_OriginDone AND ST4_B_Rev_02_OriginDone) OR OriginDone) AND NOT M9999;

(* Section DummyCheck_ダミーチェック: ladder, written here as Structured Text *)

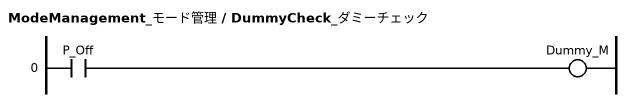
(* Rung 0 *)
Dummy_M := P_Off;

(* Section AutoMode_自動運転: ladder, written here as Structured Text *)

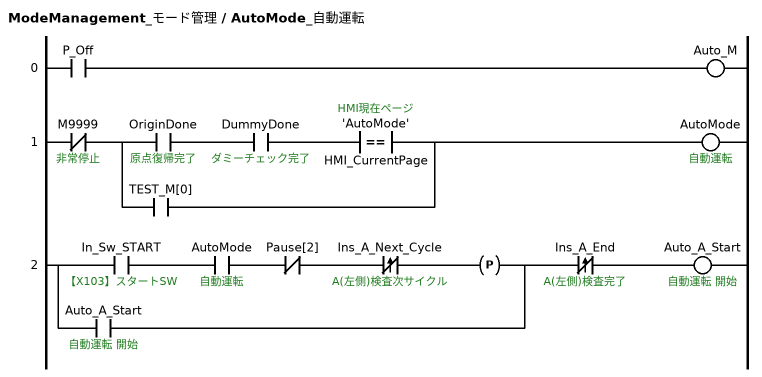
(* Rung 0 *)
Auto_M := P_Off;
(* Rung 1 *)
AutoMode := NOT M9999 AND ((OriginDone AND DummyDone AND ('AutoMode' = HMI_CurrentPage)) OR TEST_M[0]);
(* Rung 2 *)
_e25(CLK := Ins_A_Next_Cycle);
_e26(CLK := In_Sw_START AND AutoMode AND NOT Pause[2] AND NOT _e25.Q);
_e27(CLK := Ins_A_End);
Auto_A_Start := (_e26.Q OR Auto_A_Start) AND NOT _e27.Q;

(* Section Manual_手動運転: ladder, written here as Structured Text *)

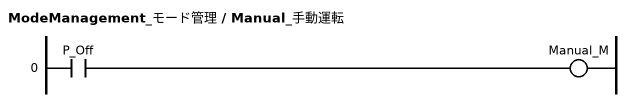
(* Rung 0 *)
Manual_M := P_Off;

(* Section Setting_設定: ladder, written here as Structured Text *)

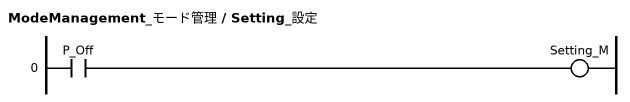
(* Rung 0 *)
Setting_M := P_Off;

(* Section Error_エラー処理: ladder, written here as Structured Text *)

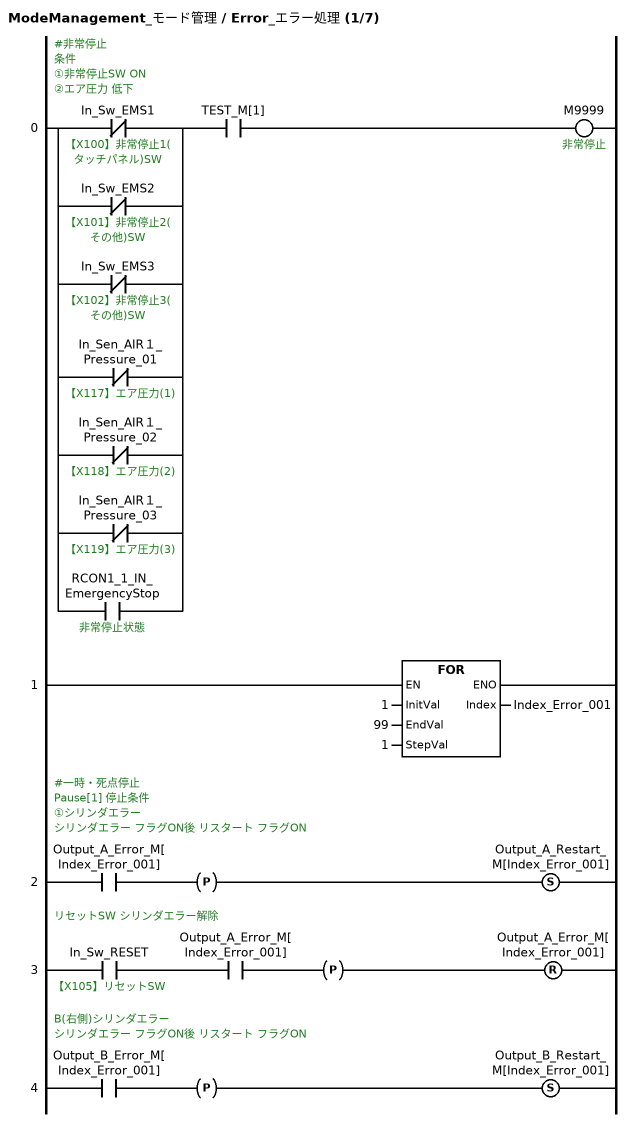
(* Rung 0: #非常停止 / 条件 / ①非常停止SW ON / ②エア圧力 低下 *)
M9999 := (NOT In_Sw_EMS1 OR NOT In_Sw_EMS2 OR NOT In_Sw_EMS3 OR NOT In_Sen_AIR１_Pressure_01 OR NOT In_Sen_AIR１_Pressure_02 OR NOT In_Sen_AIR１_Pressure_03 OR RCON1_1_IN_EmergencyStop) AND TEST_M[1];
(* Rung 1 *)
Index_Error_001 := FOR(InitVal := 1, EndVal := 99, StepVal := 1);
(* Rung 2: #一時・死点停止 / Pause[1] 停止条件 / ①シリンダエラー / シリンダエラー フラグON後 リスタート フラグON *)
_e28(CLK := Output_A_Error_M[Index_Error_001]);
IF _e28.Q THEN Output_A_Restart_M[Index_Error_001] := TRUE; END_IF;
(* Rung 3: リセットSW シリンダエラー解除 *)
_e29(CLK := In_Sw_RESET AND Output_A_Error_M[Index_Error_001]);
IF _e29.Q THEN Output_A_Error_M[Index_Error_001] := FALSE; END_IF;
(* Rung 4: B(右側)シリンダエラー / シリンダエラー フラグON後 リスタート フラグON *)
_e30(CLK := Output_B_Error_M[Index_Error_001]);
IF _e30.Q THEN Output_B_Restart_M[Index_Error_001] := TRUE; END_IF;

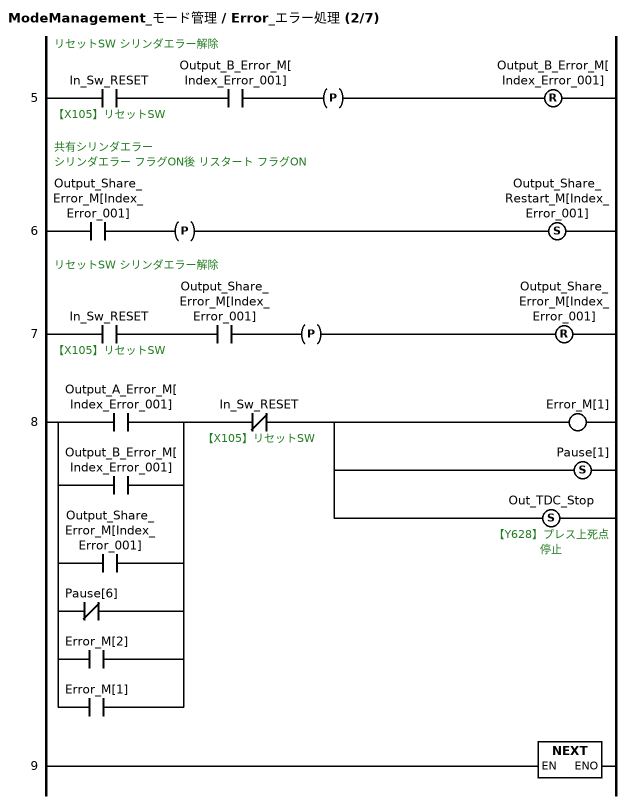
(* Rung 5: リセットSW シリンダエラー解除 *)
_e31(CLK := In_Sw_RESET AND Output_B_Error_M[Index_Error_001]);
IF _e31.Q THEN Output_B_Error_M[Index_Error_001] := FALSE; END_IF;
(* Rung 6: 共有シリンダエラー / シリンダエラー フラグON後 リスタート フラグON *)
_e32(CLK := Output_Share_Error_M[Index_Error_001]);
IF _e32.Q THEN Output_Share_Restart_M[Index_Error_001] := TRUE; END_IF;
(* Rung 7: リセットSW シリンダエラー解除 *)
_e33(CLK := In_Sw_RESET AND Output_Share_Error_M[Index_Error_001]);
IF _e33.Q THEN Output_Share_Error_M[Index_Error_001] := FALSE; END_IF;
(* Rung 8 *)
_p34 := (Output_A_Error_M[Index_Error_001] OR Output_B_Error_M[Index_Error_001] OR Output_Share_Error_M[Index_Error_001] OR NOT Pause[6] OR Error_M[2] OR Error_M[1]) AND NOT In_Sw_RESET;
Error_M[1] := _p34;
IF _p34 THEN
    Pause[1] := TRUE;
    Out_TDC_Stop := TRUE;
END_IF;
(* Rung 9 *)
NEXT();

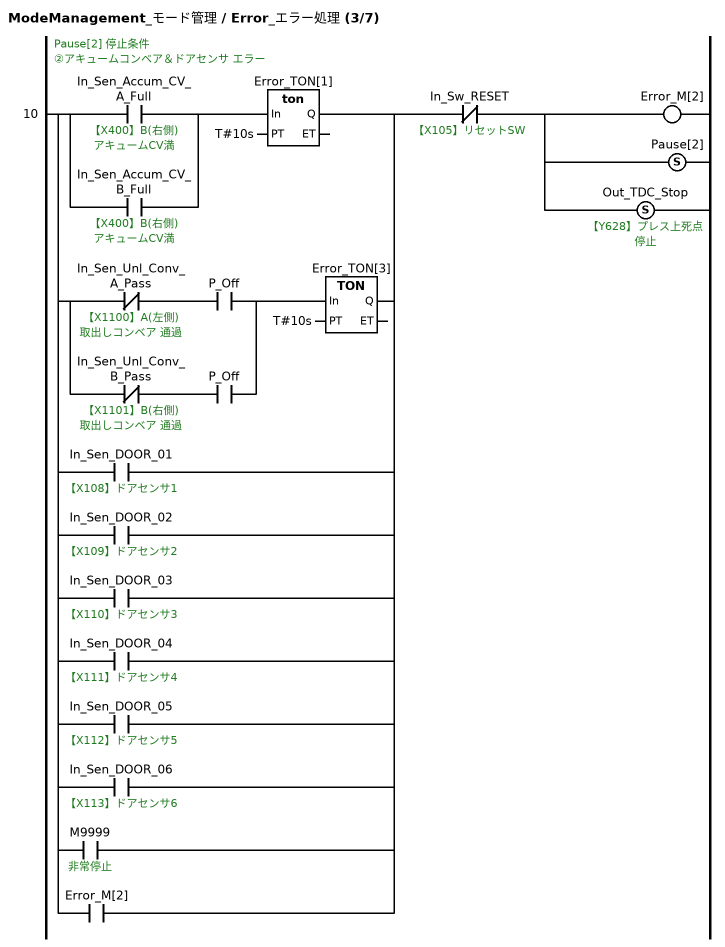
(* Rung 10: Pause[2] 停止条件 / ②アキュームコンベア＆ドアセンサ エラー *)
Error_TON[1](In := In_Sen_Accum_CV_A_Full OR In_Sen_Accum_CV_B_Full, PT := T#10s);
_p35 := Error_TON[1].Q;
Error_TON[3](In := (NOT In_Sen_Unl_Conv_A_Pass AND P_Off) OR (NOT In_Sen_Unl_Conv_B_Pass AND P_Off), PT := T#10s);
_p36 := (_p35 OR Error_TON[3].Q OR In_Sen_DOOR_01 OR In_Sen_DOOR_02 OR In_Sen_DOOR_03 OR In_Sen_DOOR_04 OR In_Sen_DOOR_05 OR In_Sen_DOOR_06 OR M9999 OR Error_M[2]) AND NOT In_Sw_RESET;
Error_M[2] := _p36;
IF _p36 THEN
    Pause[2] := TRUE;
    Out_TDC_Stop := TRUE;
END_IF;

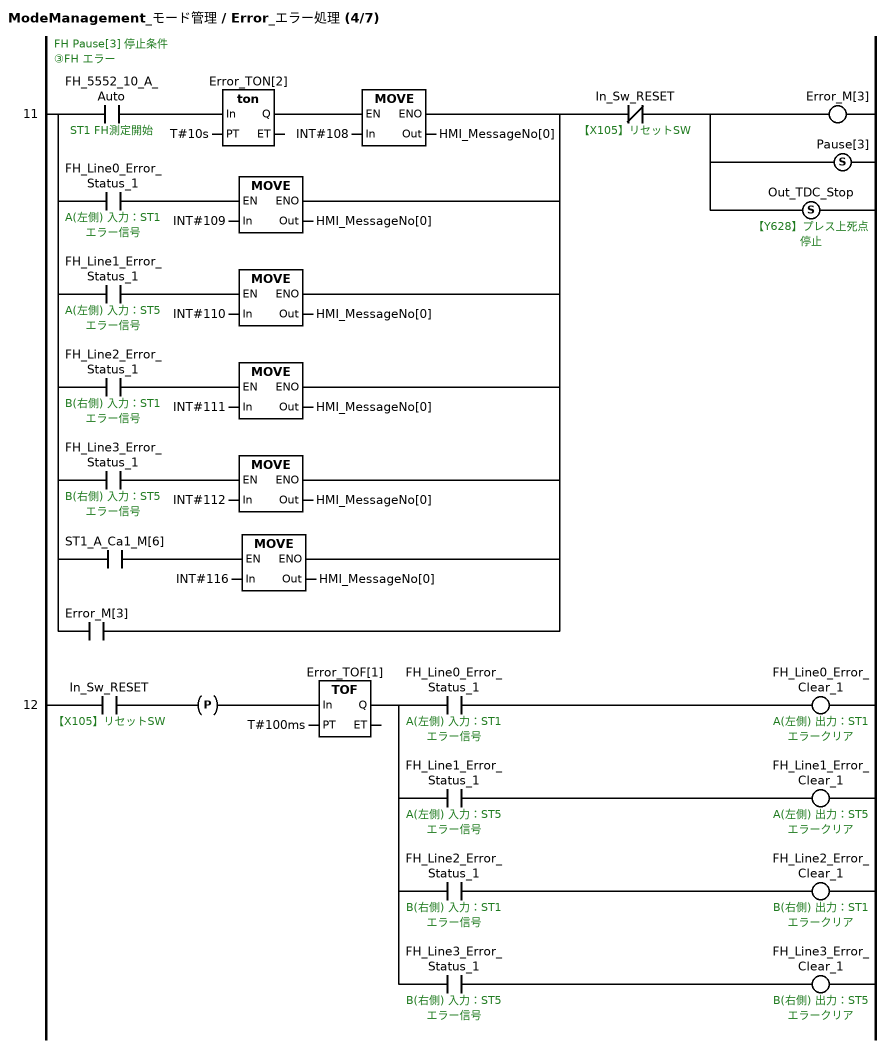
(* Rung 11: FH Pause[3] 停止条件 / ③FH エラー *)
Error_TON[2](In := FH_5552_10_A_Auto, PT := T#10s);
IF Error_TON[2].Q THEN HMI_MessageNo[0] := INT#108; END_IF;
IF FH_Line0_Error_Status_1 THEN HMI_MessageNo[0] := INT#109; END_IF;
IF FH_Line1_Error_Status_1 THEN HMI_MessageNo[0] := INT#110; END_IF;
IF FH_Line2_Error_Status_1 THEN HMI_MessageNo[0] := INT#111; END_IF;
IF FH_Line3_Error_Status_1 THEN HMI_MessageNo[0] := INT#112; END_IF;
IF ST1_A_Ca1_M[6] THEN HMI_MessageNo[0] := INT#116; END_IF;
_p37 := (Error_TON[2].Q OR FH_Line0_Error_Status_1 OR FH_Line1_Error_Status_1 OR FH_Line2_Error_Status_1 OR FH_Line3_Error_Status_1 OR ST1_A_Ca1_M[6] OR Error_M[3]) AND NOT In_Sw_RESET;
Error_M[3] := _p37;
IF _p37 THEN
    Pause[3] := TRUE;
    Out_TDC_Stop := TRUE;
END_IF;
(* Rung 12 *)
_e38(CLK := In_Sw_RESET);
Error_TOF[1](In := _e38.Q, PT := T#100ms);
FH_Line0_Error_Clear_1 := Error_TOF[1].Q AND FH_Line0_Error_Status_1;
FH_Line1_Error_Clear_1 := Error_TOF[1].Q AND FH_Line1_Error_Status_1;
FH_Line2_Error_Clear_1 := Error_TOF[1].Q AND FH_Line2_Error_Status_1;
FH_Line3_Error_Clear_1 := Error_TOF[1].Q AND FH_Line3_Error_Status_1;

